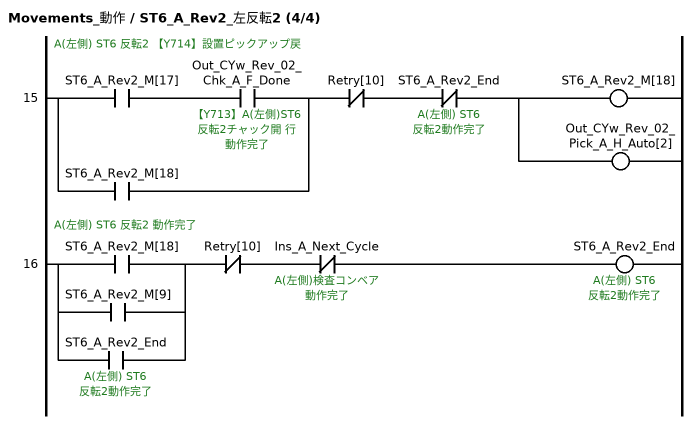
(* [picture p48: Movements_動作 / ST6_A_Rev2_左反転2, rungs 15-16] *)
(* Rung 15: A(左側) ST6 反転2 【Y714】設置ピックアップ戻 *)
_p89 := ((ST6_A_Rev2_M[17] AND Out_CYw_Rev_02_Chk_A_F_Done) OR ST6_A_Rev2_M[18]) AND NOT Retry[10] AND NOT ST6_A_Rev2_End;
ST6_A_Rev2_M[18] := _p89;
Out_CYw_Rev_02_Pick_A_H_Auto[2] := _p89;
(* Rung 16: A(左側) ST6 反転2 動作完了 *)
ST6_A_Rev2_End := (ST6_A_Rev2_M[18] OR ST6_A_Rev2_M[9] OR ST6_A_Rev2_End) AND NOT Retry[10] AND NOT Ins_A_Next_Cycle;

(* Section ST7_A_Dis2_左SF排出: ladder, written here as Structured Text *)

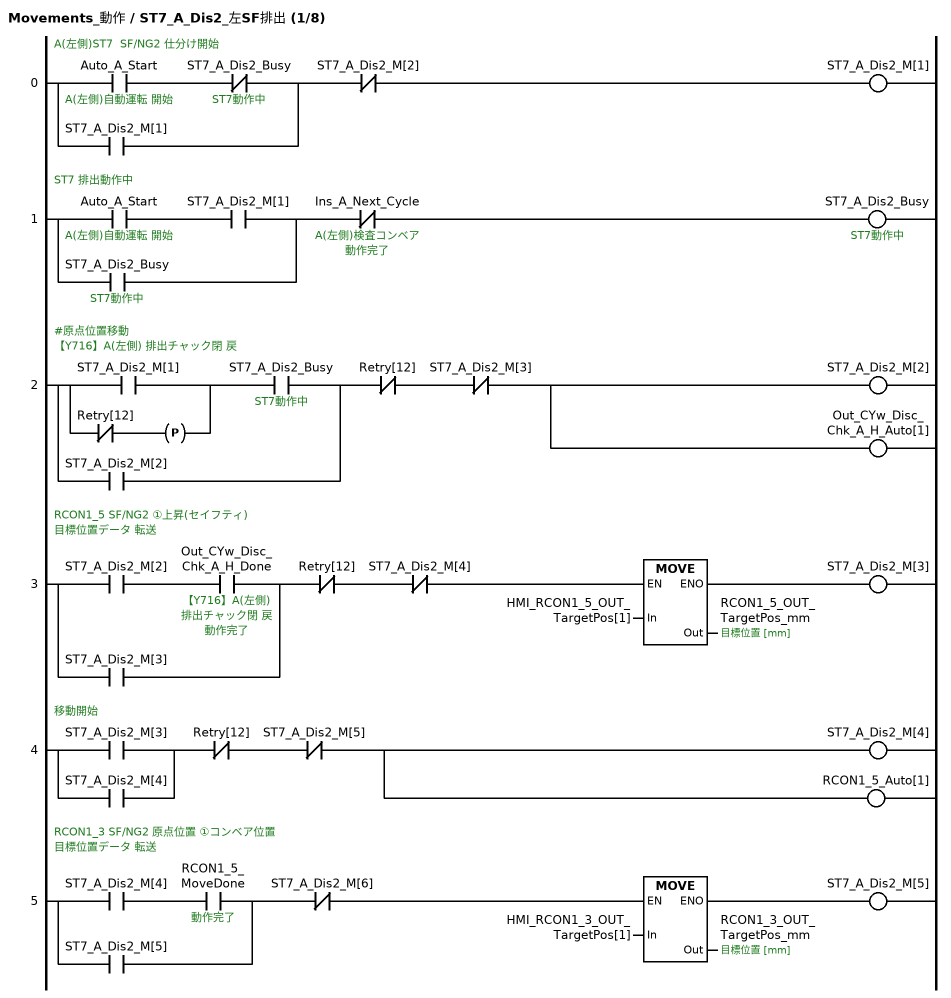
(* Rung 0: A(左側)ST7  SF/NG2 仕分け開始 *)
ST7_A_Dis2_M[1] := ((Auto_A_Start AND NOT ST7_A_Dis2_Busy) OR ST7_A_Dis2_M[1]) AND NOT ST7_A_Dis2_M[2];
(* Rung 1: ST7 排出動作中 *)
ST7_A_Dis2_Busy := ((Auto_A_Start AND ST7_A_Dis2_M[1]) OR ST7_A_Dis2_Busy) AND NOT Ins_A_Next_Cycle;
(* Rung 2: #原点位置移動 / 【Y716】A(左側) 排出チャック閉 戻 *)
_e90(CLK := NOT Retry[12]);
_p91 := (((ST7_A_Dis2_M[1] OR _e90.Q) AND ST7_A_Dis2_Busy) OR ST7_A_Dis2_M[2]) AND NOT Retry[12] AND NOT ST7_A_Dis2_M[3];
ST7_A_Dis2_M[2] := _p91;
Out_CYw_Disc_Chk_A_H_Auto[1] := _p91;
(* Rung 3: RCON1_5 SF/NG2 ①上昇(セイフティ) / 目標位置データ 転送 *)
IF ((ST7_A_Dis2_M[2] AND Out_CYw_Disc_Chk_A_H_Done) OR ST7_A_Dis2_M[3]) AND NOT Retry[12] AND NOT ST7_A_Dis2_M[4] THEN
    RCON1_5_OUT_TargetPos_mm := HMI_RCON1_5_OUT_TargetPos[1];
END_IF;
ST7_A_Dis2_M[3] := ((ST7_A_Dis2_M[2] AND Out_CYw_Disc_Chk_A_H_Done) OR ST7_A_Dis2_M[3]) AND NOT Retry[12] AND NOT ST7_A_Dis2_M[4];
(* Rung 4: 移動開始 *)
_p92 := (ST7_A_Dis2_M[3] OR ST7_A_Dis2_M[4]) AND NOT Retry[12] AND NOT ST7_A_Dis2_M[5];
ST7_A_Dis2_M[4] := _p92;
RCON1_5_Auto[1] := _p92;
(* Rung 5: RCON1_3 SF/NG2 原点位置 ①コンベア位置 / 目標位置データ 転送 *)
IF ((ST7_A_Dis2_M[4] AND RCON1_5_MoveDone) OR ST7_A_Dis2_M[5]) AND NOT ST7_A_Dis2_M[6] THEN
    RCON1_3_OUT_TargetPos_mm := HMI_RCON1_3_OUT_TargetPos[1];
END_IF;
ST7_A_Dis2_M[5] := ((ST7_A_Dis2_M[4] AND RCON1_5_MoveDone) OR ST7_A_Dis2_M[5]) AND NOT ST7_A_Dis2_M[6];

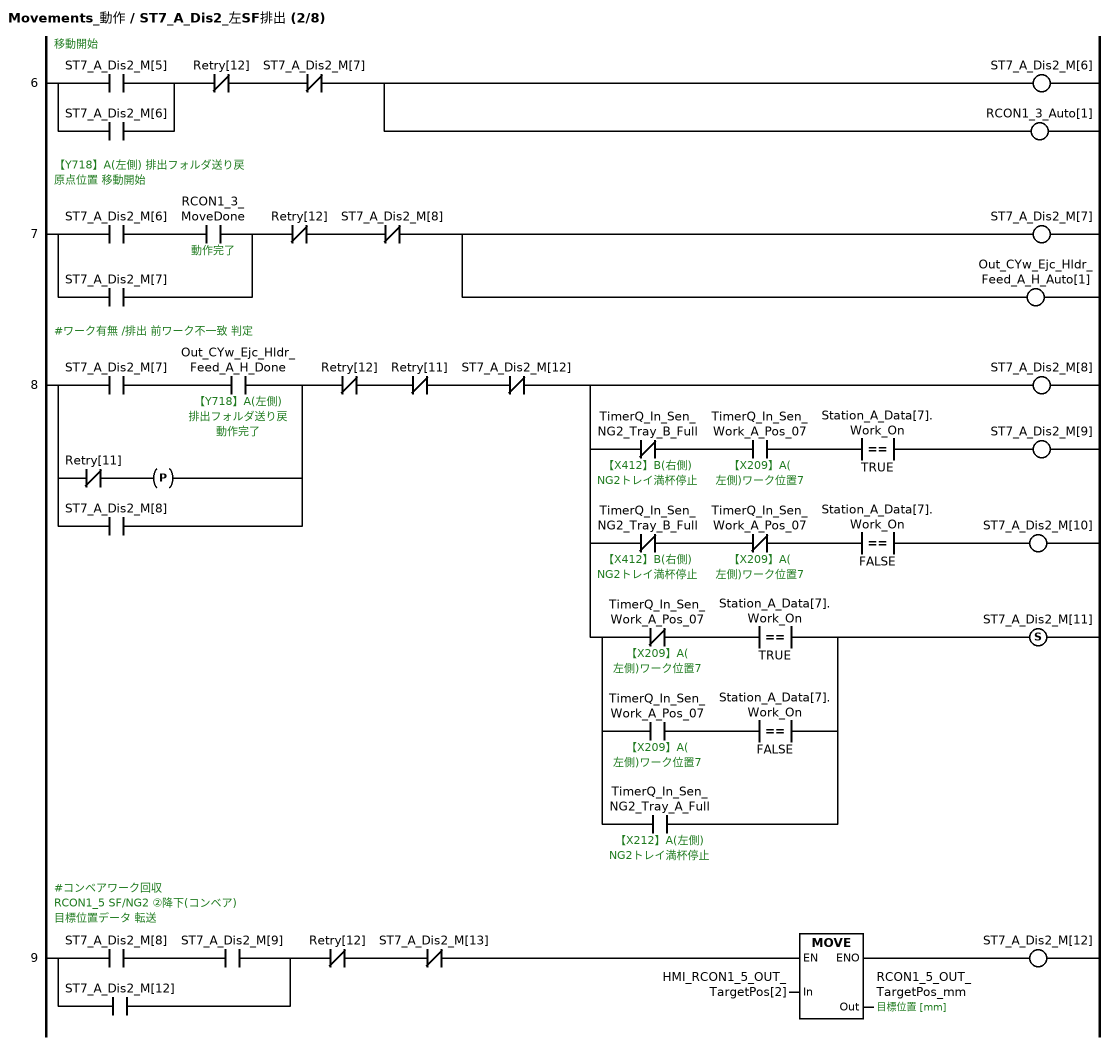
(* Rung 6: 移動開始 *)
_p93 := (ST7_A_Dis2_M[5] OR ST7_A_Dis2_M[6]) AND NOT Retry[12] AND NOT ST7_A_Dis2_M[7];
ST7_A_Dis2_M[6] := _p93;
RCON1_3_Auto[1] := _p93;
(* Rung 7: 【Y718】A(左側) 排出フォルダ送り戻 / 原点位置 移動開始 *)
_p94 := ((ST7_A_Dis2_M[6] AND RCON1_3_MoveDone) OR ST7_A_Dis2_M[7]) AND NOT Retry[12] AND NOT ST7_A_Dis2_M[8];
ST7_A_Dis2_M[7] := _p94;
Out_CYw_Ejc_Hldr_Feed_A_H_Auto[1] := _p94;
(* Rung 8: #ワーク有無 /排出 前ワーク不一致 判定 *)
_e95(CLK := NOT Retry[11]);
_p96 := ((ST7_A_Dis2_M[7] AND Out_CYw_Ejc_Hldr_Feed_A_H_Done) OR _e95.Q OR ST7_A_Dis2_M[8]) AND NOT Retry[12] AND NOT Retry[11] AND NOT ST7_A_Dis2_M[12];
ST7_A_Dis2_M[8] := _p96;
ST7_A_Dis2_M[9] := _p96 AND NOT TimerQ_In_Sen_NG2_Tray_B_Full AND TimerQ_In_Sen_Work_A_Pos_07 AND (Station_A_Data[7].Work_On = TRUE);
ST7_A_Dis2_M[10] := _p96 AND NOT TimerQ_In_Sen_NG2_Tray_B_Full AND NOT TimerQ_In_Sen_Work_A_Pos_07 AND (Station_A_Data[7].Work_On = FALSE);
IF _p96 AND ((NOT TimerQ_In_Sen_Work_A_Pos_07 AND (Station_A_Data[7].Work_On = TRUE)) OR (TimerQ_In_Sen_Work_A_Pos_07 AND (Station_A_Data[7].Work_On = FALSE)) OR TimerQ_In_Sen_NG2_Tray_A_Full) THEN
    ST7_A_Dis2_M[11] := TRUE;
END_IF;
(* Rung 9: #コンベアワーク回収 / RCON1_5 SF/NG2 ②降下(コンベア) / 目標位置データ 転送 *)
IF ((ST7_A_Dis2_M[8] AND ST7_A_Dis2_M[9]) OR ST7_A_Dis2_M[12]) AND NOT Retry[12] AND NOT ST7_A_Dis2_M[13] THEN
    RCON1_5_OUT_TargetPos_mm := HMI_RCON1_5_OUT_TargetPos[2];
END_IF;
ST7_A_Dis2_M[12] := ((ST7_A_Dis2_M[8] AND ST7_A_Dis2_M[9]) OR ST7_A_Dis2_M[12]) AND NOT Retry[12] AND NOT ST7_A_Dis2_M[13];

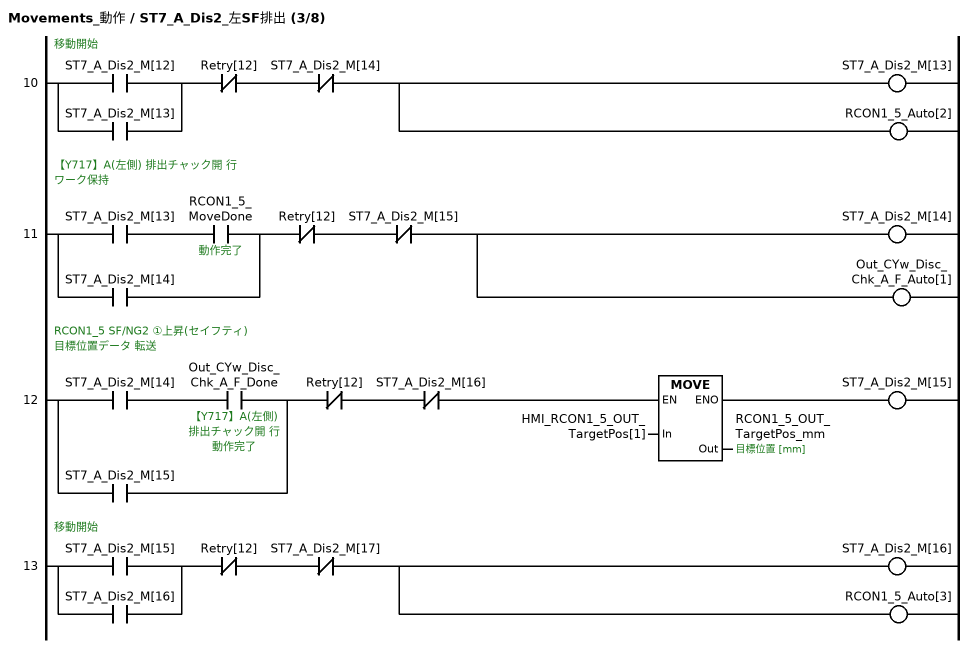
(* Rung 10: 移動開始 *)
_p97 := (ST7_A_Dis2_M[12] OR ST7_A_Dis2_M[13]) AND NOT Retry[12] AND NOT ST7_A_Dis2_M[14];
ST7_A_Dis2_M[13] := _p97;
RCON1_5_Auto[2] := _p97;
(* Rung 11: 【Y717】A(左側) 排出チャック開 行 / ワーク保持 *)
_p98 := ((ST7_A_Dis2_M[13] AND RCON1_5_MoveDone) OR ST7_A_Dis2_M[14]) AND NOT Retry[12] AND NOT ST7_A_Dis2_M[15];
ST7_A_Dis2_M[14] := _p98;
Out_CYw_Disc_Chk_A_F_Auto[1] := _p98;
(* Rung 12: RCON1_5 SF/NG2 ①上昇(セイフティ) / 目標位置データ 転送 *)
IF ((ST7_A_Dis2_M[14] AND Out_CYw_Disc_Chk_A_F_Done) OR ST7_A_Dis2_M[15]) AND NOT Retry[12] AND NOT ST7_A_Dis2_M[16] THEN
    RCON1_5_OUT_TargetPos_mm := HMI_RCON1_5_OUT_TargetPos[1];
END_IF;
ST7_A_Dis2_M[15] := ((ST7_A_Dis2_M[14] AND Out_CYw_Disc_Chk_A_F_Done) OR ST7_A_Dis2_M[15]) AND NOT Retry[12] AND NOT ST7_A_Dis2_M[16];
(* Rung 13: 移動開始 *)
_p99 := (ST7_A_Dis2_M[15] OR ST7_A_Dis2_M[16]) AND NOT Retry[12] AND NOT ST7_A_Dis2_M[17];
ST7_A_Dis2_M[16] := _p99;
RCON1_5_Auto[3] := _p99;

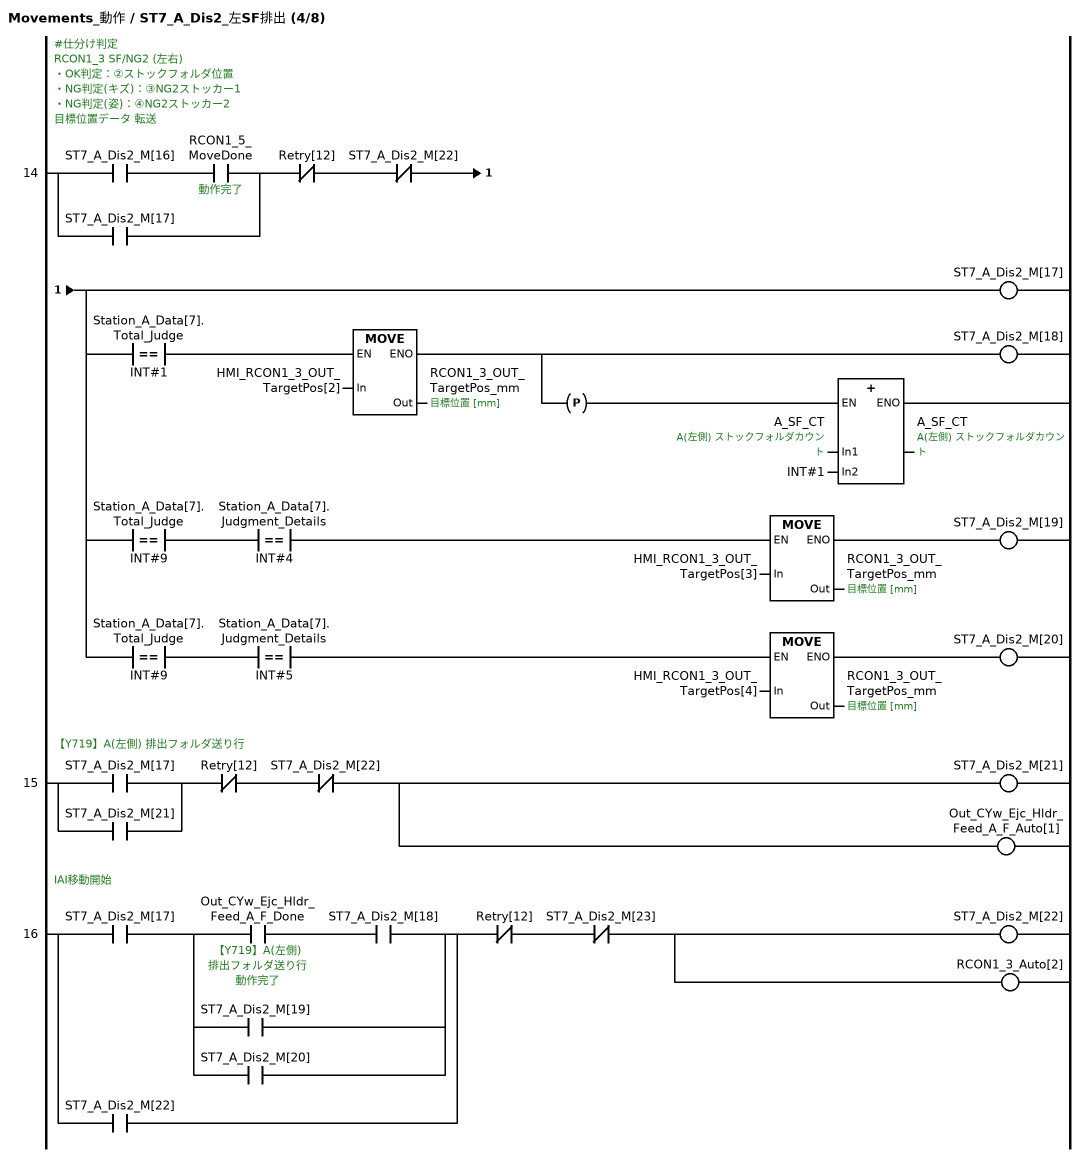
(* Rung 14: #仕分け判定 / RCON1_3 SF/NG2 (左右) / ・OK判定：②ストックフォルダ位置 / ・NG判定(キズ)：③NG2ストッカー1 / ・NG判定(姿)：④NG2ストッカー2 / 目標位置データ 転送 *)
_p100 := ((ST7_A_Dis2_M[16] AND RCON1_5_MoveDone) OR ST7_A_Dis2_M[17]) AND NOT Retry[12] AND NOT ST7_A_Dis2_M[22];
ST7_A_Dis2_M[17] := _p100;
IF _p100 AND (Station_A_Data[7].Total_Judge = INT#1) THEN
    RCON1_3_OUT_TargetPos_mm := HMI_RCON1_3_OUT_TargetPos[2];
END_IF;
_p101 := _p100 AND (Station_A_Data[7].Total_Judge = INT#1);
ST7_A_Dis2_M[18] := _p101;
_e102(CLK := _p101);
IF _e102.Q THEN A_SF_CT := A_SF_CT + INT#1; END_IF;
IF _p100 AND (Station_A_Data[7].Total_Judge = INT#9) AND (Station_A_Data[7].Judgment_Details = INT#4) THEN
    RCON1_3_OUT_TargetPos_mm := HMI_RCON1_3_OUT_TargetPos[3];
END_IF;
ST7_A_Dis2_M[19] := _p100 AND (Station_A_Data[7].Total_Judge = INT#9) AND (Station_A_Data[7].Judgment_Details = INT#4);
IF _p100 AND (Station_A_Data[7].Total_Judge = INT#9) AND (Station_A_Data[7].Judgment_Details = INT#5) THEN
    RCON1_3_OUT_TargetPos_mm := HMI_RCON1_3_OUT_TargetPos[4];
END_IF;
ST7_A_Dis2_M[20] := _p100 AND (Station_A_Data[7].Total_Judge = INT#9) AND (Station_A_Data[7].Judgment_Details = INT#5);
(* Rung 15: 【Y719】A(左側) 排出フォルダ送り行 *)
_p103 := (ST7_A_Dis2_M[17] OR ST7_A_Dis2_M[21]) AND NOT Retry[12] AND NOT ST7_A_Dis2_M[22];
ST7_A_Dis2_M[21] := _p103;
Out_CYw_Ejc_Hldr_Feed_A_F_Auto[1] := _p103;
(* Rung 16: IAI移動開始 *)
_p104 := ((ST7_A_Dis2_M[17] AND ((Out_CYw_Ejc_Hldr_Feed_A_F_Done AND ST7_A_Dis2_M[18]) OR ST7_A_Dis2_M[19] OR ST7_A_Dis2_M[20])) OR ST7_A_Dis2_M[22]) AND NOT Retry[12] AND NOT ST7_A_Dis2_M[23];
ST7_A_Dis2_M[22] := _p104;
RCON1_3_Auto[2] := _p104;

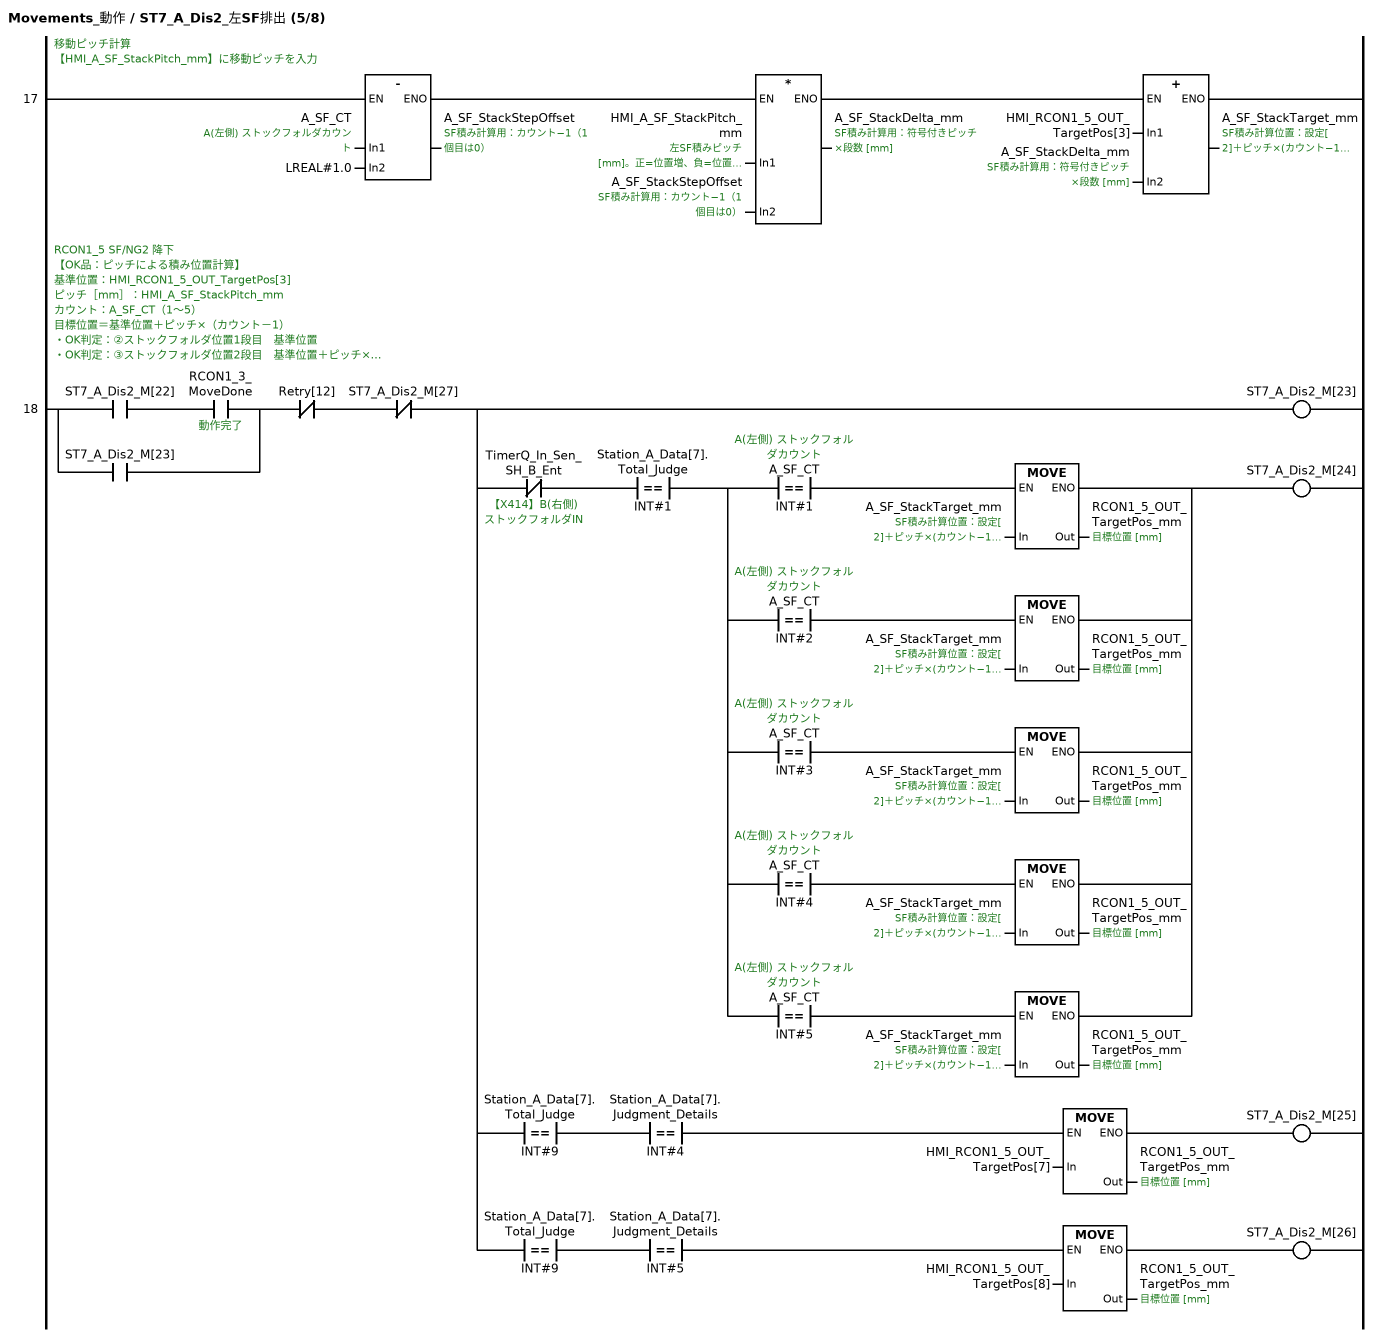
(* Rung 17: 移動ピッチ計算 / 【HMI_A_SF_StackPitch_mm】に移動ピッチを入力 *)
A_SF_StackStepOffset := A_SF_CT - LREAL#1.0;
A_SF_StackDelta_mm := HMI_A_SF_StackPitch_mm * A_SF_StackStepOffset;
A_SF_StackTarget_mm := HMI_RCON1_5_OUT_TargetPos[3] + A_SF_StackDelta_mm;
(* Rung 18: RCON1_5 SF/NG2 降下 / 【OK品：ピッチによる積み位置計算】 / 基準位置：HMI_RCON1_5_OUT_TargetPos[3] / ピッチ［mm］：HMI_A_SF_StackPitch_mm / カウント：A_SF_CT（1～5） / 目標位置＝基準位置＋ピッチ×（カウント－1） / ・OK判定：②ストックフォルダ位置1段目　基準位置 / ・OK判定：③ストックフォルダ位置2段目　基準位置＋ピッチ×1 / ・OK判定：④ストックフォルダ位置3段目　基準位置＋ピッチ×2 / ・OK判定：⑤ストックフォルダ位置4段目　基準位置＋ピッチ×3 / ・OK判定：⑥ストックフォルダ位置5段目　基準位置＋ピッチ×4 / 【NG品：従来の固定位置を使用】 / ・NG判定(キズ)：⑦NG2ストッカー1 / ・NG判定(姿)：⑧NG2ストッカー2 / 目標位置データ 転送 *)
_p105 := ((ST7_A_Dis2_M[22] AND RCON1_3_MoveDone) OR ST7_A_Dis2_M[23]) AND NOT Retry[12] AND NOT ST7_A_Dis2_M[27];
ST7_A_Dis2_M[23] := _p105;
_p106 := _p105 AND NOT TimerQ_In_Sen_SH_B_Ent AND (Station_A_Data[7].Total_Judge = INT#1);
IF _p106 AND (A_SF_CT = INT#1) THEN RCON1_5_OUT_TargetPos_mm := A_SF_StackTarget_mm; END_IF;
IF _p106 AND (A_SF_CT = INT#2) THEN RCON1_5_OUT_TargetPos_mm := A_SF_StackTarget_mm; END_IF;
IF _p106 AND (A_SF_CT = INT#3) THEN RCON1_5_OUT_TargetPos_mm := A_SF_StackTarget_mm; END_IF;
IF _p106 AND (A_SF_CT = INT#4) THEN RCON1_5_OUT_TargetPos_mm := A_SF_StackTarget_mm; END_IF;
IF _p106 AND (A_SF_CT = INT#5) THEN RCON1_5_OUT_TargetPos_mm := A_SF_StackTarget_mm; END_IF;
ST7_A_Dis2_M[24] := _p106 AND ((A_SF_CT = INT#1) OR (A_SF_CT = INT#2) OR (A_SF_CT = INT#3) OR (A_SF_CT = INT#4) OR (A_SF_CT = INT#5));
IF _p105 AND (Station_A_Data[7].Total_Judge = INT#9) AND (Station_A_Data[7].Judgment_Details = INT#4) THEN
    RCON1_5_OUT_TargetPos_mm := HMI_RCON1_5_OUT_TargetPos[7];
END_IF;
ST7_A_Dis2_M[25] := _p105 AND (Station_A_Data[7].Total_Judge = INT#9) AND (Station_A_Data[7].Judgment_Details = INT#4);
IF _p105 AND (Station_A_Data[7].Total_Judge = INT#9) AND (Station_A_Data[7].Judgment_Details = INT#5) THEN
    RCON1_5_OUT_TargetPos_mm := HMI_RCON1_5_OUT_TargetPos[8];
END_IF;
ST7_A_Dis2_M[26] := _p105 AND (Station_A_Data[7].Total_Judge = INT#9) AND (Station_A_Data[7].Judgment_Details = INT#5);

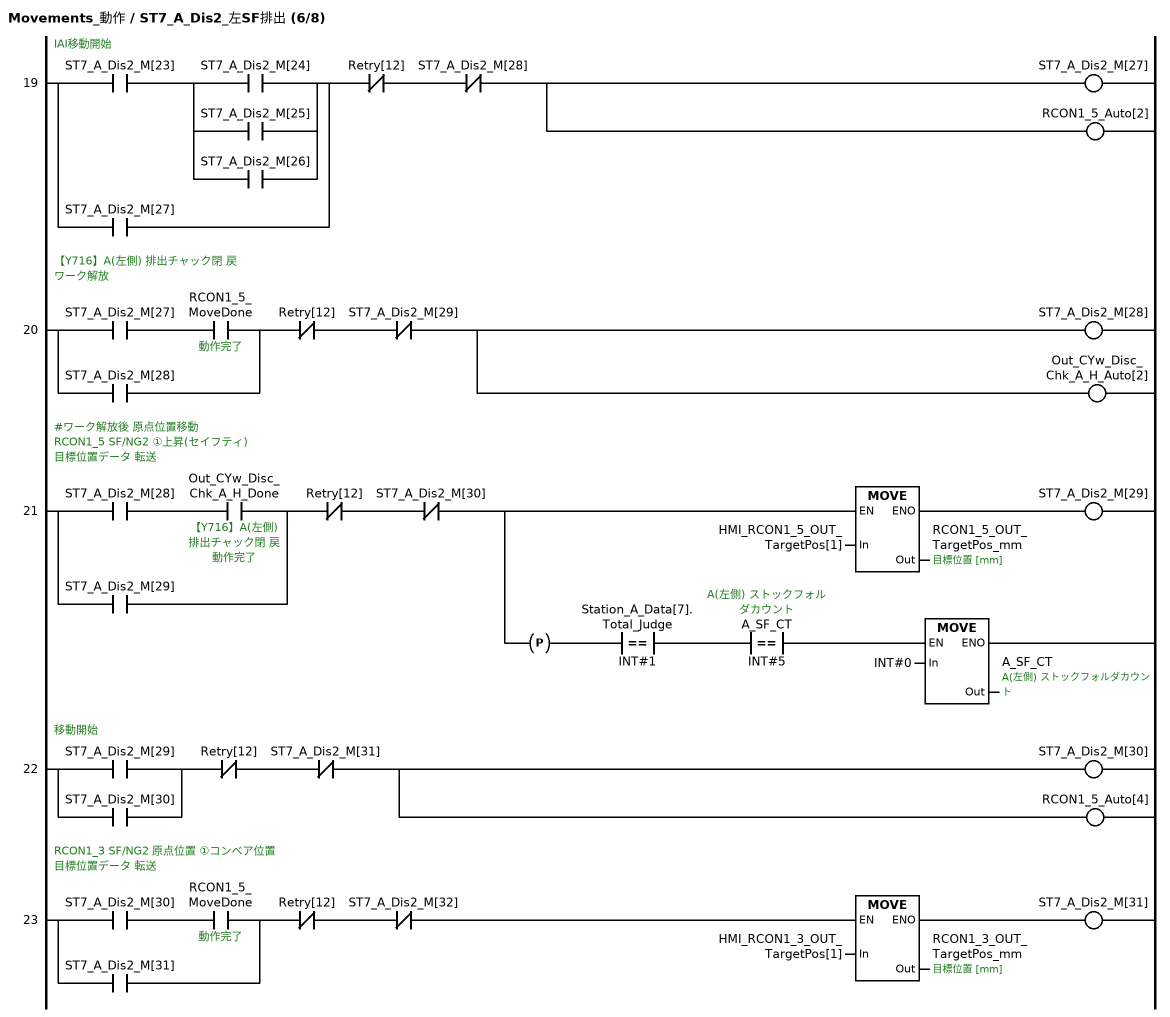
(* Rung 19: IAI移動開始 *)
_p107 := ((ST7_A_Dis2_M[23] AND (ST7_A_Dis2_M[24] OR ST7_A_Dis2_M[25] OR ST7_A_Dis2_M[26])) OR ST7_A_Dis2_M[27]) AND NOT Retry[12] AND NOT ST7_A_Dis2_M[28];
ST7_A_Dis2_M[27] := _p107;
RCON1_5_Auto[2] := _p107;
(* Rung 20: 【Y716】A(左側) 排出チャック閉 戻 / ワーク解放 *)
_p108 := ((ST7_A_Dis2_M[27] AND RCON1_5_MoveDone) OR ST7_A_Dis2_M[28]) AND NOT Retry[12] AND NOT ST7_A_Dis2_M[29];
ST7_A_Dis2_M[28] := _p108;
Out_CYw_Disc_Chk_A_H_Auto[2] := _p108;
(* Rung 21: #ワーク解放後 原点位置移動 / RCON1_5 SF/NG2 ①上昇(セイフティ) / 目標位置データ 転送 *)
_p109 := ((ST7_A_Dis2_M[28] AND Out_CYw_Disc_Chk_A_H_Done) OR ST7_A_Dis2_M[29]) AND NOT Retry[12] AND NOT ST7_A_Dis2_M[30];
IF _p109 THEN RCON1_5_OUT_TargetPos_mm := HMI_RCON1_5_OUT_TargetPos[1]; END_IF;
ST7_A_Dis2_M[29] := _p109;
_e110(CLK := _p109);
IF _e110.Q AND (Station_A_Data[7].Total_Judge = INT#1) AND (A_SF_CT = INT#5) THEN
    A_SF_CT := INT#0;
END_IF;
(* Rung 22: 移動開始 *)
_p111 := (ST7_A_Dis2_M[29] OR ST7_A_Dis2_M[30]) AND NOT Retry[12] AND NOT ST7_A_Dis2_M[31];
ST7_A_Dis2_M[30] := _p111;
RCON1_5_Auto[4] := _p111;
(* Rung 23: RCON1_3 SF/NG2 原点位置 ①コンベア位置 / 目標位置データ 転送 *)
IF ((ST7_A_Dis2_M[30] AND RCON1_5_MoveDone) OR ST7_A_Dis2_M[31]) AND NOT Retry[12] AND NOT ST7_A_Dis2_M[32] THEN
    RCON1_3_OUT_TargetPos_mm := HMI_RCON1_3_OUT_TargetPos[1];
END_IF;
ST7_A_Dis2_M[31] := ((ST7_A_Dis2_M[30] AND RCON1_5_MoveDone) OR ST7_A_Dis2_M[31]) AND NOT Retry[12] AND NOT ST7_A_Dis2_M[32];

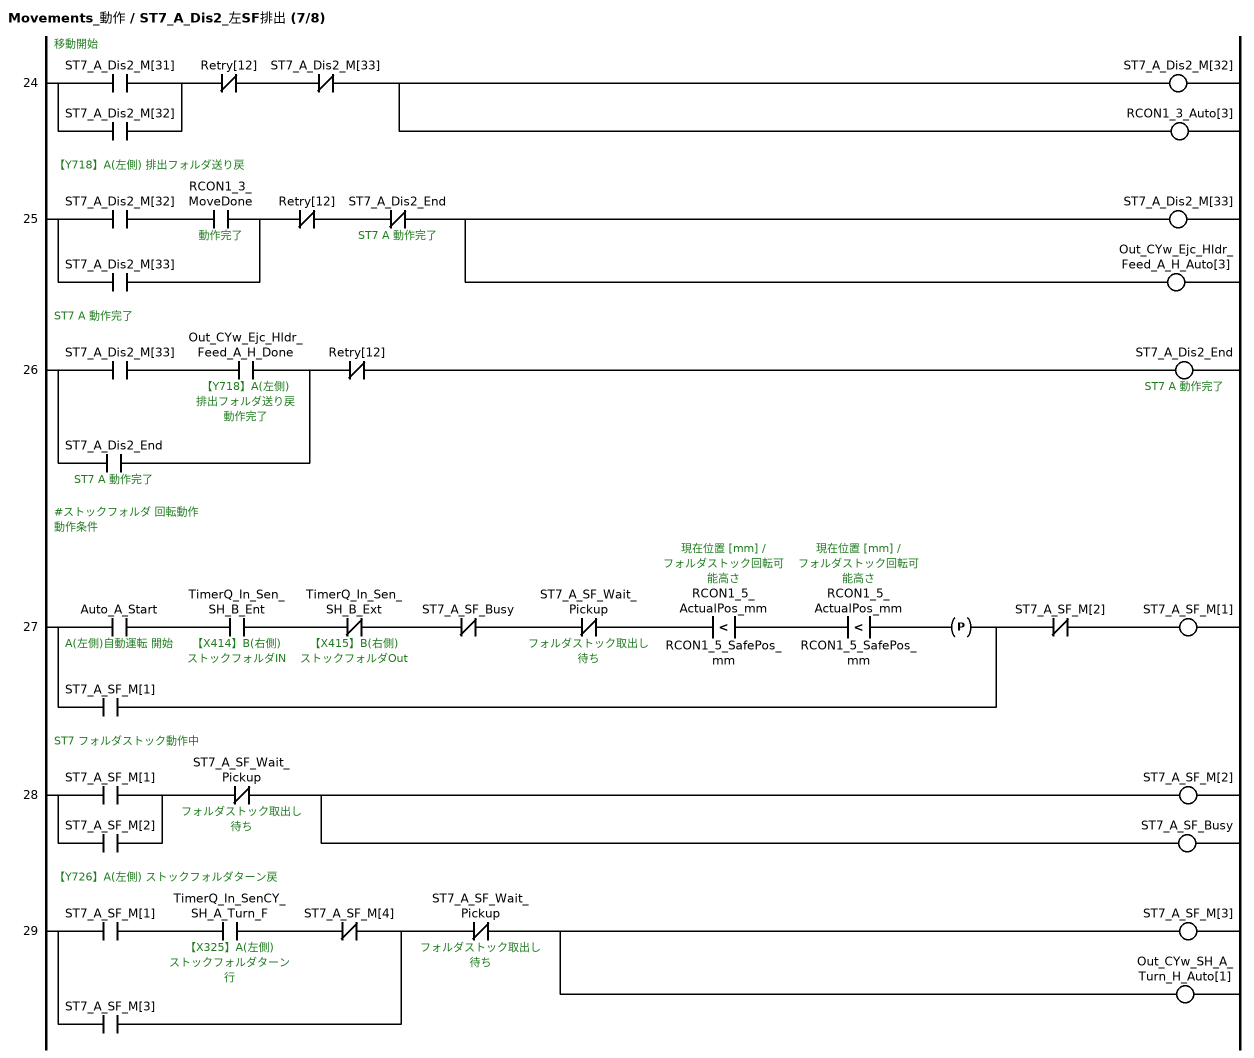
(* Rung 24: 移動開始 *)
_p112 := (ST7_A_Dis2_M[31] OR ST7_A_Dis2_M[32]) AND NOT Retry[12] AND NOT ST7_A_Dis2_M[33];
ST7_A_Dis2_M[32] := _p112;
RCON1_3_Auto[3] := _p112;
(* Rung 25: 【Y718】A(左側) 排出フォルダ送り戻 *)
_p113 := ((ST7_A_Dis2_M[32] AND RCON1_3_MoveDone) OR ST7_A_Dis2_M[33]) AND NOT Retry[12] AND NOT ST7_A_Dis2_End;
ST7_A_Dis2_M[33] := _p113;
Out_CYw_Ejc_Hldr_Feed_A_H_Auto[3] := _p113;
(* Rung 26: ST7 A 動作完了 *)
ST7_A_Dis2_End := ((ST7_A_Dis2_M[33] AND Out_CYw_Ejc_Hldr_Feed_A_H_Done) OR ST7_A_Dis2_End) AND NOT Retry[12];
(* Rung 27: #ストックフォルダ 回転動作 / 動作条件 *)
_e114(CLK := Auto_A_Start AND TimerQ_In_Sen_SH_B_Ent AND NOT TimerQ_In_Sen_SH_B_Ext AND NOT ST7_A_SF_Busy AND NOT ST7_A_SF_Wait_Pickup AND (RCON1_5_ActualPos_mm < RCON1_5_SafePos_mm) AND (RCON1_5_ActualPos_mm < RCON1_5_SafePos_mm));
ST7_A_SF_M[1] := (_e114.Q OR ST7_A_SF_M[1]) AND NOT ST7_A_SF_M[2];
(* Rung 28: ST7 フォルダストック動作中 *)
_p115 := (ST7_A_SF_M[1] OR ST7_A_SF_M[2]) AND NOT ST7_A_SF_Wait_Pickup;
ST7_A_SF_M[2] := _p115;
ST7_A_SF_Busy := _p115;
(* Rung 29: 【Y726】A(左側) ストックフォルダターン戻 *)
_p116 := ((ST7_A_SF_M[1] AND TimerQ_In_SenCY_SH_A_Turn_F AND NOT ST7_A_SF_M[4]) OR ST7_A_SF_M[3]) AND NOT ST7_A_SF_Wait_Pickup;
ST7_A_SF_M[3] := _p116;
Out_CYw_SH_A_Turn_H_Auto[1] := _p116;

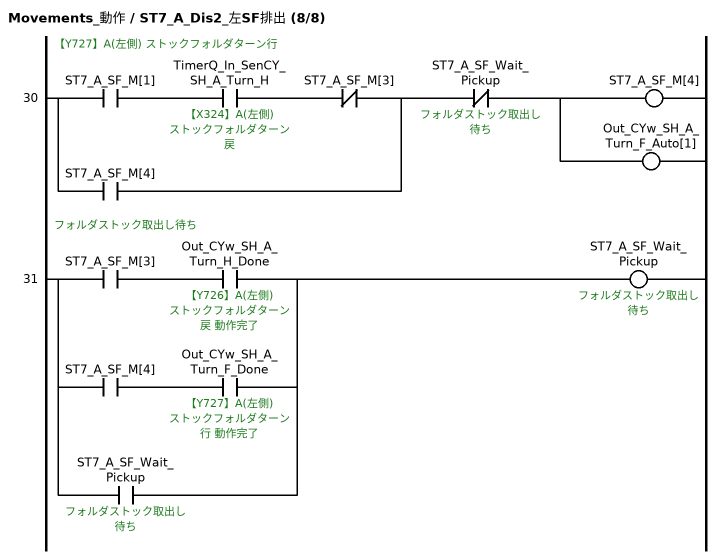
(* Rung 30: 【Y727】A(左側) ストックフォルダターン行 *)
_p117 := ((ST7_A_SF_M[1] AND TimerQ_In_SenCY_SH_A_Turn_H AND NOT ST7_A_SF_M[3]) OR ST7_A_SF_M[4]) AND NOT ST7_A_SF_Wait_Pickup;
ST7_A_SF_M[4] := _p117;
Out_CYw_SH_A_Turn_F_Auto[1] := _p117;
(* Rung 31: フォルダストック取出し待ち *)
ST7_A_SF_Wait_Pickup := (ST7_A_SF_M[3] AND Out_CYw_SH_A_Turn_H_Done) OR (ST7_A_SF_M[4] AND Out_CYw_SH_A_Turn_F_Done) OR ST7_A_SF_Wait_Pickup;

(* Section Destacker_段バラシ: ladder, written here as Structured Text *)

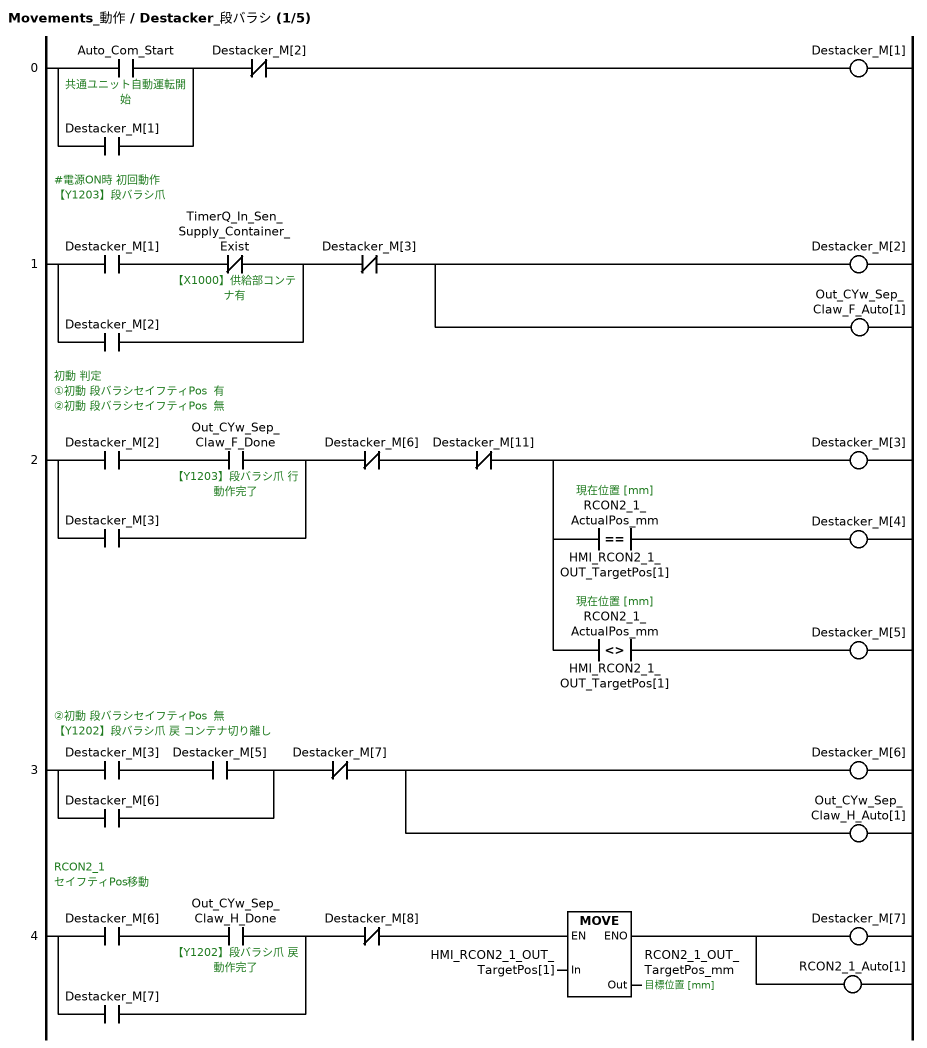
(* Rung 0 *)
Destacker_M[1] := (Auto_Com_Start OR Destacker_M[1]) AND NOT Destacker_M[2];
(* Rung 1: #電源ON時 初回動作 / 【Y1203】段バラシ爪 *)
_p118 := ((Destacker_M[1] AND NOT TimerQ_In_Sen_Supply_Container_Exist) OR Destacker_M[2]) AND NOT Destacker_M[3];
Destacker_M[2] := _p118;
Out_CYw_Sep_Claw_F_Auto[1] := _p118;
(* Rung 2: 初動 判定 / ①初動 段バラシセイフティPos  有 / ②初動 段バラシセイフティPos  無 *)
_p119 := ((Destacker_M[2] AND Out_CYw_Sep_Claw_F_Done) OR Destacker_M[3]) AND NOT Destacker_M[6] AND NOT Destacker_M[11];
Destacker_M[3] := _p119;
Destacker_M[4] := _p119 AND (RCON2_1_ActualPos_mm = HMI_RCON2_1_OUT_TargetPos[1]);
Destacker_M[5] := _p119 AND (RCON2_1_ActualPos_mm <> HMI_RCON2_1_OUT_TargetPos[1]);
(* Rung 3: ②初動 段バラシセイフティPos  無 / 【Y1202】段バラシ爪 戻 コンテナ切り離し *)
_p120 := ((Destacker_M[3] AND Destacker_M[5]) OR Destacker_M[6]) AND NOT Destacker_M[7];
Destacker_M[6] := _p120;
Out_CYw_Sep_Claw_H_Auto[1] := _p120;
(* Rung 4: RCON2_1 / セイフティPos移動 *)
IF ((Destacker_M[6] AND Out_CYw_Sep_Claw_H_Done) OR Destacker_M[7]) AND NOT Destacker_M[8] THEN
    RCON2_1_OUT_TargetPos_mm := HMI_RCON2_1_OUT_TargetPos[1];
END_IF;
_p121 := ((Destacker_M[6] AND Out_CYw_Sep_Claw_H_Done) OR Destacker_M[7]) AND NOT Destacker_M[8];
Destacker_M[7] := _p121;
RCON2_1_Auto[1] := _p121;

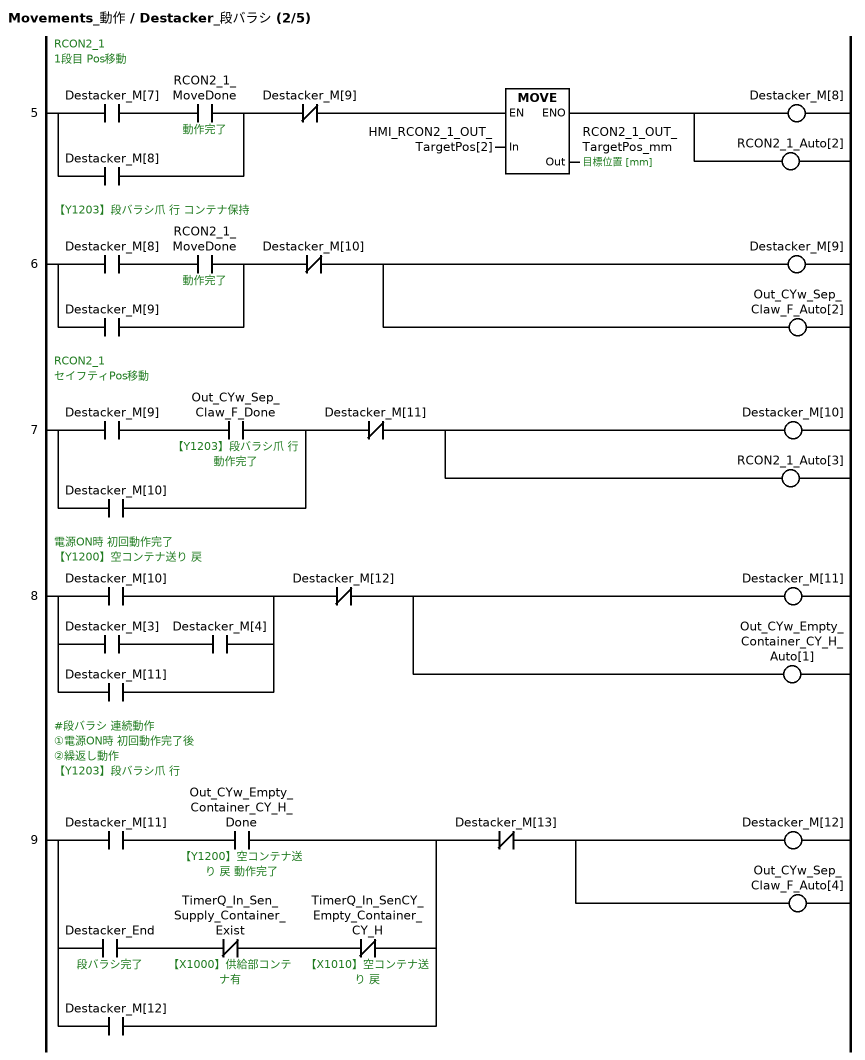
(* Rung 5: RCON2_1 / 1段目 Pos移動 *)
IF ((Destacker_M[7] AND RCON2_1_MoveDone) OR Destacker_M[8]) AND NOT Destacker_M[9] THEN
    RCON2_1_OUT_TargetPos_mm := HMI_RCON2_1_OUT_TargetPos[2];
END_IF;
_p122 := ((Destacker_M[7] AND RCON2_1_MoveDone) OR Destacker_M[8]) AND NOT Destacker_M[9];
Destacker_M[8] := _p122;
RCON2_1_Auto[2] := _p122;
(* Rung 6: 【Y1203】段バラシ爪 行 コンテナ保持 *)
_p123 := ((Destacker_M[8] AND RCON2_1_MoveDone) OR Destacker_M[9]) AND NOT Destacker_M[10];
Destacker_M[9] := _p123;
Out_CYw_Sep_Claw_F_Auto[2] := _p123;
(* Rung 7: RCON2_1 / セイフティPos移動 *)
_p124 := ((Destacker_M[9] AND Out_CYw_Sep_Claw_F_Done) OR Destacker_M[10]) AND NOT Destacker_M[11];
Destacker_M[10] := _p124;
RCON2_1_Auto[3] := _p124;
(* Rung 8: 電源ON時 初回動作完了 / 【Y1200】空コンテナ送り 戻 *)
_p125 := (Destacker_M[10] OR (Destacker_M[3] AND Destacker_M[4]) OR Destacker_M[11]) AND NOT Destacker_M[12];
Destacker_M[11] := _p125;
Out_CYw_Empty_Container_CY_H_Auto[1] := _p125;
(* Rung 9: #段バラシ 連続動作 / ①電源ON時 初回動作完了後 / ②繰返し動作 / 【Y1203】段バラシ爪 行 *)
_p126 := ((Destacker_M[11] AND Out_CYw_Empty_Container_CY_H_Done) OR (Destacker_End AND NOT TimerQ_In_Sen_Supply_Container_Exist AND NOT TimerQ_In_SenCY_Empty_Container_CY_H) OR Destacker_M[12]) AND NOT Destacker_M[13];
Destacker_M[12] := _p126;
Out_CYw_Sep_Claw_F_Auto[4] := _p126;

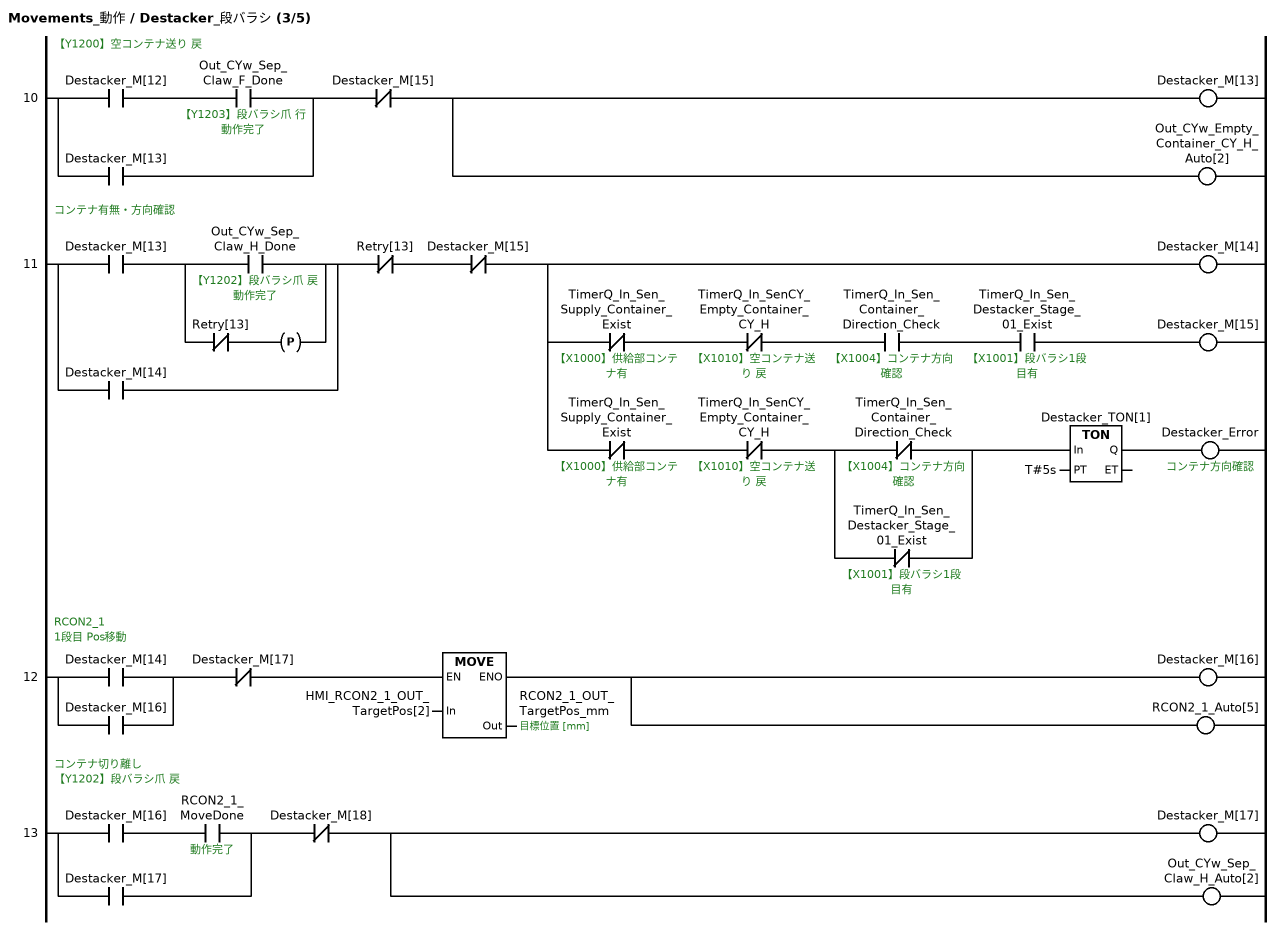
(* Rung 10: 【Y1200】空コンテナ送り 戻 *)
_p127 := ((Destacker_M[12] AND Out_CYw_Sep_Claw_F_Done) OR Destacker_M[13]) AND NOT Destacker_M[15];
Destacker_M[13] := _p127;
Out_CYw_Empty_Container_CY_H_Auto[2] := _p127;
(* Rung 11: コンテナ有無・方向確認 *)
_e128(CLK := Destacker_M[13] AND NOT Retry[13]);
_p129 := ((Destacker_M[13] AND Out_CYw_Sep_Claw_H_Done) OR _e128.Q OR Destacker_M[14]) AND NOT Retry[13] AND NOT Destacker_M[15];
Destacker_M[14] := _p129;
Destacker_M[15] := _p129 AND NOT TimerQ_In_Sen_Supply_Container_Exist AND NOT TimerQ_In_SenCY_Empty_Container_CY_H AND TimerQ_In_Sen_Container_Direction_Check AND TimerQ_In_Sen_Destacker_Stage_01_Exist;
Destacker_TON[1](In := _p129 AND NOT TimerQ_In_Sen_Supply_Container_Exist AND NOT TimerQ_In_SenCY_Empty_Container_CY_H AND (NOT TimerQ_In_Sen_Container_Direction_Check OR NOT TimerQ_In_Sen_Destacker_Stage_01_Exist), PT := T#5s);
Destacker_Error := Destacker_TON[1].Q;
(* Rung 12: RCON2_1 / 1段目 Pos移動 *)
IF (Destacker_M[14] OR Destacker_M[16]) AND NOT Destacker_M[17] THEN
    RCON2_1_OUT_TargetPos_mm := HMI_RCON2_1_OUT_TargetPos[2];
END_IF;
_p130 := (Destacker_M[14] OR Destacker_M[16]) AND NOT Destacker_M[17];
Destacker_M[16] := _p130;
RCON2_1_Auto[5] := _p130;
(* Rung 13: コンテナ切り離し / 【Y1202】段バラシ爪 戻 *)
_p131 := ((Destacker_M[16] AND RCON2_1_MoveDone) OR Destacker_M[17]) AND NOT Destacker_M[18];
Destacker_M[17] := _p131;
Out_CYw_Sep_Claw_H_Auto[2] := _p131;

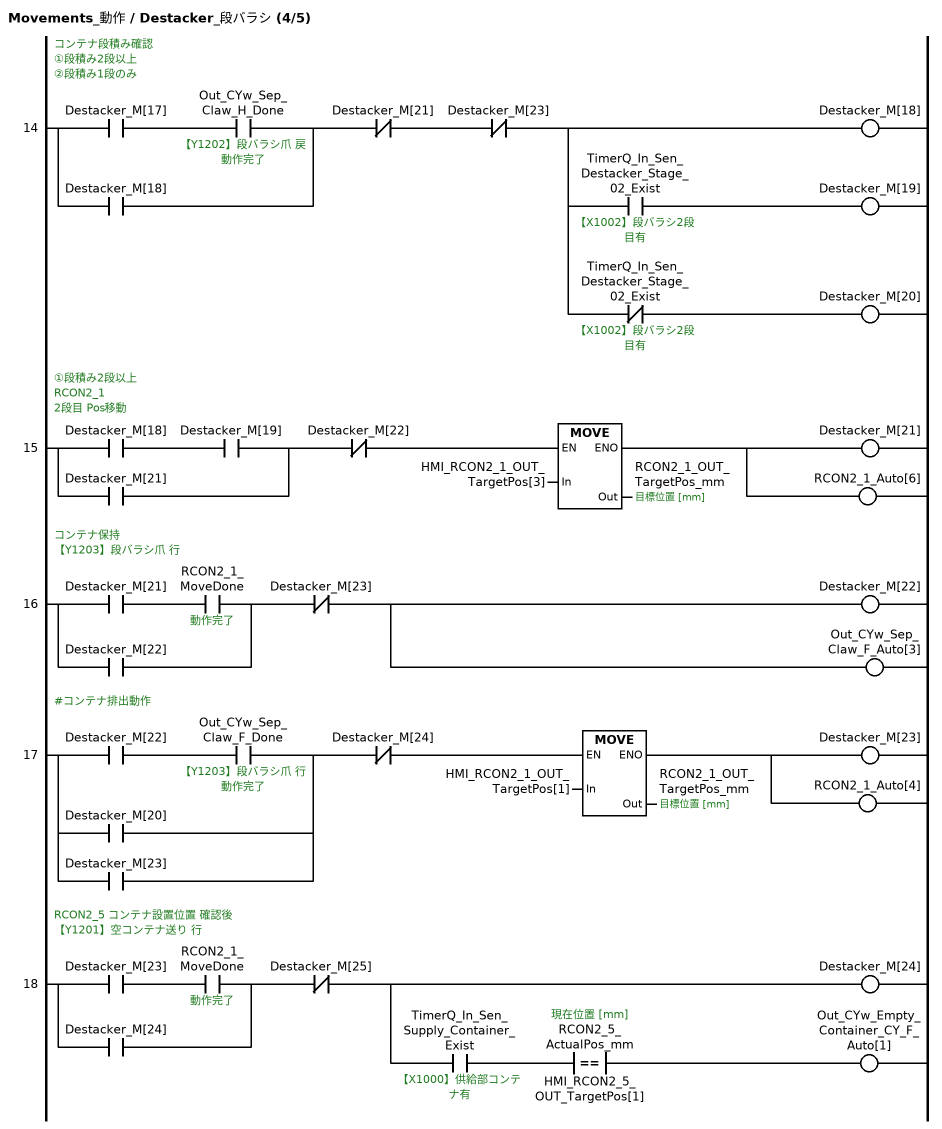
(* Rung 14: コンテナ段積み確認 / ①段積み2段以上 / ②段積み1段のみ *)
_p132 := ((Destacker_M[17] AND Out_CYw_Sep_Claw_H_Done) OR Destacker_M[18]) AND NOT Destacker_M[21] AND NOT Destacker_M[23];
Destacker_M[18] := _p132;
Destacker_M[19] := _p132 AND TimerQ_In_Sen_Destacker_Stage_02_Exist;
Destacker_M[20] := _p132 AND NOT TimerQ_In_Sen_Destacker_Stage_02_Exist;
(* Rung 15: ①段積み2段以上 / RCON2_1 / 2段目 Pos移動 *)
IF ((Destacker_M[18] AND Destacker_M[19]) OR Destacker_M[21]) AND NOT Destacker_M[22] THEN
    RCON2_1_OUT_TargetPos_mm := HMI_RCON2_1_OUT_TargetPos[3];
END_IF;
_p133 := ((Destacker_M[18] AND Destacker_M[19]) OR Destacker_M[21]) AND NOT Destacker_M[22];
Destacker_M[21] := _p133;
RCON2_1_Auto[6] := _p133;
(* Rung 16: コンテナ保持 / 【Y1203】段バラシ爪 行 *)
_p134 := ((Destacker_M[21] AND RCON2_1_MoveDone) OR Destacker_M[22]) AND NOT Destacker_M[23];
Destacker_M[22] := _p134;
Out_CYw_Sep_Claw_F_Auto[3] := _p134;
(* Rung 17: #コンテナ排出動作 *)
IF ((Destacker_M[22] AND Out_CYw_Sep_Claw_F_Done) OR Destacker_M[20] OR Destacker_M[23]) AND NOT Destacker_M[24] THEN
    RCON2_1_OUT_TargetPos_mm := HMI_RCON2_1_OUT_TargetPos[1];
END_IF;
_p135 := ((Destacker_M[22] AND Out_CYw_Sep_Claw_F_Done) OR Destacker_M[20] OR Destacker_M[23]) AND NOT Destacker_M[24];
Destacker_M[23] := _p135;
RCON2_1_Auto[4] := _p135;
(* Rung 18: RCON2_5 コンテナ設置位置 確認後 / 【Y1201】空コンテナ送り 行 *)
_p136 := ((Destacker_M[23] AND RCON2_1_MoveDone) OR Destacker_M[24]) AND NOT Destacker_M[25];
Destacker_M[24] := _p136;
Out_CYw_Empty_Container_CY_F_Auto[1] := _p136 AND TimerQ_In_Sen_Supply_Container_Exist AND (RCON2_5_ActualPos_mm = HMI_RCON2_5_OUT_TargetPos[1]);

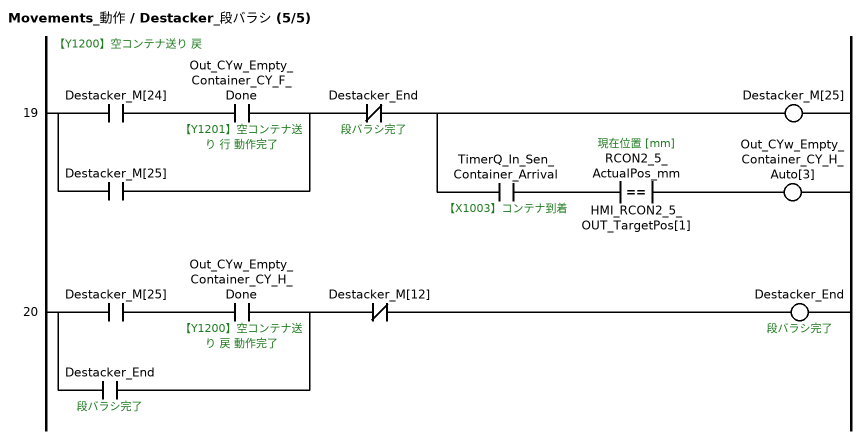
(* Rung 19: 【Y1200】空コンテナ送り 戻 *)
_p137 := ((Destacker_M[24] AND Out_CYw_Empty_Container_CY_F_Done) OR Destacker_M[25]) AND NOT Destacker_End;
Destacker_M[25] := _p137;
Out_CYw_Empty_Container_CY_H_Auto[3] := _p137 AND TimerQ_In_Sen_Container_Arrival AND (RCON2_5_ActualPos_mm = HMI_RCON2_5_OUT_TargetPos[1]);
(* Rung 20 *)
Destacker_End := ((Destacker_M[25] AND Out_CYw_Empty_Container_CY_H_Done) OR Destacker_End) AND NOT Destacker_M[12];

(* Section BoxPacking_箱詰め: ladder, written here as Structured Text *)

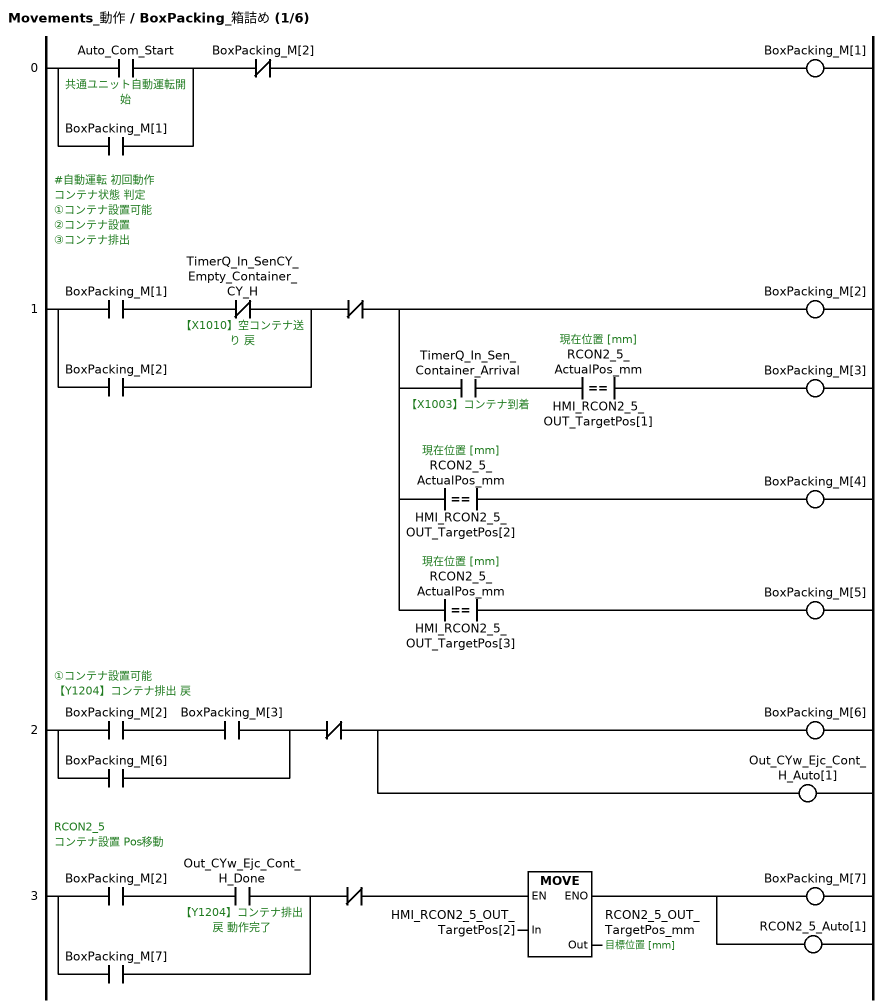
(* Rung 0 *)
BoxPacking_M[1] := (Auto_Com_Start OR BoxPacking_M[1]) AND NOT BoxPacking_M[2];
(* Rung 1: #自動運転 初回動作 / コンテナ状態 判定 / ①コンテナ設置可能 / ②コンテナ設置 / ③コンテナ排出 *)
_p138 := ((BoxPacking_M[1] AND NOT TimerQ_In_SenCY_Empty_Container_CY_H) OR BoxPacking_M[2]) AND NOT ();
BoxPacking_M[2] := _p138;
BoxPacking_M[3] := _p138 AND TimerQ_In_Sen_Container_Arrival AND (RCON2_5_ActualPos_mm = HMI_RCON2_5_OUT_TargetPos[1]);
BoxPacking_M[4] := _p138 AND (RCON2_5_ActualPos_mm = HMI_RCON2_5_OUT_TargetPos[2]);
BoxPacking_M[5] := _p138 AND (RCON2_5_ActualPos_mm = HMI_RCON2_5_OUT_TargetPos[3]);
(* Rung 2: ①コンテナ設置可能 / 【Y1204】コンテナ排出 戻 *)
_p139 := ((BoxPacking_M[2] AND BoxPacking_M[3]) OR BoxPacking_M[6]) AND NOT ();
BoxPacking_M[6] := _p139;
Out_CYw_Ejc_Cont_H_Auto[1] := _p139;
(* Rung 3: RCON2_5 / コンテナ設置 Pos移動 *)
IF ((BoxPacking_M[2] AND Out_CYw_Ejc_Cont_H_Done) OR BoxPacking_M[7]) AND NOT () THEN
    RCON2_5_OUT_TargetPos_mm := HMI_RCON2_5_OUT_TargetPos[2];
END_IF;
_p140 := ((BoxPacking_M[2] AND Out_CYw_Ejc_Cont_H_Done) OR BoxPacking_M[7]) AND NOT ();
BoxPacking_M[7] := _p140;
RCON2_5_Auto[1] := _p140;

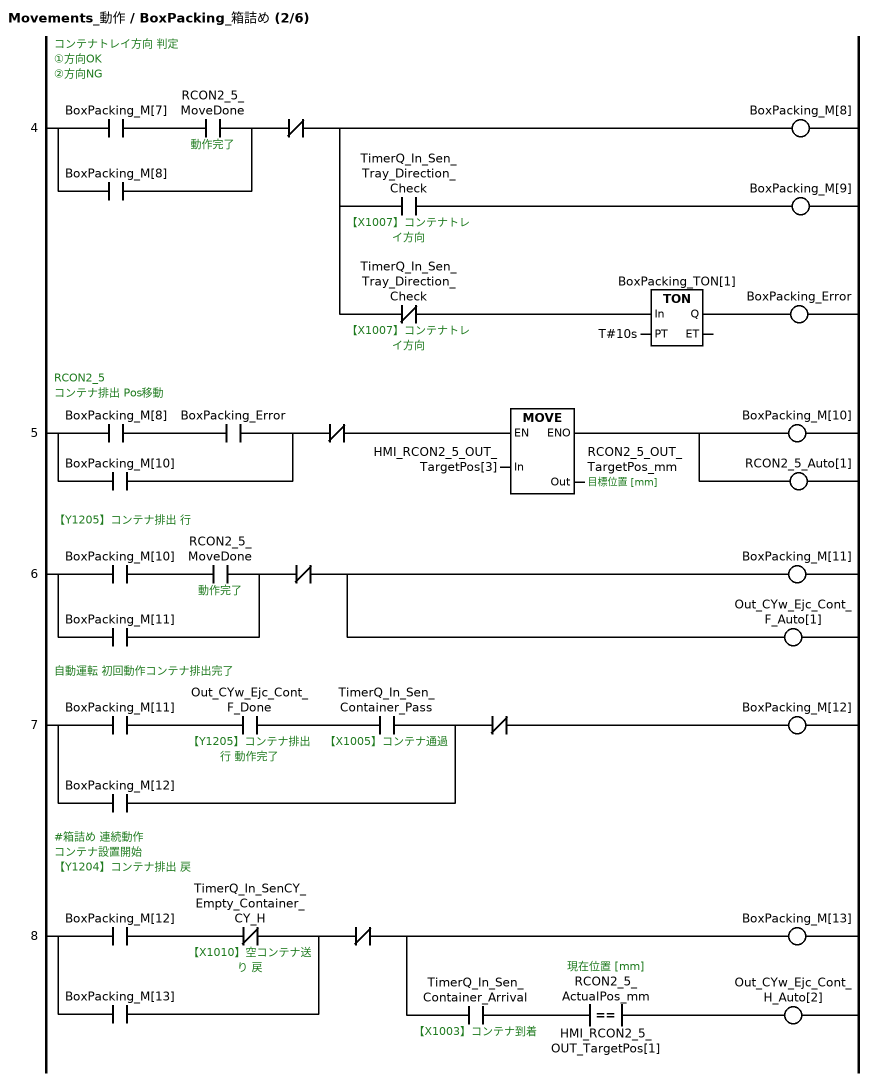
(* Rung 4: コンテナトレイ方向 判定 / ①方向OK / ②方向NG *)
_p141 := ((BoxPacking_M[7] AND RCON2_5_MoveDone) OR BoxPacking_M[8]) AND NOT ();
BoxPacking_M[8] := _p141;
BoxPacking_M[9] := _p141 AND TimerQ_In_Sen_Tray_Direction_Check;
BoxPacking_TON[1](In := _p141 AND NOT TimerQ_In_Sen_Tray_Direction_Check, PT := T#10s);
BoxPacking_Error := BoxPacking_TON[1].Q;
(* Rung 5: RCON2_5 / コンテナ排出 Pos移動 *)
IF ((BoxPacking_M[8] AND BoxPacking_Error) OR BoxPacking_M[10]) AND NOT () THEN
    RCON2_5_OUT_TargetPos_mm := HMI_RCON2_5_OUT_TargetPos[3];
END_IF;
_p142 := ((BoxPacking_M[8] AND BoxPacking_Error) OR BoxPacking_M[10]) AND NOT ();
BoxPacking_M[10] := _p142;
RCON2_5_Auto[1] := _p142;
(* Rung 6: 【Y1205】コンテナ排出 行 *)
_p143 := ((BoxPacking_M[10] AND RCON2_5_MoveDone) OR BoxPacking_M[11]) AND NOT ();
BoxPacking_M[11] := _p143;
Out_CYw_Ejc_Cont_F_Auto[1] := _p143;
(* Rung 7: 自動運転 初回動作コンテナ排出完了 *)
BoxPacking_M[12] := ((BoxPacking_M[11] AND Out_CYw_Ejc_Cont_F_Done AND TimerQ_In_Sen_Container_Pass) OR BoxPacking_M[12]) AND NOT ();
(* Rung 8: #箱詰め 連続動作 / コンテナ設置開始 / 【Y1204】コンテナ排出 戻 *)
_p144 := ((BoxPacking_M[12] AND NOT TimerQ_In_SenCY_Empty_Container_CY_H) OR BoxPacking_M[13]) AND NOT ();
BoxPacking_M[13] := _p144;
Out_CYw_Ejc_Cont_H_Auto[2] := _p144 AND TimerQ_In_Sen_Container_Arrival AND (RCON2_5_ActualPos_mm = HMI_RCON2_5_OUT_TargetPos[1]);

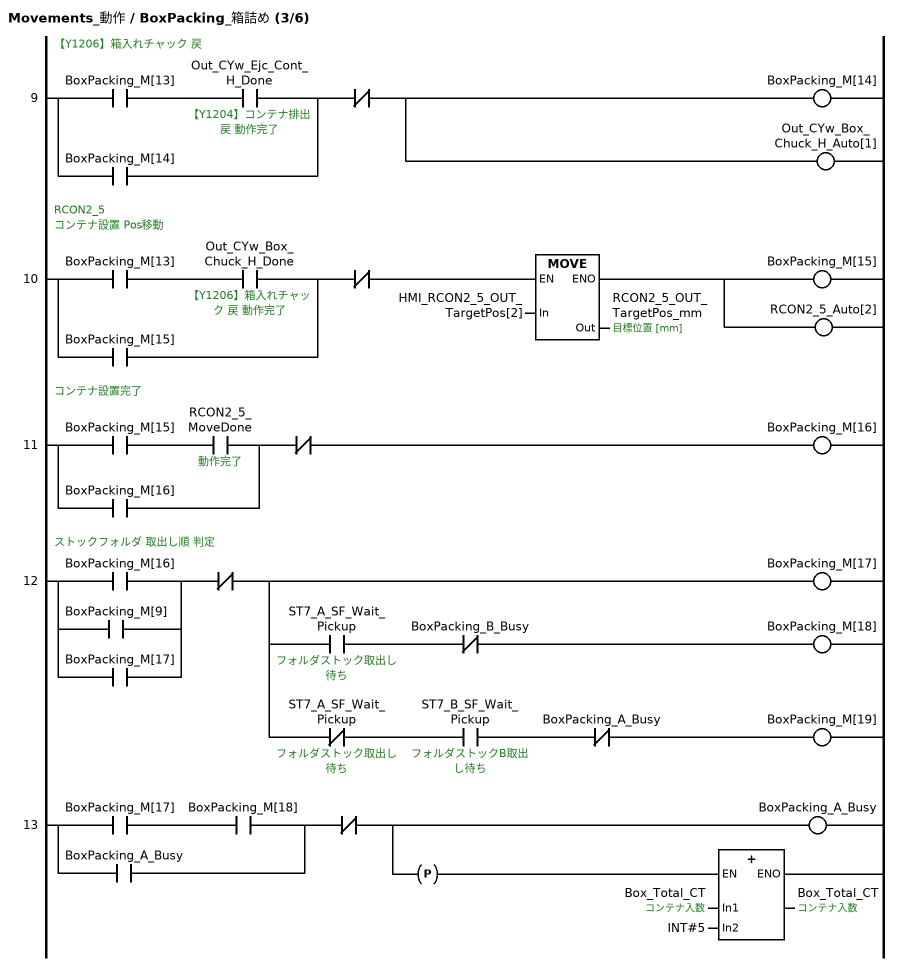
(* Rung 9: 【Y1206】箱入れチャック 戻 *)
_p145 := ((BoxPacking_M[13] AND Out_CYw_Ejc_Cont_H_Done) OR BoxPacking_M[14]) AND NOT ();
BoxPacking_M[14] := _p145;
Out_CYw_Box_Chuck_H_Auto[1] := _p145;
(* Rung 10: RCON2_5 / コンテナ設置 Pos移動 *)
IF ((BoxPacking_M[13] AND Out_CYw_Box_Chuck_H_Done) OR BoxPacking_M[15]) AND NOT () THEN
    RCON2_5_OUT_TargetPos_mm := HMI_RCON2_5_OUT_TargetPos[2];
END_IF;
_p146 := ((BoxPacking_M[13] AND Out_CYw_Box_Chuck_H_Done) OR BoxPacking_M[15]) AND NOT ();
BoxPacking_M[15] := _p146;
RCON2_5_Auto[2] := _p146;
(* Rung 11: コンテナ設置完了 *)
BoxPacking_M[16] := ((BoxPacking_M[15] AND RCON2_5_MoveDone) OR BoxPacking_M[16]) AND NOT ();
(* Rung 12: ストックフォルダ 取出し順 判定 *)
_p147 := (BoxPacking_M[16] OR BoxPacking_M[9] OR BoxPacking_M[17]) AND NOT ();
BoxPacking_M[17] := _p147;
BoxPacking_M[18] := _p147 AND ST7_A_SF_Wait_Pickup AND NOT BoxPacking_B_Busy;
BoxPacking_M[19] := _p147 AND NOT ST7_A_SF_Wait_Pickup AND ST7_B_SF_Wait_Pickup AND NOT BoxPacking_A_Busy;
(* Rung 13 *)
_p148 := ((BoxPacking_M[17] AND BoxPacking_M[18]) OR BoxPacking_A_Busy) AND NOT ();
BoxPacking_A_Busy := _p148;
_e149(CLK := _p148);
IF _e149.Q THEN Box_Total_CT := Box_Total_CT + INT#5; END_IF;

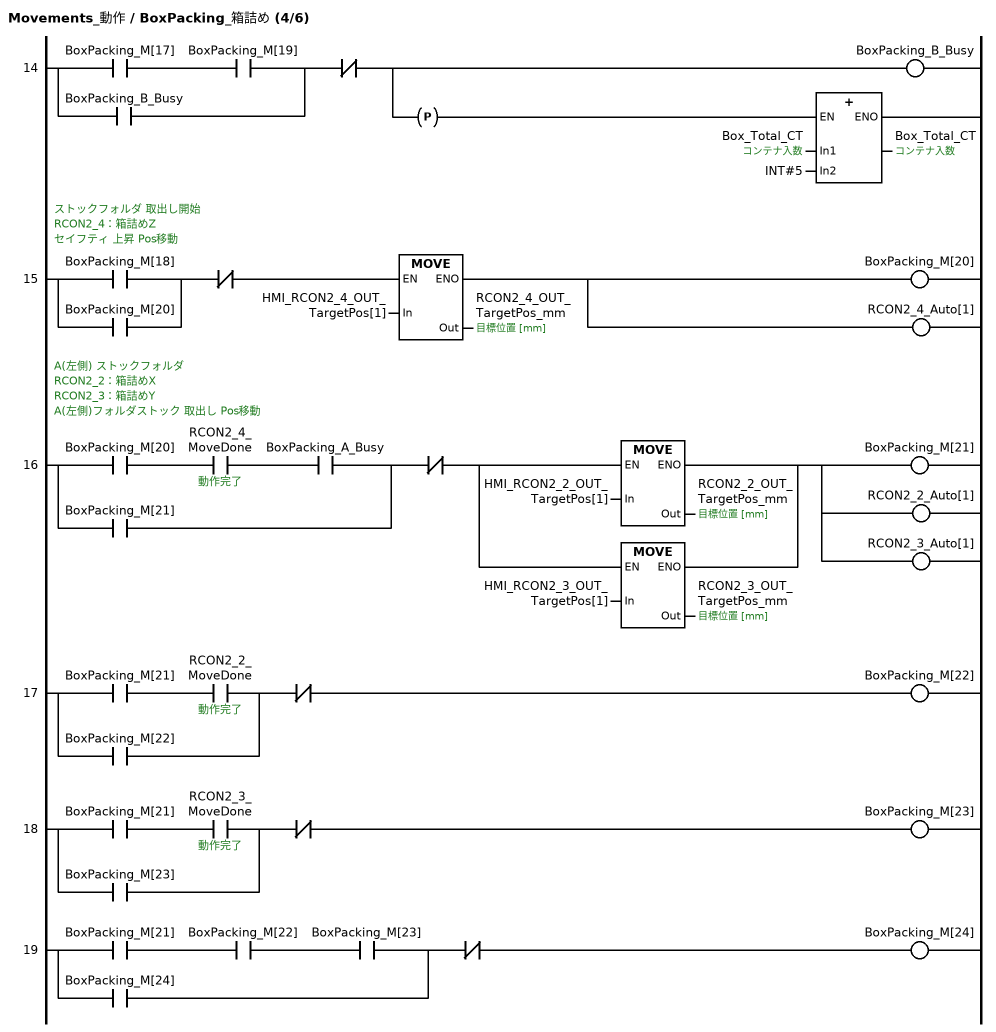
(* Rung 14 *)
_p150 := ((BoxPacking_M[17] AND BoxPacking_M[19]) OR BoxPacking_B_Busy) AND NOT ();
BoxPacking_B_Busy := _p150;
_e151(CLK := _p150);
IF _e151.Q THEN Box_Total_CT := Box_Total_CT + INT#5; END_IF;
(* Rung 15: ストックフォルダ 取出し開始 / RCON2_4：箱詰めZ / セイフティ 上昇 Pos移動 *)
IF (BoxPacking_M[18] OR BoxPacking_M[20]) AND NOT () THEN
    RCON2_4_OUT_TargetPos_mm := HMI_RCON2_4_OUT_TargetPos[1];
END_IF;
_p152 := (BoxPacking_M[18] OR BoxPacking_M[20]) AND NOT ();
BoxPacking_M[20] := _p152;
RCON2_4_Auto[1] := _p152;
(* Rung 16: A(左側) ストックフォルダ / RCON2_2：箱詰めX / RCON2_3：箱詰めY / A(左側)フォルダストック 取出し Pos移動 *)
_p153 := ((BoxPacking_M[20] AND RCON2_4_MoveDone AND BoxPacking_A_Busy) OR BoxPacking_M[21]) AND NOT ();
IF _p153 THEN
    RCON2_2_OUT_TargetPos_mm := HMI_RCON2_2_OUT_TargetPos[1];
    RCON2_3_OUT_TargetPos_mm := HMI_RCON2_3_OUT_TargetPos[1];
END_IF;
BoxPacking_M[21] := _p153;
RCON2_2_Auto[1] := _p153;
RCON2_3_Auto[1] := _p153;
(* Rung 17 *)
BoxPacking_M[22] := ((BoxPacking_M[21] AND RCON2_2_MoveDone) OR BoxPacking_M[22]) AND NOT ();
(* Rung 18 *)
BoxPacking_M[23] := ((BoxPacking_M[21] AND RCON2_3_MoveDone) OR BoxPacking_M[23]) AND NOT ();
(* Rung 19 *)
BoxPacking_M[24] := ((BoxPacking_M[21] AND BoxPacking_M[22] AND BoxPacking_M[23]) OR BoxPacking_M[24]) AND NOT ();

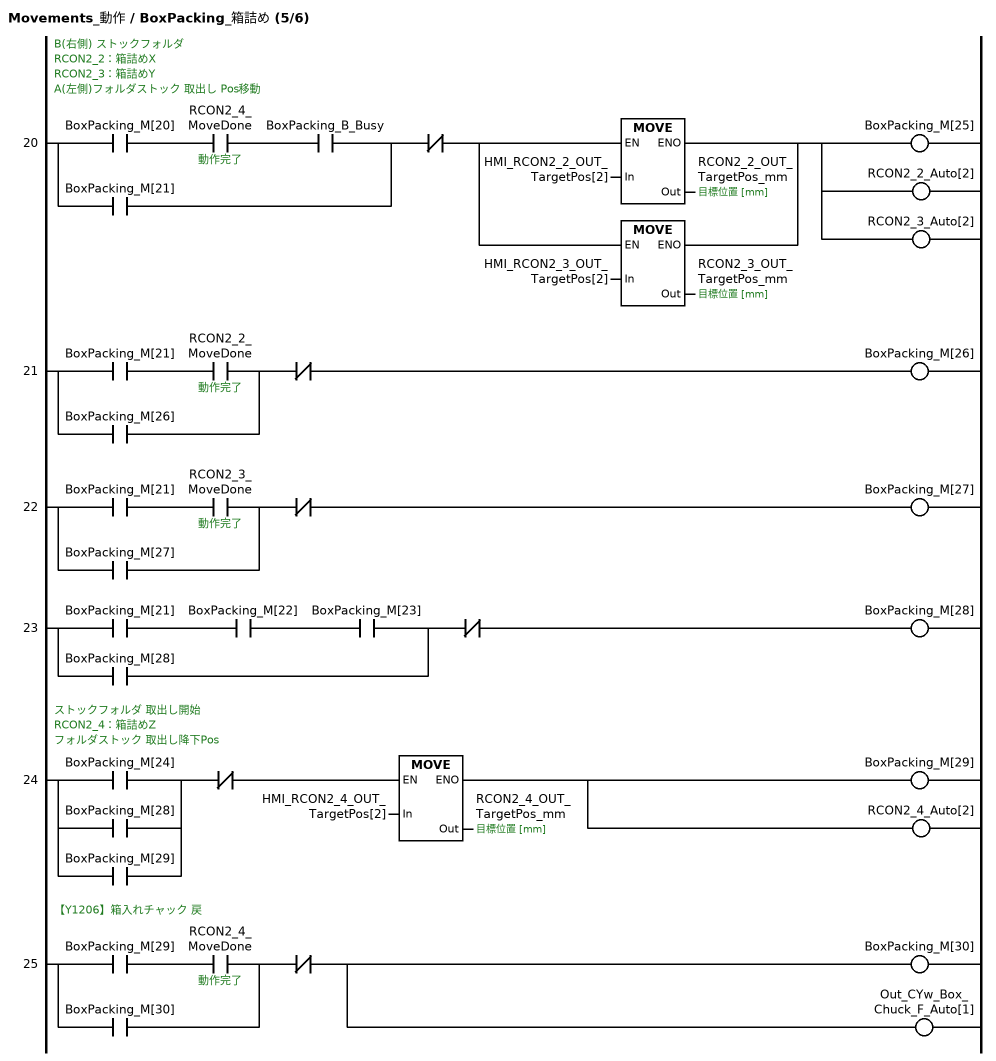
(* Rung 20: B(右側) ストックフォルダ / RCON2_2：箱詰めX / RCON2_3：箱詰めY / A(左側)フォルダストック 取出し Pos移動 *)
_p154 := ((BoxPacking_M[20] AND RCON2_4_MoveDone AND BoxPacking_B_Busy) OR BoxPacking_M[21]) AND NOT ();
IF _p154 THEN
    RCON2_2_OUT_TargetPos_mm := HMI_RCON2_2_OUT_TargetPos[2];
    RCON2_3_OUT_TargetPos_mm := HMI_RCON2_3_OUT_TargetPos[2];
END_IF;
BoxPacking_M[25] := _p154;
RCON2_2_Auto[2] := _p154;
RCON2_3_Auto[2] := _p154;
(* Rung 21 *)
BoxPacking_M[26] := ((BoxPacking_M[21] AND RCON2_2_MoveDone) OR BoxPacking_M[26]) AND NOT ();
(* Rung 22 *)
BoxPacking_M[27] := ((BoxPacking_M[21] AND RCON2_3_MoveDone) OR BoxPacking_M[27]) AND NOT ();
(* Rung 23 *)
BoxPacking_M[28] := ((BoxPacking_M[21] AND BoxPacking_M[22] AND BoxPacking_M[23]) OR BoxPacking_M[28]) AND NOT ();
(* Rung 24: ストックフォルダ 取出し開始 / RCON2_4：箱詰めZ / フォルダストック 取出し降下Pos *)
IF (BoxPacking_M[24] OR BoxPacking_M[28] OR BoxPacking_M[29]) AND NOT () THEN
    RCON2_4_OUT_TargetPos_mm := HMI_RCON2_4_OUT_TargetPos[2];
END_IF;
_p155 := (BoxPacking_M[24] OR BoxPacking_M[28] OR BoxPacking_M[29]) AND NOT ();
BoxPacking_M[29] := _p155;
RCON2_4_Auto[2] := _p155;
(* Rung 25: 【Y1206】箱入れチャック 戻 *)
_p156 := ((BoxPacking_M[29] AND RCON2_4_MoveDone) OR BoxPacking_M[30]) AND NOT ();
BoxPacking_M[30] := _p156;
Out_CYw_Box_Chuck_F_Auto[1] := _p156;

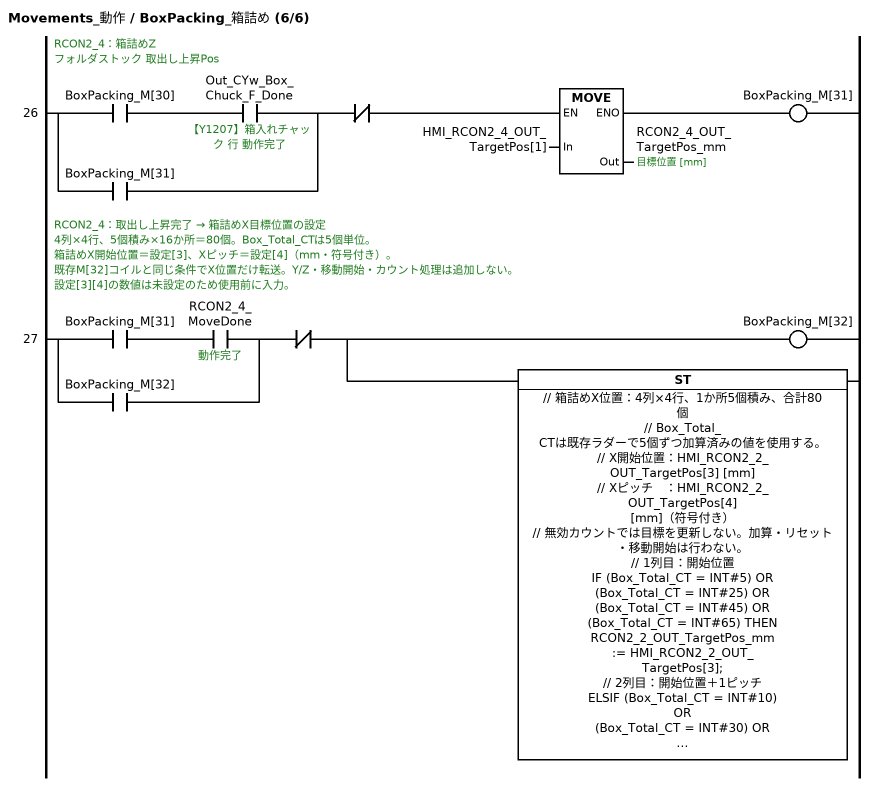
(* Rung 26: RCON2_4：箱詰めZ / フォルダストック 取出し上昇Pos *)
IF ((BoxPacking_M[30] AND Out_CYw_Box_Chuck_F_Done) OR BoxPacking_M[31]) AND NOT () THEN
    RCON2_4_OUT_TargetPos_mm := HMI_RCON2_4_OUT_TargetPos[1];
END_IF;
BoxPacking_M[31] := ((BoxPacking_M[30] AND Out_CYw_Box_Chuck_F_Done) OR BoxPacking_M[31]) AND NOT ();
(* Rung 27: RCON2_4：取出し上昇完了 → 箱詰めX目標位置の設定 / 4列×4行、5個積み×16か所＝80個。Box_Total_CTは5個単位。 / 箱詰めX開始位置＝設定[3]、Xピッチ＝設定[4]（mm・符号付き）。 / 既存M[32]コイルと同じ条件でX位置だけ転送。Y/Z・移動開始・カウント処理は追加しない。 / 設定[3][4]の数値は未設定のため使用前に入力。 *)
_p157 := ((BoxPacking_M[31] AND RCON2_4_MoveDone) OR BoxPacking_M[32]) AND NOT ();
BoxPacking_M[32] := _p157;
IF _p157 THEN
    // 箱詰めX位置：4列×4行、1か所5個積み、合計80個
    // Box_Total_CTは既存ラダーで5個ずつ加算済みの値を使用する。
    // X開始位置：HMI_RCON2_2_OUT_TargetPos[3] [mm]
    // Xピッチ　：HMI_RCON2_2_OUT_TargetPos[4] [mm]（符号付き）
    // 無効カウントでは目標を更新しない。加算・リセット・移動開始は行わない。
    
    // 1列目：開始位置
    IF (Box_Total_CT = INT#5) OR
       (Box_Total_CT = INT#25) OR
       (Box_Total_CT = INT#45) OR
       (Box_Total_CT = INT#65) THEN
    
        RCON2_2_OUT_TargetPos_mm := HMI_RCON2_2_OUT_TargetPos[3];
    
    // 2列目：開始位置＋1ピッチ
    ELSIF (Box_Total_CT = INT#10) OR
          (Box_Total_CT = INT#30) OR
          (Box_Total_CT = INT#50) OR
          (Box_Total_CT = INT#70) THEN
    
        RCON2_2_OUT_TargetPos_mm :=
            HMI_RCON2_2_OUT_TargetPos[3] +
            HMI_RCON2_2_OUT_TargetPos[4];
    
    // 3列目：開始位置＋2ピッチ
    ELSIF (Box_Total_CT = INT#15) OR
          (Box_Total_CT = INT#35) OR
          (Box_Total_CT = INT#55) OR
          (Box_Total_CT = INT#75) THEN
    
        RCON2_2_OUT_TargetPos_mm :=
            HMI_RCON2_2_OUT_TargetPos[3] +
            HMI_RCON2_2_OUT_TargetPos[4] * LREAL#2.0;
    
    // 4列目：開始位置＋3ピッチ
    ELSIF (Box_Total_CT = INT#20) OR
          (Box_Total_CT = INT#40) OR
          (Box_Total_CT = INT#60) OR
          (Box_Total_CT = INT#80) THEN
    
        RCON2_2_OUT_TargetPos_mm :=
            HMI_RCON2_2_OUT_TargetPos[3] +
            HMI_RCON2_2_OUT_TargetPos[4] * LREAL#3.0;
    END_IF;
END_IF;
END_PROGRAM

PROGRAM OtherDevice_外部機器
VAR
    FH_M : BOOL;
    GT2_M : BOOL;
    IAI_M : BOOL;  (* 旧ダミーマーカー（ST許可ではない） *)
    HMI_M : BOOL;
    FH_A_ST1_M : ARRAY[0..99] OF Bool;  (* [1] ST1 FH測定中; [5] ST1 測定完了 *)
    FH_A_ST1_OK : BOOL;  (* ST1 OK判定 *)
    FH_A_ST1_NG : BOOL;  (* ST1 NG 判定 *)
    FH_A_ST1_TON : ARRAY[0..99] OF TON;
    FH_A_ST1_TOF : ARRAY[0..99] OF TOF;
    ４ : UINT;
    ConvWordIndex : INT;  (* 作業用 ワード番号 *)
    ConvAxisIndex : INT;  (* 作業用 軸番号（RCON1:1～6／RCON2:1～5） *)
    ConvBase : INT;  (* 作業用 軸先頭ワード番号 *)
    ConvDWord : DWORD;  (* 作業用 32bit分割・結合 *)
    ConvPos : DINT;  (* 作業用 目標位置 [0.01mm・符号付き] *)
    ConvBand : UDINT;  (* 作業用 位置決め幅 [0.01mm] *)
    ConvSpeed : UINT;  (* 作業用 速度送信値 *)
    ConvAccDec : UINT;  (* 作業用 共通加減速 [0.01G] *)
    ConvPush : UINT;  (* 作業用 押付け制限 [255=100%] *)
    ConvScaled : LREAL;  (* 作業用 換算後の小数値 *)
    ConvWord : WORD;  (* 作業用 16bitワード *)
    ConvUnitOK : BOOL;  (* 作業用 速度単位正常 *)
    RCON1_1_TOF : ARRAY[0..99] OF TOF;  (* 開始要求100ms保持; [1] 開始要求100ms保持 *)
    RCON1_1_TON : ARRAY[0..99] OF TON;  (* 準備・完了タイマー; [1] 準備100ms確認; [2] 動作完了100ms保持 *)
    Stm_A_Rev_Axis000_ZeroSet : MC_SetPosition;
    Stm_A_Rev_Axis000_HomeWithParameter : MC_HomeWithParameter;
    Stm_A_Rev_Axis000_Power : MC_Power;  (* A(左側)ステッピングモータ000 電源ON状態 *)
    Stm_A_Rev_Axis000_MoveAbsolute : MC_MoveAbsolute;
    Stm_A_Rev_Axis000_MoveVel : LREAL;  (* 動作速度 *)
    Stm_A_Rev_Axis000_MoveAcc : LREAL;  (* 動作加速度 *)
    Stm_A_Rev_Axis000_MoveDec : LREAL;  (* 動作減速度 *)
    Stm_A_Rev_Axis000_MoveBusy : BOOL;  (* 動作中 *)
    Stm_A_Rev_Axis000_TON : ARRAY[0..99] OF TON;
    FH_A_ST5_M : ARRAY[0..99] OF Bool;  (* A(左側) ST5 FH工程; [1] A(左側) ST5 測定要求; [2] A(左側) ST5 シーン切替; [3] A(左側) ST5 コマンド完了; [4] A(左側) ST5 測定トリガー; [5] A(左側) ST5 測定完了; [6] A(左側) ST5 OK保持; [7] A(左側) ST5 NG／完了保持 *)
    FH_A_ST5_OK : BOOL;  (* A(左側) ST5 OK判定 *)
    FH_A_ST5_NG : BOOL;  (* A(左側) ST5 NG判定 *)
    FH_A_ST5_TON : ARRAY[0..99] OF TON;  (* A(左側) ST5 FH遅延タイマー *)
    FH_A_ST5_TOF : ARRAY[0..99] OF TOF;  (* A(左側) ST5 FHトリガ保持; [1] A(左側) ST5 トリガー100ms *)
    Stm_A_Rev_Axis001_ZeroSet : MC_SetPosition;  (* A(左側) ST6 反転2 位置ゼロ設定 *)
    Stm_A_Rev_Axis001_HomeWithParameter : MC_HomeWithParameter;  (* A(左側) ST6 反転2 原点復帰FB *)
    Stm_A_Rev_Axis001_Power : MC_Power;  (* A(左側) ST6 反転2 電源ON状態 *)
    Stm_A_Rev_Axis001_MoveAbsolute : MC_MoveAbsolute;  (* A(左側) ST6 反転2 絶対位置決めFB *)
    Stm_A_Rev_Axis001_MoveVel : LREAL;  (* A(左側) ST6 反転2 速度 *)
    Stm_A_Rev_Axis001_MoveAcc : LREAL;  (* A(左側) ST6 反転2 加速度 *)
    Stm_A_Rev_Axis001_MoveDec : LREAL;  (* A(左側) ST6 反転2 減速度 *)
    Stm_A_Rev_Axis001_MoveBusy : BOOL;  (* A(左側) ST6 反転2 移動中 *)
    Stm_A_Rev_Axis001_TON : ARRAY[0..99] OF TON;  (* A(左側) ST6 反転2 完了保持タイマー *)
    RCON1_2_TOF : ARRAY[0..99] OF TOF;  (* 開始要求100ms保持; [1] 開始要求100ms保持 *)
    RCON1_2_TON : ARRAY[0..99] OF TON;  (* 準備・完了タイマー; [1] 準備100ms確認; [2] 動作完了100ms保持 *)
    RCON1_3_TOF : ARRAY[0..99] OF TOF;  (* 開始要求100ms保持; [1] 開始要求100ms保持 *)
    RCON1_3_TON : ARRAY[0..99] OF TON;  (* 準備・完了タイマー; [1] 準備100ms確認; [2] 動作完了100ms保持 *)
    RCON1_4_TOF : ARRAY[0..99] OF TOF;  (* 開始要求100ms保持; [1] 開始要求100ms保持 *)
    RCON1_4_TON : ARRAY[0..99] OF TON;  (* 準備・完了タイマー; [1] 準備100ms確認; [2] 動作完了100ms保持 *)
    RCON1_5_TOF : ARRAY[0..99] OF TOF;  (* 開始要求100ms保持; [1] 開始要求100ms保持 *)
    RCON1_5_TON : ARRAY[0..99] OF TON;  (* 準備・完了タイマー; [1] 準備100ms確認; [2] 動作完了100ms保持 *)
    RCON1_6_TOF : ARRAY[0..99] OF TOF;  (* 開始要求100ms保持; [1] 開始要求100ms保持 *)
    RCON1_6_TON : ARRAY[0..99] OF TON;  (* 準備・完了タイマー; [1] 準備100ms確認; [2] 動作完了100ms保持 *)
    RCON2_1_TOF : ARRAY[0..99] OF TOF;  (* 開始要求100ms保持; [1] 開始要求100ms保持 *)
    RCON2_1_TON : ARRAY[0..99] OF TON;  (* 準備・完了タイマー; [1] 準備100ms確認; [2] 動作完了100ms保持 *)
    RCON2_2_TOF : ARRAY[0..99] OF TOF;  (* 開始要求100ms保持; [1] 開始要求100ms保持 *)
    RCON2_2_TON : ARRAY[0..99] OF TON;  (* 準備・完了タイマー; [1] 準備100ms確認; [2] 動作完了100ms保持 *)
    RCON2_3_TOF : ARRAY[0..99] OF TOF;  (* 開始要求100ms保持; [1] 開始要求100ms保持 *)
    RCON2_3_TON : ARRAY[0..99] OF TON;  (* 準備・完了タイマー; [1] 準備100ms確認; [2] 動作完了100ms保持 *)
    RCON2_4_TOF : ARRAY[0..99] OF TOF;  (* 開始要求100ms保持; [1] 開始要求100ms保持 *)
    RCON2_4_TON : ARRAY[0..99] OF TON;  (* 準備・完了タイマー; [1] 準備100ms確認; [2] 動作完了100ms保持 *)
    RCON2_5_TOF : ARRAY[0..99] OF TOF;  (* 開始要求100ms保持; [1] 開始要求100ms保持 *)
    RCON2_5_TON : ARRAY[0..99] OF TON;  (* 準備・完了タイマー; [1] 準備100ms確認; [2] 動作完了100ms保持 *)
END_VAR
VAR_EXTERNAL
    HMI_MessageNo : ARRAY[0..9] OF UINT;
    HMI_Message : ARRAY[0..9] OF String[256];
    HMI_Language : BOOL;
    FH_Line0_Trigger_Ready_1 : BOOL;
    FH_Line0_Trigger_1 : BOOL;
    M9999 : BOOL;
    FH_Line0_Busy_1 : BOOL;
    FH_Line0_Result_Notification_1 : BOOL;
    FH_Line0_DINT_Result_Data_0_1 : DINT;
    FH_Line0_DINT_Result_Data_1_1 : DINT;
    FH_Line0_DINT_Result_Data_2_1 : DINT;
    FH_Line0_Command_Code_1 : DWORD;
    FH_Line0_Command_Request_1 : BOOL;
    FH_Line0_Command_Completion_1 : BOOL;
    MdlChg : BOOL;  (* 機種切替：ON【GA120】 OFF【GA90】 *)
    FH_Line0_Error_Status_1 : BOOL;
    FH_A_ST1_Auto : BOOL;  (* ST1 FH測定開始 *)
    FH_A_ST1_Manual : BOOL;  (* ST1 *)
    Pause : ARRAY[0..99] OF Bool;  (* [3] FH A(左側) ST1; [9] FH A(左側) ST5; [10] FH B(右側) ST1; [11] FH B(右側) ST5; [12] A(左側) ST6 反転2 ワーク不一致 *)
    FH_A_ST1_Done : BOOL;  (* ST1 画像検査完了 *)
    Station_A_Data : ARRAY[0..8] OF sData;
    DLEP1_OUT : ARRAY[0..79] OF BOOL;
    DLEP2_OUT : ARRAY[0..79] OF BOOL;
    DLEP1_IN : ARRAY[0..167] OF byte;
    DLEP2_IN : ARRAY[0..167] OF byte;
    DLEP2_IN_Error : BOOL;  (* B(右側)センサエラー *)
    DLEP1_IN_Error : BOOL;  (* A(右側)センサエラー *)
    GT2_A_CurrentVal : INT;  (* A(左側) 測定値 *)
    GT2_B_CurrentVal : INT;  (* B(右側) 測定値 *)
    Hgt_A_Ins_Data : LREAL;  (* A測定データに変換 *)
    Hgt_B_Ins_Data : LREAL;
    Hgt_A_ComputedValueData : LREAL;  (* A測定データ+13.000mm 算定データ *)
    Hgt_B_ComputedValueData : LREAL;  (* B測定データ+13.000mm 算定データ *)
    E001_In_IN00_2004_01 : UINT;  (* IN00 GW状態 *)
    E001_In_IN01_2004_02 : UINT;  (* IN01 軸リンク状態 *)
    E001_In_IN02_2004_03 : UINT;  (* IN02 電源状態0 *)
    E001_In_IN03_2004_04 : UINT;  (* IN03 電源状態1 *)
    E001_In_IN04_2004_05 : UINT;  (* IN04 電源状態2 *)
    E001_In_IN05_2004_06 : UINT;  (* IN05 電源状態3 *)
    E001_In_IN06_2004_07 : UINT;  (* IN06 電源状態4（構成依存） *)
    E001_In_IN07_2004_08 : UINT;  (* IN07 予約（使用禁止） *)
    E001_In_IN08_2004_09 : UINT;  (* IN08 現在位置 下位 [0.01mm] *)
    E001_In_IN09_2004_0A : UINT;  (* IN09 現在位置 上位 [0.01mm] *)
    E001_In_IN10_2004_0B : UINT;  (* IN10 指令電流 下位 [mA] *)
    E001_In_IN11_2004_0C : UINT;  (* IN11 指令電流 上位 [mA] *)
    E001_In_IN12_2004_0D : UINT;  (* IN12 現在速度 [実機単位・符号付き] *)
    E001_In_IN13_2004_0E : UINT;  (* IN13 予約（使用禁止） *)
    E001_In_IN14_2004_0F : UINT;  (* IN14 軸異常コード *)
    E001_In_IN15_2004_10 : UINT;  (* IN15 状態信号（PEND/SV等） *)
    E001_In_IN16_2004_11 : UINT;  (* IN16 現在位置 下位 [0.01mm] *)
    E001_In_IN17_2004_12 : UINT;  (* IN17 現在位置 上位 [0.01mm] *)
    E001_In_IN18_2004_13 : UINT;  (* IN18 指令電流 下位 [mA] *)
    E001_In_IN19_2004_14 : UINT;  (* IN19 指令電流 上位 [mA] *)
    E001_In_IN20_2004_15 : UINT;  (* IN20 現在速度 [実機単位・符号付き] *)
    E001_In_IN21_2004_16 : UINT;  (* IN21 予約（使用禁止） *)
    E001_In_IN22_2004_17 : UINT;  (* IN22 軸異常コード *)
    E001_In_IN23_2004_18 : UINT;  (* IN23 状態信号（PEND/SV等） *)
    E001_In_IN24_2004_19 : UINT;  (* IN24 現在位置 下位 [0.01mm] *)
    E001_In_IN25_2004_1A : UINT;  (* IN25 現在位置 上位 [0.01mm] *)
    E001_In_IN26_2004_1B : UINT;  (* IN26 指令電流 下位 [mA] *)
    E001_In_IN27_2004_1C : UINT;  (* IN27 指令電流 上位 [mA] *)
    E001_In_IN28_2004_1D : UINT;  (* IN28 現在速度 [実機単位・符号付き] *)
    E001_In_IN29_2004_1E : UINT;  (* IN29 予約（使用禁止） *)
    E001_In_IN30_2004_1F : UINT;  (* IN30 軸異常コード *)
    E001_In_IN31_2004_20 : UINT;  (* IN31 状態信号（PEND/SV等） *)
    E001_In_IN32_2004_21 : UINT;  (* IN32 現在位置 下位 [0.01mm] *)
    E001_In_IN33_2004_22 : UINT;  (* IN33 現在位置 上位 [0.01mm] *)
    E001_In_IN34_2004_23 : UINT;  (* IN34 指令電流 下位 [mA] *)
    E001_In_IN35_2004_24 : UINT;  (* IN35 指令電流 上位 [mA] *)
    E001_In_IN36_2004_25 : UINT;  (* IN36 現在速度 [実機単位・符号付き] *)
    E001_In_IN37_2004_26 : UINT;  (* IN37 予約（使用禁止） *)
    E001_In_IN38_2004_27 : UINT;  (* IN38 軸異常コード *)
    E001_In_IN39_2004_28 : UINT;  (* IN39 状態信号（PEND/SV等） *)
    E001_In_IN40_2004_29 : UINT;  (* IN40 現在位置 下位 [0.01mm] *)
    E001_In_IN41_2004_2A : UINT;  (* IN41 現在位置 上位 [0.01mm] *)
    E001_In_IN42_2004_2B : UINT;  (* IN42 指令電流 下位 [mA] *)
    E001_In_IN43_2004_2C : UINT;  (* IN43 指令電流 上位 [mA] *)
    E001_In_IN44_2004_2D : UINT;  (* IN44 現在速度 [実機単位・符号付き] *)
    E001_In_IN45_2004_2E : UINT;  (* IN45 予約（使用禁止） *)
    E001_In_IN46_2004_2F : UINT;  (* IN46 軸異常コード *)
    E001_In_IN47_2004_30 : UINT;  (* IN47 状態信号（PEND/SV等） *)
    E001_In_IN48_2004_31 : UINT;  (* IN48 現在位置 下位 [0.01mm] *)
    E001_In_IN49_2004_32 : UINT;  (* IN49 現在位置 上位 [0.01mm] *)
    E001_In_IN50_2004_33 : UINT;  (* IN50 指令電流 下位 [mA] *)
    E001_In_IN51_2004_34 : UINT;  (* IN51 指令電流 上位 [mA] *)
    E001_In_IN52_2004_35 : UINT;  (* IN52 現在速度 [実機単位・符号付き] *)
    E001_In_IN53_2004_36 : UINT;  (* IN53 予約（使用禁止） *)
    E001_In_IN54_2004_37 : UINT;  (* IN54 軸異常コード *)
    E001_In_IN55_2004_38 : UINT;  (* IN55 状態信号（PEND/SV等） *)
    E001_In_IN56_2004_39 : UINT;  (* IN56 112Byte範囲外（未割付・不使用） *)
    E001_In_IN57_2004_3A : UINT;  (* IN57 112Byte範囲外（未割付・不使用） *)
    E001_In_IN58_2004_3B : UINT;  (* IN58 112Byte範囲外（未割付・不使用） *)
    E001_In_IN59_2004_3C : UINT;  (* IN59 112Byte範囲外（未割付・不使用） *)
    E001_In_IN60_2004_3D : UINT;  (* IN60 112Byte範囲外（未割付・不使用） *)
    E001_In_IN61_2004_3E : UINT;  (* IN61 112Byte範囲外（未割付・不使用） *)
    E001_In_IN62_2004_3F : UINT;  (* IN62 112Byte範囲外（未割付・不使用） *)
    E001_In_IN63_2004_40 : UINT;  (* IN63 112Byte範囲外（未割付・不使用） *)
    E001_In_IN64_2004_41 : UINT;  (* IN64 112Byte範囲外（未割付・不使用） *)
    E001_In_IN65_2004_42 : UINT;  (* IN65 112Byte範囲外（未割付・不使用） *)
    E001_In_IN66_2004_43 : UINT;  (* IN66 112Byte範囲外（未割付・不使用） *)
    E001_In_IN67_2004_44 : UINT;  (* IN67 112Byte範囲外（未割付・不使用） *)
    E001_In_IN68_2004_45 : UINT;  (* IN68 112Byte範囲外（未割付・不使用） *)
    E001_In_IN69_2004_46 : UINT;  (* IN69 112Byte範囲外（未割付・不使用） *)
    E001_In_IN70_2004_47 : UINT;  (* IN70 112Byte範囲外（未割付・不使用） *)
    E001_In_IN71_2004_48 : UINT;  (* IN71 112Byte範囲外（未割付・不使用） *)
    E001_Out_OUT00_2003_01 : UINT;  (* OUT00 共通制御（MON/RTE） *)
    E001_Out_OUT08_2003_09 : UINT;  (* OUT08 目標位置 下位 [0.01mm] *)
    E001_Out_OUT09_2003_0A : UINT;  (* OUT09 目標位置 上位 [0.01mm] *)
    E001_Out_OUT10_2003_0B : UINT;  (* OUT10 位置決め幅 下位 [0.01mm] *)
    E001_Out_OUT11_2003_0C : UINT;  (* OUT11 位置決め幅 上位 [0.01mm] *)
    E001_Out_OUT12_2003_0D : UINT;  (* OUT12 速度指令 [実機単位] *)
    E001_Out_OUT13_2003_0E : UINT;  (* OUT13 共通加減速 [0.01G] *)
    E001_Out_OUT14_2003_0F : UINT;  (* OUT14 押付け制限 [255=100%] *)
    E001_Out_OUT15_2003_10 : UINT;  (* OUT15 制御信号（DSTR/SON等） *)
    E001_Out_OUT16_2003_11 : UINT;  (* OUT16 目標位置 下位 [0.01mm] *)
    E001_Out_OUT17_2003_12 : UINT;  (* OUT17 目標位置 上位 [0.01mm] *)
    E001_Out_OUT18_2003_13 : UINT;  (* OUT18 位置決め幅 下位 [0.01mm] *)
    E001_Out_OUT19_2003_14 : UINT;  (* OUT19 位置決め幅 上位 [0.01mm] *)
    E001_Out_OUT20_2003_15 : UINT;  (* OUT20 速度指令 [実機単位] *)
    E001_Out_OUT21_2003_16 : UINT;  (* OUT21 共通加減速 [0.01G] *)
    E001_Out_OUT22_2003_17 : UINT;  (* OUT22 押付け制限 [255=100%] *)
    E001_Out_OUT23_2003_18 : UINT;  (* OUT23 制御信号（DSTR/SON等） *)
    E001_Out_OUT24_2003_19 : UINT;  (* OUT24 目標位置 下位 [0.01mm] *)
    E001_Out_OUT25_2003_1A : UINT;  (* OUT25 目標位置 上位 [0.01mm] *)
    E001_Out_OUT26_2003_1B : UINT;  (* OUT26 位置決め幅 下位 [0.01mm] *)
    E001_Out_OUT27_2003_1C : UINT;  (* OUT27 位置決め幅 上位 [0.01mm] *)
    E001_Out_OUT28_2003_1D : UINT;  (* OUT28 速度指令 [実機単位] *)
    E001_Out_OUT29_2003_1E : UINT;  (* OUT29 共通加減速 [0.01G] *)
    E001_Out_OUT30_2003_1F : UINT;  (* OUT30 押付け制限 [255=100%] *)
    E001_Out_OUT31_2003_20 : UINT;  (* OUT31 制御信号（DSTR/SON等） *)
    E001_Out_OUT32_2003_21 : UINT;  (* OUT32 目標位置 下位 [0.01mm] *)
    E001_Out_OUT33_2003_22 : UINT;  (* OUT33 目標位置 上位 [0.01mm] *)
    E001_Out_OUT34_2003_23 : UINT;  (* OUT34 位置決め幅 下位 [0.01mm] *)
    E001_Out_OUT35_2003_24 : UINT;  (* OUT35 位置決め幅 上位 [0.01mm] *)
    E001_Out_OUT36_2003_25 : UINT;  (* OUT36 速度指令 [実機単位] *)
    E001_Out_OUT37_2003_26 : UINT;  (* OUT37 共通加減速 [0.01G] *)
    E001_Out_OUT38_2003_27 : UINT;  (* OUT38 押付け制限 [255=100%] *)
    E001_Out_OUT39_2003_28 : UINT;  (* OUT39 制御信号（DSTR/SON等） *)
    E001_Out_OUT40_2003_29 : UINT;  (* OUT40 目標位置 下位 [0.01mm] *)
    E001_Out_OUT41_2003_2A : UINT;  (* OUT41 目標位置 上位 [0.01mm] *)
    E001_Out_OUT42_2003_2B : UINT;  (* OUT42 位置決め幅 下位 [0.01mm] *)
    E001_Out_OUT43_2003_2C : UINT;  (* OUT43 位置決め幅 上位 [0.01mm] *)
    E001_Out_OUT44_2003_2D : UINT;  (* OUT44 速度指令 [実機単位] *)
    E001_Out_OUT45_2003_2E : UINT;  (* OUT45 共通加減速 [0.01G] *)
    E001_Out_OUT46_2003_2F : UINT;  (* OUT46 押付け制限 [255=100%] *)
    E001_Out_OUT47_2003_30 : UINT;  (* OUT47 制御信号（DSTR/SON等） *)
    E001_Out_OUT48_2003_31 : UINT;  (* OUT48 目標位置 下位 [0.01mm] *)
    E001_Out_OUT49_2003_32 : UINT;  (* OUT49 目標位置 上位 [0.01mm] *)
    E001_Out_OUT50_2003_33 : UINT;  (* OUT50 位置決め幅 下位 [0.01mm] *)
    E001_Out_OUT51_2003_34 : UINT;  (* OUT51 位置決め幅 上位 [0.01mm] *)
    E001_Out_OUT52_2003_35 : UINT;  (* OUT52 速度指令 [実機単位] *)
    E001_Out_OUT53_2003_36 : UINT;  (* OUT53 共通加減速 [0.01G] *)
    E001_Out_OUT54_2003_37 : UINT;  (* OUT54 押付け制限 [255=100%] *)
    E001_Out_OUT55_2003_38 : UINT;  (* OUT55 制御信号（DSTR/SON等） *)
    E005_In_IN00_2004_01_1 : UINT;  (* IN00 GW状態 *)
    E005_In_IN01_2004_02_1 : UINT;  (* IN01 軸リンク状態 *)
    E005_In_IN02_2004_03_1 : UINT;  (* IN02 電源状態0 *)
    E005_In_IN03_2004_04_1 : UINT;  (* IN03 電源状態1 *)
    E005_In_IN04_2004_05_1 : UINT;  (* IN04 電源状態2 *)
    E005_In_IN05_2004_06_1 : UINT;  (* IN05 電源状態3 *)
    E005_In_IN06_2004_07_1 : UINT;  (* IN06 電源状態4（構成依存） *)
    E005_In_IN07_2004_08_1 : UINT;  (* IN07 予約（使用禁止） *)
    E005_In_IN08_2004_09_1 : UINT;  (* #RCON2_1 段バラシ / IN08 現在位置 下位 [0.01mm] *)
    E005_In_IN09_2004_0A_1 : UINT;  (* IN09 現在位置 上位 [0.01mm] *)
    E005_In_IN10_2004_0B_1 : UINT;  (* IN10 指令電流 下位 [mA] *)
    E005_In_IN11_2004_0C_1 : UINT;  (* IN11 指令電流 上位 [mA] *)
    E005_In_IN12_2004_0D_1 : UINT;  (* IN12 現在速度 [実機単位・符号付き] *)
    E005_In_IN13_2004_0E_1 : UINT;  (* IN13 予約（使用禁止） *)
    E005_In_IN14_2004_0F_1 : UINT;  (* IN14 軸異常コード *)
    E005_In_IN15_2004_10_1 : UINT;  (* IN15 状態信号（PEND/SV等） *)
    E005_In_IN16_2004_11_1 : UINT;  (* #RCON2_2 箱詰めX / IN16 現在位置 下位 [0.01mm] *)
    E005_In_IN17_2004_12_1 : UINT;  (* IN17 現在位置 上位 [0.01mm] *)
    E005_In_IN18_2004_13_1 : UINT;  (* IN18 指令電流 下位 [mA] *)
    E005_In_IN19_2004_14_1 : UINT;  (* IN19 指令電流 上位 [mA] *)
    E005_In_IN20_2004_15_1 : UINT;  (* IN20 現在速度 [実機単位・符号付き] *)
    E005_In_IN21_2004_16_1 : UINT;  (* IN21 予約（使用禁止） *)
    E005_In_IN22_2004_17_1 : UINT;  (* IN22 軸異常コード *)
    E005_In_IN23_2004_18_1 : UINT;  (* IN23 状態信号（PEND/SV等） *)
    E005_In_IN24_2004_19_1 : UINT;  (* #RCON2_3 箱詰めY / IN24 現在位置 下位 [0.01mm] *)
    E005_In_IN25_2004_1A_1 : UINT;  (* IN25 現在位置 上位 [0.01mm] *)
    E005_In_IN26_2004_1B_1 : UINT;  (* IN26 指令電流 下位 [mA] *)
    E005_In_IN27_2004_1C_1 : UINT;  (* IN27 指令電流 上位 [mA] *)
    E005_In_IN28_2004_1D_1 : UINT;  (* IN28 現在速度 [実機単位・符号付き] *)
    E005_In_IN29_2004_1E_1 : UINT;  (* IN29 予約（使用禁止） *)
    E005_In_IN30_2004_1F_1 : UINT;  (* IN30 軸異常コード *)
    E005_In_IN31_2004_20_1 : UINT;  (* IN31 状態信号（PEND/SV等） *)
    E005_In_IN32_2004_21_1 : UINT;  (* #RCON2_4 箱詰めZ / IN32 現在位置 下位 [0.01mm] *)
    E005_In_IN33_2004_22_1 : UINT;  (* IN33 現在位置 上位 [0.01mm] *)
    E005_In_IN34_2004_23_1 : UINT;  (* IN34 指令電流 下位 [mA] *)
    E005_In_IN35_2004_24_1 : UINT;  (* IN35 指令電流 上位 [mA] *)
    E005_In_IN36_2004_25_1 : UINT;  (* IN36 現在速度 [実機単位・符号付き] *)
    E005_In_IN37_2004_26_1 : UINT;  (* IN37 予約（使用禁止） *)
    E005_In_IN38_2004_27_1 : UINT;  (* IN38 軸異常コード *)
    E005_In_IN39_2004_28_1 : UINT;  (* IN39 状態信号（PEND/SV等） *)
    E005_In_IN40_2004_29_1 : UINT;  (* #RCON2_5 コンテナ設置 / IN40 現在位置 下位 [0.01mm] *)
    E005_In_IN41_2004_2A_1 : UINT;  (* IN41 現在位置 上位 [0.01mm] *)
    E005_In_IN42_2004_2B_1 : UINT;  (* IN42 指令電流 下位 [mA] *)
    E005_In_IN43_2004_2C_1 : UINT;  (* IN43 指令電流 上位 [mA] *)
    E005_In_IN44_2004_2D_1 : UINT;  (* IN44 現在速度 [実機単位・符号付き] *)
    E005_In_IN45_2004_2E_1 : UINT;  (* IN45 予約（使用禁止） *)
    E005_In_IN46_2004_2F_1 : UINT;  (* IN46 軸異常コード *)
    E005_In_IN47_2004_30_1 : UINT;  (* IN47 状態信号（PEND/SV等） *)
    E005_In_IN48_2004_31_1 : UINT;  (* IN48 用途未確認（今回未使用） *)
    E005_In_IN49_2004_32_1 : UINT;  (* IN49 用途未確認（今回未使用） *)
    E005_In_IN50_2004_33_1 : UINT;  (* IN50 用途未確認（今回未使用） *)
    E005_In_IN51_2004_34_1 : UINT;  (* IN51 用途未確認（今回未使用） *)
    E005_In_IN52_2004_35_1 : UINT;  (* IN52 用途未確認（今回未使用） *)
    E005_In_IN53_2004_36_1 : UINT;  (* IN53 用途未確認（今回未使用） *)
    E005_In_IN54_2004_37_1 : UINT;  (* IN54 用途未確認（今回未使用） *)
    E005_In_IN55_2004_38_1 : UINT;  (* IN55 用途未確認（今回未使用） *)
    E005_Out_OUT00_2003_01_1 : UINT;  (* OUT00 共通制御（MON/RTE） *)
    E005_Out_OUT08_2003_09_1 : UINT;  (* #RCON2_1 段バラシ / OUT08 目標位置 下位 [0.01mm] *)
    E005_Out_OUT09_2003_0A_1 : UINT;  (* OUT09 目標位置 上位 [0.01mm] *)
    E005_Out_OUT10_2003_0B_1 : UINT;  (* OUT10 位置決め幅 下位 [0.01mm] *)
    E005_Out_OUT11_2003_0C_1 : UINT;  (* OUT11 位置決め幅 上位 [0.01mm] *)
    E005_Out_OUT12_2003_0D_1 : UINT;  (* OUT12 速度指令 [実機単位] *)
    E005_Out_OUT13_2003_0E_1 : UINT;  (* OUT13 共通加減速 [0.01G] *)
    E005_Out_OUT14_2003_0F_1 : UINT;  (* OUT14 押付け制限 [255=100%] *)
    E005_Out_OUT15_2003_10_1 : UINT;  (* OUT15 制御信号（DSTR/SON等） *)
    E005_Out_OUT16_2003_11_1 : UINT;  (* #RCON2_2 箱詰めX / OUT16 目標位置 下位 [0.01mm] *)
    E005_Out_OUT17_2003_12_1 : UINT;  (* OUT17 目標位置 上位 [0.01mm] *)
    E005_Out_OUT18_2003_13_1 : UINT;  (* OUT18 位置決め幅 下位 [0.01mm] *)
    E005_Out_OUT19_2003_14_1 : UINT;  (* OUT19 位置決め幅 上位 [0.01mm] *)
    E005_Out_OUT20_2003_15_1 : UINT;  (* OUT20 速度指令 [実機単位] *)
    E005_Out_OUT21_2003_16_1 : UINT;  (* OUT21 共通加減速 [0.01G] *)
    E005_Out_OUT22_2003_17_1 : UINT;  (* OUT22 押付け制限 [255=100%] *)
    E005_Out_OUT23_2003_18_1 : UINT;  (* OUT23 制御信号（DSTR/SON等） *)
    E005_Out_OUT24_2003_19_1 : UINT;  (* #RCON2_3 箱詰めY / OUT24 目標位置 下位 [0.01mm] *)
    E005_Out_OUT25_2003_1A_1 : UINT;  (* OUT25 目標位置 上位 [0.01mm] *)
    E005_Out_OUT26_2003_1B_1 : UINT;  (* OUT26 位置決め幅 下位 [0.01mm] *)
    E005_Out_OUT27_2003_1C_1 : UINT;  (* OUT27 位置決め幅 上位 [0.01mm] *)
    E005_Out_OUT28_2003_1D_1 : UINT;  (* OUT28 速度指令 [実機単位] *)
    E005_Out_OUT29_2003_1E_1 : UINT;  (* OUT29 共通加減速 [0.01G] *)
    E005_Out_OUT30_2003_1F_1 : UINT;  (* OUT30 押付け制限 [255=100%] *)
    E005_Out_OUT31_2003_20_1 : UINT;  (* OUT31 制御信号（DSTR/SON等） *)
    E005_Out_OUT32_2003_21_1 : UINT;  (* #RCON2_4 箱詰めZ / OUT32 目標位置 下位 [0.01mm] *)
    E005_Out_OUT33_2003_22_1 : UINT;  (* OUT33 目標位置 上位 [0.01mm] *)
    E005_Out_OUT34_2003_23_1 : UINT;  (* OUT34 位置決め幅 下位 [0.01mm] *)
    E005_Out_OUT35_2003_24_1 : UINT;  (* OUT35 位置決め幅 上位 [0.01mm] *)
    E005_Out_OUT36_2003_25_1 : UINT;  (* OUT36 速度指令 [実機単位] *)
    E005_Out_OUT37_2003_26_1 : UINT;  (* OUT37 共通加減速 [0.01G] *)
    E005_Out_OUT38_2003_27_1 : UINT;  (* OUT38 押付け制限 [255=100%] *)
    E005_Out_OUT39_2003_28_1 : UINT;  (* OUT39 制御信号（DSTR/SON等） *)
    E005_Out_OUT40_2003_29_1 : UINT;  (* #RCON2_5 コンテナ設置 / OUT40 目標位置 下位 [0.01mm] *)
    E005_Out_OUT41_2003_2A_1 : UINT;  (* OUT41 目標位置 上位 [0.01mm] *)
    E005_Out_OUT42_2003_2B_1 : UINT;  (* OUT42 位置決め幅 下位 [0.01mm] *)
    E005_Out_OUT43_2003_2C_1 : UINT;  (* OUT43 位置決め幅 上位 [0.01mm] *)
    E005_Out_OUT44_2003_2D_1 : UINT;  (* OUT44 速度指令 [実機単位] *)
    E005_Out_OUT45_2003_2E_1 : UINT;  (* OUT45 共通加減速 [0.01G] *)
    E005_Out_OUT46_2003_2F_1 : UINT;  (* OUT46 押付け制限 [255=100%] *)
    E005_Out_OUT47_2003_30_1 : UINT;  (* OUT47 制御信号（DSTR/SON等） *)
    RCON1_AxisApply : ARRAY[1..6] OF BOOL;  (* 軸別出力更新許可（OFF=前値保持）; [1] 出力更新許可（OFF=前値保持）; [2] 出力更新許可（OFF=前値保持）; [3] 出力更新許可（OFF=前値保持）; [4] 出力更新許可（OFF=前値保持）; [5] 出力更新許可（OFF=前値保持）; [6] 出力更新許可（OFF=前値保持） *)
    RCON1_AxisLinked : ARRAY[1..6] OF BOOL;  (* 軸別リンク状態; [1] リンク状態; [2] リンク状態; [3] リンク状態; [4] リンク状態; [5] リンク状態; [6] リンク状態 *)
    RCON1_AxisWritten : ARRAY[1..6] OF BOOL;  (* 軸別出力代入済み（RCON受付とは別）; [1] 出力代入済み（RCON受付とは別）; [2] 出力代入済み（RCON受付とは別）; [3] 出力代入済み（RCON受付とは別）; [4] 出力代入済み（RCON受付とは別）; [5] 出力代入済み（RCON受付とは別）; [6] 出力代入済み（RCON受付とは別） *)
    RCON1_ByteOrderConfirmed : BOOL;  (* ワード・バイト順確認済み（初期OFF） *)
    RCON1_CommOK : BOOL;  (* 通信正常（外部判定・固定ON不可） *)
    RCON1_EncodeError : ARRAY[1..6] OF UINT;  (* 軸別変換エラー番号（0=正常）; [1] 変換エラー番号; [2] 変換エラー番号; [3] 変換エラー番号; [4] 変換エラー番号; [5] 変換エラー番号; [6] 変換エラー番号 *)
    RCON1_EncodeOK : ARRAY[1..6] OF BOOL;  (* 軸別変換正常（運転許可とは別）; [1] 変換正常; [2] 変換正常; [3] 変換正常; [4] 変換正常; [5] 変換正常; [6] 変換正常 *)
    RCON1_GwAlarmCode : UINT;  (* GW異常コード（ALMC/b0～7） *)
    RCON1_GwApply : BOOL;  (* 共通出力更新許可（OFF=前値保持） *)
    RCON1_GwAxisCommError : BOOL;  (* GW－軸 通信異常（ERRT/b13） *)
    RCON1_GwControllerCommLatch : BOOL;  (* GW通信異常保持（LERC/b14） *)
    RCON1_GwHeavyAlarm : BOOL;  (* GW重故障（ALMH/b11） *)
    RCON1_GwLightAlarm : BOOL;  (* GW軽故障（ALML/b10） *)
    RCON1_GwMON_Request : BOOL;  (* MON要求（b15） *)
    RCON1_GwManual : BOOL;  (* 手動モード（MOD/b12） *)
    RCON1_GwRTE_Request : BOOL;  (* 通信異常ラッチ解除要求（b13） *)
    RCON1_GwRun : BOOL;  (* GW動作中（RUN/b15） *)
    RCON1_GwSystemStop : BOOL;  (* システム停止状態（SEMG/b8・監視用） *)
    RCON1_GwWritten : BOOL;  (* 共通出力代入済み（RCON受付とは別） *)
    RCON1_IN : ARRAY[1..6] OF ST_RCON_Direct_IN_Axis;  (* #RCON1 入力値; [1] #A(左側) NG1排出(上下); [2] #B(右側) NG1排出(上下); [3] #A(左側) SF/NG2仕分け(左右); [4] #B(右側) SF/NG2排出(送り); [5] #A(左側) SF/NG2排出(上下); [6] #B(右側) SF/NG2排出(上下); [1].ActualPos_mm 現在位置 [mm]; [1].Current_mA 指令電流 [mA]; [1].ActualSpeed_mm_s 現在速度 [mm/s]; [1].AlarmCode 異常コード; [1].DataValid 入力有効（安全許可とは別）; [1].Status.PositionDone 位置決め完了; [1].Status.HomeDone 原点復帰完了; [1].Status.Moving 移動中; [1].Status.Alarm 軸異常; [1].Status.ServoReady サーボON状態; [1].Status.PushMiss 押付け空振り（未使用）; [1].Status.OverloadWarning 過負荷警告; [1].Status.CommandDone 指令完了（空振り含む）; [1].Status.Zone1 ゾーン1内; [1].Status.Zone2 ゾーン2内; [1].Status.ControllerReady 準備完了; [1].Status.EmergencyStop 非常停止状態（監視）; [2].ActualPos_mm 現在位置 [mm]; [2].Current_mA 指令電流 [mA]; [2].ActualSpeed_mm_s 現在速度 [mm/s]; [2].AlarmCode 異常コード; [2].DataValid 入力有効（安全許可とは別）; [2].Status.PositionDone 位置決め完了; [2].Status.HomeDone 原点復帰完了; [2].Status.Moving 移動中; [2].Status.Alarm 軸異常; [2].Status.ServoReady サーボON状態; [2].Status.PushMiss 押付け空振り（未使用）; [2].Status.OverloadWarning 過負荷警告; [2].Status.CommandDone 指令完了（空振り含む）; [2].Status.Zone1 ゾーン1内; [2].Status.Zone2 ゾーン2内; [2].Status.ControllerReady 準備完了; [2].Status.EmergencyStop 非常停止状態（監視）; [3].ActualPos_mm 現在位置 [mm]; [3].Current_mA 指令電流 [mA]; [3].ActualSpeed_mm_s 現在速度 [mm/s]; [3].AlarmCode 異常コード; [3].DataValid 入力有効（安全許可とは別）; [3].Status.PositionDone 位置決め完了; [3].Status.HomeDone 原点復帰完了; [3].Status.Moving 移動中; [3].Status.Alarm 軸異常; [3].Status.ServoReady サーボON状態; [3].Status.PushMiss 押付け空振り（未使用）; [3].Status.OverloadWarning 過負荷警告; [3].Status.CommandDone 指令完了（空振り含む）; [3].Status.Zone1 ゾーン1内; [3].Status.Zone2 ゾーン2内; [3].Status.ControllerReady 準備完了; [3].Status.EmergencyStop 非常停止状態（監視）; [4].ActualPos_mm 現在位置 [mm]; [4].Current_mA 指令電流 [mA]; [4].ActualSpeed_mm_s 現在速度 [mm/s]; [4].AlarmCode 異常コード; [4].DataValid 入力有効（安全許可とは別）; [4].Status.PositionDone 位置決め完了; [4].Status.HomeDone 原点復帰完了; [4].Status.Moving 移動中; [4].Status.Alarm 軸異常; [4].Status.ServoReady サーボON状態; [4].Status.PushMiss 押付け空振り（未使用）; [4].Status.OverloadWarning 過負荷警告; [4].Status.CommandDone 指令完了（空振り含む）; [4].Status.Zone1 ゾーン1内; [4].Status.Zone2 ゾーン2内; [4].Status.ControllerReady 準備完了; [4].Status.EmergencyStop 非常停止状態（監視）; [5].ActualPos_mm 現在位置 [mm]; [5].Current_mA 指令電流 [mA]; [5].ActualSpeed_mm_s 現在速度 [mm/s]; [5].AlarmCode 異常コード; [5].DataValid 入力有効（安全許可とは別）; [5].Status.PositionDone 位置決め完了; [5].Status.HomeDone 原点復帰完了; [5].Status.Moving 移動中; [5].Status.Alarm 軸異常; [5].Status.ServoReady サーボON状態; [5].Status.PushMiss 押付け空振り（未使用）; [5].Status.OverloadWarning 過負荷警告; [5].Status.CommandDone 指令完了（空振り含む）; [5].Status.Zone1 ゾーン1内; [5].Status.Zone2 ゾーン2内; [5].Status.ControllerReady 準備完了; [5].Status.EmergencyStop 非常停止状態（監視）; [6].ActualPos_mm 現在位置 [mm]; [6].Current_mA 指令電流 [mA]; [6].ActualSpeed_mm_s 現在速度 [mm/s]; [6].AlarmCode 異常コード; [6].DataValid 入力有効（安全許可とは別）; [6].Status.PositionDone 位置決め完了; [6].Status.HomeDone 原点復帰完了; [6].Status.Moving 移動中; [6].Status.Alarm 軸異常; [6].Status.ServoReady サーボON状態; [6].Status.PushMiss 押付け空振り（未使用）; [6].Status.OverloadWarning 過負荷警告; [6].Status.CommandDone 指令完了（空振り含む）; [6].Status.Zone1 ゾーン1内; [6].Status.Zone2 ゾーン2内; [6].Status.ControllerReady 準備完了; [6].Status.EmergencyStop 非常停止状態（監視） *)
    RCON1_LayoutConfirmed : BOOL;  (* I/O配置確認済み（初期OFF） *)
    RCON1_MotionPermit : ARRAY[1..6] OF BOOL;  (* 軸別運転許可（外部判定・初期OFF）; [1] 運転許可（外部判定）; [2] 運転許可（外部判定）; [3] 運転許可（外部判定）; [4] 運転許可（外部判定）; [5] 運転許可（外部判定）; [6] 運転許可（外部判定） *)
    RCON1_OUT : ARRAY[1..6] OF ST_RCON_Direct_OUT_Axis;  (* #RCON1 出力値; [2] #B(右側) NG1排出(上下); [3] #A(左側) SF/NG2仕分け(左右); [4] #B(右側) SF/NG2排出(送り); [5] #A(左側) SF/NG2排出(上下); [6] #B(右側) SF/NG2排出(上下); [1].Control.Pause 一時停止（安全停止とは別）（未接続）; [1] #A(左側) NG1排出(上下); [1].TargetPos_mm 目標位置 [mm]; [1].PositionBand_mm 位置決め幅 [mm]; [1].Speed_mm_s 指令速度 [mm/s]; [1].AccDec_G 加減速度 [G]; [1].PushLimit_pct 押付け制限 [%]（未使用）; [1].Control.Start 移動開始; [1].Control.Home 原点復帰（未接続）; [1].Control.Reset 異常リセット; [1].Control.ServoOn サーボON; [1].Control.InchingSelect インチング選択（OFF=ジョグ）; [1].Control.JogSpeedSelect ジョグ速度切替（未接続）; [1].Control.JogMinus 原点方向ジョグ（未接続）; [1].Control.JogPlus 反原点方向ジョグ（未接続）; [1].Control.GainSelect0 ゲイン選択0（未使用）; [1].Control.GainSelect1 ゲイン選択1（未使用）; [1].Control.PushEnable 押付け選択（OFF=位置決め）（未使用）; [1].Control.PushDirection 押付け方向（未使用）; [1].Control.RelativeMove 相対移動（OFF=絶対）（未使用）; [1].Control.BrakeRelease ブレーキ強制解除（落下注意）; [2].TargetPos_mm 目標位置 [mm]; [2].PositionBand_mm 位置決め幅 [mm]; [2].Speed_mm_s 指令速度 [mm/s]; [2].AccDec_G 加減速度 [G]; [2].PushLimit_pct 押付け制限 [%]（未使用）; [2].Control.Start 移動開始; [2].Control.Home 原点復帰（未接続）; [2].Control.Pause 一時停止（安全停止とは別）（未接続）; [2].Control.Reset 異常リセット; [2].Control.ServoOn サーボON; [2].Control.InchingSelect インチング選択（OFF=ジョグ）; [2].Control.JogSpeedSelect ジョグ速度切替（未接続）; [2].Control.JogMinus 原点方向ジョグ（未接続）; [2].Control.JogPlus 反原点方向ジョグ（未接続）; [2].Control.GainSelect0 ゲイン選択0（未使用）; [2].Control.GainSelect1 ゲイン選択1（未使用）; [2].Control.PushEnable 押付け選択（OFF=位置決め）（未使用）; [2].Control.PushDirection 押付け方向（未使用）; [2].Control.RelativeMove 相対移動（OFF=絶対）（未使用）; [2].Control.BrakeRelease ブレーキ強制解除（落下注意）; [3].TargetPos_mm 目標位置 [mm]; [3].PositionBand_mm 位置決め幅 [mm]; [3].Speed_mm_s 指令速度 [mm/s]; [3].AccDec_G 加減速度 [G]; [3].PushLimit_pct 押付け制限 [%]（未使用）; [3].Control.Start 移動開始; [3].Control.Home 原点復帰（未接続）; [3].Control.Pause 一時停止（安全停止とは別）（未接続）; [3].Control.Reset 異常リセット; [3].Control.ServoOn サーボON; [3].Control.InchingSelect インチング選択（OFF=ジョグ）; [3].Control.JogSpeedSelect ジョグ速度切替（未接続）; [3].Control.JogMinus 原点方向ジョグ（未接続）; [3].Control.JogPlus 反原点方向ジョグ（未接続）; [3].Control.GainSelect0 ゲイン選択0（未使用）; [3].Control.GainSelect1 ゲイン選択1（未使用）; [3].Control.PushEnable 押付け選択（OFF=位置決め）（未使用）; [3].Control.PushDirection 押付け方向（未使用）; [3].Control.RelativeMove 相対移動（OFF=絶対）（未使用）; [3].Control.BrakeRelease ブレーキ強制解除（落下注意）; [4].TargetPos_mm 目標位置 [mm]; [4].PositionBand_mm 位置決め幅 [mm]; [4].Speed_mm_s 指令速度 [mm/s]; [4].AccDec_G 加減速度 [G]; [4].PushLimit_pct 押付け制限 [%]（未使用）; [4].Control.Start 移動開始; [4].Control.Home 原点復帰（未接続）; [4].Control.Pause 一時停止（安全停止とは別）（未接続）; [4].Control.Reset 異常リセット; [4].Control.ServoOn サーボON; [4].Control.InchingSelect インチング選択（OFF=ジョグ）; [4].Control.JogSpeedSelect ジョグ速度切替（未接続）; [4].Control.JogMinus 原点方向ジョグ（未接続）; [4].Control.JogPlus 反原点方向ジョグ（未接続）; [4].Control.GainSelect0 ゲイン選択0（未使用）; [4].Control.GainSelect1 ゲイン選択1（未使用）; [4].Control.PushEnable 押付け選択（OFF=位置決め）（未使用）; [4].Control.PushDirection 押付け方向（未使用）; [4].Control.RelativeMove 相対移動（OFF=絶対）（未使用）; [4].Control.BrakeRelease ブレーキ強制解除（落下注意）; [5].TargetPos_mm 目標位置 [mm]; [5].PositionBand_mm 位置決め幅 [mm]; [5].Speed_mm_s 指令速度 [mm/s]; [5].AccDec_G 加減速度 [G]; [5].PushLimit_pct 押付け制限 [%]（未使用）; [5].Control.Start 移動開始; [5].Control.Home 原点復帰（未接続）; [5].Control.Pause 一時停止（安全停止とは別）（未接続）; [5].Control.Reset 異常リセット; [5].Control.ServoOn サーボON; [5].Control.InchingSelect インチング選択（OFF=ジョグ）; [5].Control.JogSpeedSelect ジョグ速度切替（未接続）; [5].Control.JogMinus 原点方向ジョグ（未接続）; [5].Control.JogPlus 反原点方向ジョグ（未接続）; [5].Control.GainSelect0 ゲイン選択0（未使用）; [5].Control.GainSelect1 ゲイン選択1（未使用）; [5].Control.PushEnable 押付け選択（OFF=位置決め）（未使用）; [5].Control.PushDirection 押付け方向（未使用）; [5].Control.RelativeMove 相対移動（OFF=絶対）（未使用）; [5].Control.BrakeRelease ブレーキ強制解除（落下注意）; [6].TargetPos_mm 目標位置 [mm]; [6].PositionBand_mm 位置決め幅 [mm]; [6].Speed_mm_s 指令速度 [mm/s]; [6].AccDec_G 加減速度 [G]; [6].PushLimit_pct 押付け制限 [%]（未使用）; [6].Control.Start 移動開始; [6].Control.Home 原点復帰（未接続）; [6].Control.Pause 一時停止（安全停止とは別）（未接続）; [6].Control.Reset 異常リセット; [6].Control.ServoOn サーボON; [6].Control.InchingSelect インチング選択（OFF=ジョグ）; [6].Control.JogSpeedSelect ジョグ速度切替（未接続）; [6].Control.JogMinus 原点方向ジョグ（未接続）; [6].Control.JogPlus 反原点方向ジョグ（未接続）; [6].Control.GainSelect0 ゲイン選択0（未使用）; [6].Control.GainSelect1 ゲイン選択1（未使用）; [6].Control.PushEnable 押付け選択（OFF=位置決め）（未使用）; [6].Control.PushDirection 押付け方向（未使用）; [6].Control.RelativeMove 相対移動（OFF=絶対）（未使用）; [6].Control.BrakeRelease ブレーキ強制解除（落下注意） *)
    RCON1_PowerStateRaw : ARRAY[0..4] OF WORD;  (* 電源状態ワード（詳細未確認）; [0] IN02 電源状態0（詳細未確認）; [1] IN03 電源状態1（詳細未確認）; [2] IN04 電源状態2（詳細未確認）; [3] IN05 電源状態3（詳細未確認）; [4] IN06 電源状態4（詳細未確認） *)
    RCON1_RxRaw : ARRAY[0..55] OF UINT;  (* 受信値（バイト交換前）; [0] IN00 GW状態; [1] IN01 軸リンク状態; [2] IN02 電源状態0; [3] IN03 電源状態1; [4] IN04 電源状態2; [5] IN05 電源状態3; [6] IN06 電源状態4（構成依存）; [7] IN07 予約（使用禁止）; [8] IN08 A(左側) RCON1_1 NG1上下降 現在位置 下位 [0.01mm]; [9] IN09 A(左側) RCON1_1 NG1上下降 現在位置 上位 [0.01mm]; [10] IN10 A(左側) RCON1_1 NG1上下降 指令電流 下位 [mA]; [11] IN11 A(左側) RCON1_1 NG1上下降 指令電流 上位 [mA]; [12] IN12 A(左側) RCON1_1 NG1上下降 現在速度 [実機単位・符号付き]; [13] IN13 A(左側) RCON1_1 NG1上下降 予約（使用禁止）; [14] IN14 A(左側) RCON1_1 NG1上下降 軸異常コード; [15] IN15 A(左側) RCON1_1 NG1上下降 状態信号（PEND/SV等）; [16] IN16 B(右側) RCON1_2 NG1上下降 現在位置 下位 [0.01mm]; [17] IN17 B(右側) RCON1_2 NG1上下降 現在位置 上位 [0.01mm]; [18] IN18 B(右側) RCON1_2 NG1上下降 指令電流 下位 [mA]; [19] IN19 B(右側) RCON1_2 NG1上下降 指令電流 上位 [mA]; [20] IN20 B(右側) RCON1_2 NG1上下降 現在速度 [実機単位・符号付き]; [21] IN21 B(右側) RCON1_2 NG1上下降 予約（使用禁止）; [22] IN22 B(右側) RCON1_2 NG1上下降 軸異常コード; [23] IN23 B(右側) RCON1_2 NG1上下降 状態信号（PEND/SV等）; [24] IN24 A(左側) RCON1_3 SF/NG2仕分け(左右) 現在位置 下位 [0.01mm]; [25] IN25 A(左側) RCON1_3 SF/NG2仕分け(左右) 現在位置 上位 [0.01mm]; [26] IN26 A(左側) RCON1_3 SF/NG2仕分け(左右) 指令電流 下位 [mA]; [27] IN27 A(左側) RCON1_3 SF/NG2仕分け(左右) 指令電流 上位 [mA]; [28] IN28 A(左側) RCON1_3 SF/NG2仕分け(左右) 現在速度 [実機単位・符号付き]; [29] IN29 A(左側) RCON1_3 SF/NG2仕分け(左右) 予約（使用禁止）; [30] IN30 A(左側) RCON1_3 SF/NG2仕分け(左右) 軸異常コード; [31] IN31 A(左側) RCON1_3 SF/NG2仕分け(左右) 状態信号（PEND/SV等）; [32] IN32 B(右側) RCON1_4 SF/NG2送り 現在位置 下位 [0.01mm]; [33] IN33 B(右側) RCON1_4 SF/NG2送り 現在位置 上位 [0.01mm]; [34] IN34 B(右側) RCON1_4 SF/NG2送り 指令電流 下位 [mA]; [35] IN35 B(右側) RCON1_4 SF/NG2送り 指令電流 上位 [mA]; [36] IN36 B(右側) RCON1_4 SF/NG2送り 現在速度 [実機単位・符号付き]; [37] IN37 B(右側) RCON1_4 SF/NG2送り 予約（使用禁止）; [38] IN38 B(右側) RCON1_4 SF/NG2送り 軸異常コード; [39] IN39 B(右側) RCON1_4 SF/NG2送り 状態信号（PEND/SV等）; [40] IN40 A(左側) RCON1_5 SF/NG2上下降 現在位置 下位 [0.01mm]; [41] IN41 A(左側) RCON1_5 SF/NG2上下降 現在位置 上位 [0.01mm]; [42] IN42 A(左側) RCON1_5 SF/NG2上下降 指令電流 下位 [mA]; [43] IN43 A(左側) RCON1_5 SF/NG2上下降 指令電流 上位 [mA]; [44] IN44 A(左側) RCON1_5 SF/NG2上下降 現在速度 [実機単位・符号付き]; [45] IN45 A(左側) RCON1_5 SF/NG2上下降 予約（使用禁止）; [46] IN46 A(左側) RCON1_5 SF/NG2上下降 軸異常コード; [47] IN47 A(左側) RCON1_5 SF/NG2上下降 状態信号（PEND/SV等）; [48] IN48 B(右側) RCON1_6 SF/NG2上下降 現在位置 下位 [0.01mm]; [49] IN49 B(右側) RCON1_6 SF/NG2上下降 現在位置 上位 [0.01mm]; [50] IN50 B(右側) RCON1_6 SF/NG2上下降 指令電流 下位 [mA]; [51] IN51 B(右側) RCON1_6 SF/NG2上下降 指令電流 上位 [mA]; [52] IN52 B(右側) RCON1_6 SF/NG2上下降 現在速度 [実機単位・符号付き]; [53] IN53 B(右側) RCON1_6 SF/NG2上下降 予約（使用禁止）; [54] IN54 B(右側) RCON1_6 SF/NG2上下降 軸異常コード; [55] IN55 B(右側) RCON1_6 SF/NG2上下降 状態信号（PEND/SV等） *)
    RCON1_RxWord : ARRAY[0..55] OF WORD;  (* 受信ワード（正規化後）; [0] IN00 GW状態; [1] IN01 軸リンク状態; [2] IN02 電源状態0; [3] IN03 電源状態1; [4] IN04 電源状態2; [5] IN05 電源状態3; [6] IN06 電源状態4（構成依存）; [7] IN07 予約（使用禁止）; [8] IN08 A(左側) RCON1_1 NG1上下降 現在位置 下位 [0.01mm]; [9] IN09 A(左側) RCON1_1 NG1上下降 現在位置 上位 [0.01mm]; [10] IN10 A(左側) RCON1_1 NG1上下降 指令電流 下位 [mA]; [11] IN11 A(左側) RCON1_1 NG1上下降 指令電流 上位 [mA]; [12] IN12 A(左側) RCON1_1 NG1上下降 現在速度 [実機単位・符号付き]; [13] IN13 A(左側) RCON1_1 NG1上下降 予約（使用禁止）; [14] IN14 A(左側) RCON1_1 NG1上下降 軸異常コード; [15] IN15 A(左側) RCON1_1 NG1上下降 状態信号（PEND/SV等）; [16] IN16 B(右側) RCON1_2 NG1上下降 現在位置 下位 [0.01mm]; [17] IN17 B(右側) RCON1_2 NG1上下降 現在位置 上位 [0.01mm]; [18] IN18 B(右側) RCON1_2 NG1上下降 指令電流 下位 [mA]; [19] IN19 B(右側) RCON1_2 NG1上下降 指令電流 上位 [mA]; [20] IN20 B(右側) RCON1_2 NG1上下降 現在速度 [実機単位・符号付き]; [21] IN21 B(右側) RCON1_2 NG1上下降 予約（使用禁止）; [22] IN22 B(右側) RCON1_2 NG1上下降 軸異常コード; [23] IN23 B(右側) RCON1_2 NG1上下降 状態信号（PEND/SV等）; [24] IN24 A(左側) RCON1_3 SF/NG2仕分け(左右) 現在位置 下位 [0.01mm]; [25] IN25 A(左側) RCON1_3 SF/NG2仕分け(左右) 現在位置 上位 [0.01mm]; [26] IN26 A(左側) RCON1_3 SF/NG2仕分け(左右) 指令電流 下位 [mA]; [27] IN27 A(左側) RCON1_3 SF/NG2仕分け(左右) 指令電流 上位 [mA]; [28] IN28 A(左側) RCON1_3 SF/NG2仕分け(左右) 現在速度 [実機単位・符号付き]; [29] IN29 A(左側) RCON1_3 SF/NG2仕分け(左右) 予約（使用禁止）; [30] IN30 A(左側) RCON1_3 SF/NG2仕分け(左右) 軸異常コード; [31] IN31 A(左側) RCON1_3 SF/NG2仕分け(左右) 状態信号（PEND/SV等）; [32] IN32 B(右側) RCON1_4 SF/NG2送り 現在位置 下位 [0.01mm]; [33] IN33 B(右側) RCON1_4 SF/NG2送り 現在位置 上位 [0.01mm]; [34] IN34 B(右側) RCON1_4 SF/NG2送り 指令電流 下位 [mA]; [35] IN35 B(右側) RCON1_4 SF/NG2送り 指令電流 上位 [mA]; [36] IN36 B(右側) RCON1_4 SF/NG2送り 現在速度 [実機単位・符号付き]; [37] IN37 B(右側) RCON1_4 SF/NG2送り 予約（使用禁止）; [38] IN38 B(右側) RCON1_4 SF/NG2送り 軸異常コード; [39] IN39 B(右側) RCON1_4 SF/NG2送り 状態信号（PEND/SV等）; [40] IN40 A(左側) RCON1_5 SF/NG2上下降 現在位置 下位 [0.01mm]; [41] IN41 A(左側) RCON1_5 SF/NG2上下降 現在位置 上位 [0.01mm]; [42] IN42 A(左側) RCON1_5 SF/NG2上下降 指令電流 下位 [mA]; [43] IN43 A(左側) RCON1_5 SF/NG2上下降 指令電流 上位 [mA]; [44] IN44 A(左側) RCON1_5 SF/NG2上下降 現在速度 [実機単位・符号付き]; [45] IN45 A(左側) RCON1_5 SF/NG2上下降 予約（使用禁止）; [46] IN46 A(左側) RCON1_5 SF/NG2上下降 軸異常コード; [47] IN47 A(左側) RCON1_5 SF/NG2上下降 状態信号（PEND/SV等）; [48] IN48 B(右側) RCON1_6 SF/NG2上下降 現在位置 下位 [0.01mm]; [49] IN49 B(右側) RCON1_6 SF/NG2上下降 現在位置 上位 [0.01mm]; [50] IN50 B(右側) RCON1_6 SF/NG2上下降 指令電流 下位 [mA]; [51] IN51 B(右側) RCON1_6 SF/NG2上下降 指令電流 上位 [mA]; [52] IN52 B(右側) RCON1_6 SF/NG2上下降 現在速度 [実機単位・符号付き]; [53] IN53 B(右側) RCON1_6 SF/NG2上下降 予約（使用禁止）; [54] IN54 B(右側) RCON1_6 SF/NG2上下降 軸異常コード; [55] IN55 B(右側) RCON1_6 SF/NG2上下降 状態信号（PEND/SV等） *)
    RCON1_SpeedUnit_mm_s : LREAL;  (* 速度単位 [mm/s/カウント]（1.0/0.1） *)
    RCON1_SwapBytes : BOOL;  (* 上下バイト交換設定（ON=交換） *)
    RCON1_TxUInt : ARRAY[0..55] OF UINT;  (* 送信UINT候補（実I/Oではない）; [0] OUT00 共通制御（MON/RTE）; [1] OUT01 予約（書込禁止）; [2] OUT02 予約（書込禁止）; [3] OUT03 予約（書込禁止）; [4] OUT04 予約（書込禁止）; [5] OUT05 予約（書込禁止）; [6] OUT06 予約（書込禁止）; [7] OUT07 予約（書込禁止）; [8] OUT08 A(左側) RCON1_1 NG1上下降 目標位置 下位 [0.01mm]; [9] OUT09 A(左側) RCON1_1 NG1上下降 目標位置 上位 [0.01mm]; [10] OUT10 A(左側) RCON1_1 NG1上下降 位置決め幅 下位 [0.01mm]; [11] OUT11 A(左側) RCON1_1 NG1上下降 位置決め幅 上位 [0.01mm]; [12] OUT12 A(左側) RCON1_1 NG1上下降 速度指令 [実機単位]; [13] OUT13 A(左側) RCON1_1 NG1上下降 共通加減速 [0.01G]; [14] OUT14 A(左側) RCON1_1 NG1上下降 押付け制限 [255=100%]; [15] OUT15 A(左側) RCON1_1 NG1上下降 制御信号（DSTR/SON等）; [16] OUT16 B(右側) RCON1_2 NG1上下降 目標位置 下位 [0.01mm]; [17] OUT17 B(右側) RCON1_2 NG1上下降 目標位置 上位 [0.01mm]; [18] OUT18 B(右側) RCON1_2 NG1上下降 位置決め幅 下位 [0.01mm]; [19] OUT19 B(右側) RCON1_2 NG1上下降 位置決め幅 上位 [0.01mm]; [20] OUT20 B(右側) RCON1_2 NG1上下降 速度指令 [実機単位]; [21] OUT21 B(右側) RCON1_2 NG1上下降 共通加減速 [0.01G]; [22] OUT22 B(右側) RCON1_2 NG1上下降 押付け制限 [255=100%]; [23] OUT23 B(右側) RCON1_2 NG1上下降 制御信号（DSTR/SON等）; [24] OUT24 A(左側) RCON1_3 SF/NG2仕分け(左右) 目標位置 下位 [0.01mm]; [25] OUT25 A(左側) RCON1_3 SF/NG2仕分け(左右) 目標位置 上位 [0.01mm]; [26] OUT26 A(左側) RCON1_3 SF/NG2仕分け(左右) 位置決め幅 下位 [0.01mm]; [27] OUT27 A(左側) RCON1_3 SF/NG2仕分け(左右) 位置決め幅 上位 [0.01mm]; [28] OUT28 A(左側) RCON1_3 SF/NG2仕分け(左右) 速度指令 [実機単位]; [29] OUT29 A(左側) RCON1_3 SF/NG2仕分け(左右) 共通加減速 [0.01G]; [30] OUT30 A(左側) RCON1_3 SF/NG2仕分け(左右) 押付け制限 [255=100%]; [31] OUT31 A(左側) RCON1_3 SF/NG2仕分け(左右) 制御信号（DSTR/SON等）; [32] OUT32 B(右側) RCON1_4 SF/NG2送り 目標位置 下位 [0.01mm]; [33] OUT33 B(右側) RCON1_4 SF/NG2送り 目標位置 上位 [0.01mm]; [34] OUT34 B(右側) RCON1_4 SF/NG2送り 位置決め幅 下位 [0.01mm]; [35] OUT35 B(右側) RCON1_4 SF/NG2送り 位置決め幅 上位 [0.01mm]; [36] OUT36 B(右側) RCON1_4 SF/NG2送り 速度指令 [実機単位]; [37] OUT37 B(右側) RCON1_4 SF/NG2送り 共通加減速 [0.01G]; [38] OUT38 B(右側) RCON1_4 SF/NG2送り 押付け制限 [255=100%]; [39] OUT39 B(右側) RCON1_4 SF/NG2送り 制御信号（DSTR/SON等）; [40] OUT40 A(左側) RCON1_5 SF/NG2上下降 目標位置 下位 [0.01mm]; [41] OUT41 A(左側) RCON1_5 SF/NG2上下降 目標位置 上位 [0.01mm]; [42] OUT42 A(左側) RCON1_5 SF/NG2上下降 位置決め幅 下位 [0.01mm]; [43] OUT43 A(左側) RCON1_5 SF/NG2上下降 位置決め幅 上位 [0.01mm]; [44] OUT44 A(左側) RCON1_5 SF/NG2上下降 速度指令 [実機単位]; [45] OUT45 A(左側) RCON1_5 SF/NG2上下降 共通加減速 [0.01G]; [46] OUT46 A(左側) RCON1_5 SF/NG2上下降 押付け制限 [255=100%]; [47] OUT47 A(左側) RCON1_5 SF/NG2上下降 制御信号（DSTR/SON等）; [48] OUT48 B(右側) RCON1_6 SF/NG2上下降 目標位置 下位 [0.01mm]; [49] OUT49 B(右側) RCON1_6 SF/NG2上下降 目標位置 上位 [0.01mm]; [50] OUT50 B(右側) RCON1_6 SF/NG2上下降 位置決め幅 下位 [0.01mm]; [51] OUT51 B(右側) RCON1_6 SF/NG2上下降 位置決め幅 上位 [0.01mm]; [52] OUT52 B(右側) RCON1_6 SF/NG2上下降 速度指令 [実機単位]; [53] OUT53 B(右側) RCON1_6 SF/NG2上下降 共通加減速 [0.01G]; [54] OUT54 B(右側) RCON1_6 SF/NG2上下降 押付け制限 [255=100%]; [55] OUT55 B(右側) RCON1_6 SF/NG2上下降 制御信号（DSTR/SON等） *)
    RCON1_TxWord : ARRAY[0..55] OF WORD;  (* 送信ワード候補; [0] OUT00 共通制御（MON/RTE）; [1] OUT01 予約（書込禁止）; [2] OUT02 予約（書込禁止）; [3] OUT03 予約（書込禁止）; [4] OUT04 予約（書込禁止）; [5] OUT05 予約（書込禁止）; [6] OUT06 予約（書込禁止）; [7] OUT07 予約（書込禁止）; [8] OUT08 A(左側) RCON1_1 NG1上下降 目標位置 下位 [0.01mm]; [9] OUT09 A(左側) RCON1_1 NG1上下降 目標位置 上位 [0.01mm]; [10] OUT10 A(左側) RCON1_1 NG1上下降 位置決め幅 下位 [0.01mm]; [11] OUT11 A(左側) RCON1_1 NG1上下降 位置決め幅 上位 [0.01mm]; [12] OUT12 A(左側) RCON1_1 NG1上下降 速度指令 [実機単位]; [13] OUT13 A(左側) RCON1_1 NG1上下降 共通加減速 [0.01G]; [14] OUT14 A(左側) RCON1_1 NG1上下降 押付け制限 [255=100%]; [15] OUT15 A(左側) RCON1_1 NG1上下降 制御信号（DSTR/SON等）; [16] OUT16 B(右側) RCON1_2 NG1上下降 目標位置 下位 [0.01mm]; [17] OUT17 B(右側) RCON1_2 NG1上下降 目標位置 上位 [0.01mm]; [18] OUT18 B(右側) RCON1_2 NG1上下降 位置決め幅 下位 [0.01mm]; [19] OUT19 B(右側) RCON1_2 NG1上下降 位置決め幅 上位 [0.01mm]; [20] OUT20 B(右側) RCON1_2 NG1上下降 速度指令 [実機単位]; [21] OUT21 B(右側) RCON1_2 NG1上下降 共通加減速 [0.01G]; [22] OUT22 B(右側) RCON1_2 NG1上下降 押付け制限 [255=100%]; [23] OUT23 B(右側) RCON1_2 NG1上下降 制御信号（DSTR/SON等）; [24] OUT24 A(左側) RCON1_3 SF/NG2仕分け(左右) 目標位置 下位 [0.01mm]; [25] OUT25 A(左側) RCON1_3 SF/NG2仕分け(左右) 目標位置 上位 [0.01mm]; [26] OUT26 A(左側) RCON1_3 SF/NG2仕分け(左右) 位置決め幅 下位 [0.01mm]; [27] OUT27 A(左側) RCON1_3 SF/NG2仕分け(左右) 位置決め幅 上位 [0.01mm]; [28] OUT28 A(左側) RCON1_3 SF/NG2仕分け(左右) 速度指令 [実機単位]; [29] OUT29 A(左側) RCON1_3 SF/NG2仕分け(左右) 共通加減速 [0.01G]; [30] OUT30 A(左側) RCON1_3 SF/NG2仕分け(左右) 押付け制限 [255=100%]; [31] OUT31 A(左側) RCON1_3 SF/NG2仕分け(左右) 制御信号（DSTR/SON等）; [32] OUT32 B(右側) RCON1_4 SF/NG2送り 目標位置 下位 [0.01mm]; [33] OUT33 B(右側) RCON1_4 SF/NG2送り 目標位置 上位 [0.01mm]; [34] OUT34 B(右側) RCON1_4 SF/NG2送り 位置決め幅 下位 [0.01mm]; [35] OUT35 B(右側) RCON1_4 SF/NG2送り 位置決め幅 上位 [0.01mm]; [36] OUT36 B(右側) RCON1_4 SF/NG2送り 速度指令 [実機単位]; [37] OUT37 B(右側) RCON1_4 SF/NG2送り 共通加減速 [0.01G]; [38] OUT38 B(右側) RCON1_4 SF/NG2送り 押付け制限 [255=100%]; [39] OUT39 B(右側) RCON1_4 SF/NG2送り 制御信号（DSTR/SON等）; [40] OUT40 A(左側) RCON1_5 SF/NG2上下降 目標位置 下位 [0.01mm]; [41] OUT41 A(左側) RCON1_5 SF/NG2上下降 目標位置 上位 [0.01mm]; [42] OUT42 A(左側) RCON1_5 SF/NG2上下降 位置決め幅 下位 [0.01mm]; [43] OUT43 A(左側) RCON1_5 SF/NG2上下降 位置決め幅 上位 [0.01mm]; [44] OUT44 A(左側) RCON1_5 SF/NG2上下降 速度指令 [実機単位]; [45] OUT45 A(左側) RCON1_5 SF/NG2上下降 共通加減速 [0.01G]; [46] OUT46 A(左側) RCON1_5 SF/NG2上下降 押付け制限 [255=100%]; [47] OUT47 A(左側) RCON1_5 SF/NG2上下降 制御信号（DSTR/SON等）; [48] OUT48 B(右側) RCON1_6 SF/NG2上下降 目標位置 下位 [0.01mm]; [49] OUT49 B(右側) RCON1_6 SF/NG2上下降 目標位置 上位 [0.01mm]; [50] OUT50 B(右側) RCON1_6 SF/NG2上下降 位置決め幅 下位 [0.01mm]; [51] OUT51 B(右側) RCON1_6 SF/NG2上下降 位置決め幅 上位 [0.01mm]; [52] OUT52 B(右側) RCON1_6 SF/NG2上下降 速度指令 [実機単位]; [53] OUT53 B(右側) RCON1_6 SF/NG2上下降 共通加減速 [0.01G]; [54] OUT54 B(右側) RCON1_6 SF/NG2上下降 押付け制限 [255=100%]; [55] OUT55 B(右側) RCON1_6 SF/NG2上下降 制御信号（DSTR/SON等） *)
    RCON1_WriteEnable : BOOL;  (* 実出力書込み許可（OFF=前値保持・停止不可） *)
    RCON2_AxisApply : ARRAY[1..5] OF BOOL;  (* 軸別出力更新許可（OFF=前値保持）; [1] 1軸目（No.0）出力更新許可（OFF=前値保持）; [2] 2軸目（No.1）出力更新許可（OFF=前値保持）; [3] 3軸目（No.2）出力更新許可（OFF=前値保持）; [4] 4軸目（No.3）出力更新許可（OFF=前値保持）; [5] 5軸目（No.4）出力更新許可（OFF=前値保持） *)
    RCON2_AxisLinked : ARRAY[1..5] OF BOOL;  (* 軸別リンク状態; [1] 1軸目（No.0）リンク状態; [2] 2軸目（No.1）リンク状態; [3] 3軸目（No.2）リンク状態; [4] 4軸目（No.3）リンク状態; [5] 5軸目（No.4）リンク状態 *)
    RCON2_AxisWritten : ARRAY[1..5] OF BOOL;  (* 軸別出力代入済み（RCON受付とは別）; [1] 1軸目（No.0）出力代入済み（RCON受付とは別）; [2] 2軸目（No.1）出力代入済み（RCON受付とは別）; [3] 3軸目（No.2）出力代入済み（RCON受付とは別）; [4] 4軸目（No.3）出力代入済み（RCON受付とは別）; [5] 5軸目（No.4）出力代入済み（RCON受付とは別） *)
    RCON2_ByteOrderConfirmed : BOOL;  (* ワード・バイト順確認済み（初期OFF） *)
    RCON2_CommOK : BOOL;  (* 通信正常（外部判定・固定ON不可） *)
    RCON2_EncodeError : ARRAY[1..5] OF UINT;  (* 軸別変換エラー番号（0=正常）; [1] 1軸目（No.0）変換エラー番号; [2] 2軸目（No.1）変換エラー番号; [3] 3軸目（No.2）変換エラー番号; [4] 4軸目（No.3）変換エラー番号; [5] 5軸目（No.4）変換エラー番号 *)
    RCON2_EncodeOK : ARRAY[1..5] OF BOOL;  (* 軸別変換正常（運転許可とは別）; [1] 1軸目（No.0）変換正常; [2] 2軸目（No.1）変換正常; [3] 3軸目（No.2）変換正常; [4] 4軸目（No.3）変換正常; [5] 5軸目（No.4）変換正常 *)
    RCON2_GwAlarmCode : UINT;  (* GW異常コード（ALMC/b0～7） *)
    RCON2_GwApply : BOOL;  (* 共通出力更新許可（OFF=前値保持） *)
    RCON2_GwAxisCommError : BOOL;  (* GW－軸 通信異常（ERRT/b13） *)
    RCON2_GwControllerCommLatch : BOOL;  (* GW通信異常保持（LERC/b14） *)
    RCON2_GwHeavyAlarm : BOOL;  (* GW重故障（ALMH/b11） *)
    RCON2_GwLightAlarm : BOOL;  (* GW軽故障（ALML/b10） *)
    RCON2_GwMON_Request : BOOL;  (* MON要求（b15） *)
    RCON2_GwManual : BOOL;  (* 手動モード（MOD/b12） *)
    RCON2_GwRTE_Request : BOOL;  (* 通信異常ラッチ解除要求（b13） *)
    RCON2_GwRun : BOOL;  (* GW動作中（RUN/b15） *)
    RCON2_GwSystemStop : BOOL;  (* システム停止状態（SEMG/b8・監視用） *)
    RCON2_GwWritten : BOOL;  (* 共通出力代入済み（RCON受付とは別） *)
    RCON2_IN : ARRAY[1..5] OF ST_RCON_Direct_IN_Axis;  (* #RCON2 入力値; [1] #RCON2_1 段バラシ; [2] #RCON2_2 箱詰めX; [3] #RCON2_3 箱詰めY; [4] #RCON2_4 箱詰めZ; [5] #RCON2_5 コンテナ設置 *)
    RCON2_LayoutConfirmed : BOOL;  (* I/O配置確認済み（初期OFF） *)
    RCON2_MotionPermit : ARRAY[1..5] OF BOOL;  (* 軸別運転許可（外部判定・初期OFF）; [1] 1軸目（No.0）運転許可（外部判定）; [2] 2軸目（No.1）運転許可（外部判定）; [3] 3軸目（No.2）運転許可（外部判定）; [4] 4軸目（No.3）運転許可（外部判定）; [5] 5軸目（No.4）運転許可（外部判定） *)
    RCON2_OUT : ARRAY[1..5] OF ST_RCON_Direct_OUT_Axis;  (* #RCON2 出力値; [1] #RCON2_1 段バラシ; [2] #RCON2_2 箱詰めX; [3] #RCON2_3 箱詰めY; [4] #RCON2_4 箱詰めZ; [5] #RCON2_5 コンテナ設置 *)
    RCON2_PowerStateRaw : ARRAY[0..4] OF WORD;  (* 電源状態ワード（詳細未確認）; [0] IN02 電源状態0（詳細未確認）; [1] IN03 電源状態1（詳細未確認）; [2] IN04 電源状態2（詳細未確認）; [3] IN05 電源状態3（詳細未確認）; [4] IN06 電源状態4（詳細未確認） *)
    RCON2_RxRaw : ARRAY[0..55] OF UINT;  (* 受信値（バイト交換前）; [0] IN00 GW状態; [1] IN01 軸リンク状態; [2] IN02 電源状態0; [3] IN03 電源状態1; [4] IN04 電源状態2; [5] IN05 電源状態3; [6] IN06 電源状態4（構成依存）; [7] IN07 予約（使用禁止）; [8] IN08 1軸目 現在位置 下位 [0.01mm]; [9] IN09 1軸目 現在位置 上位 [0.01mm]; [10] IN10 1軸目 指令電流 下位 [mA]; [11] IN11 1軸目 指令電流 上位 [mA]; [12] IN12 1軸目 現在速度 [実機単位・符号付き]; [13] IN13 1軸目 予約（使用禁止）; [14] IN14 1軸目 軸異常コード; [15] IN15 1軸目 状態信号（PEND/SV等）; [16] IN16 2軸目 現在位置 下位 [0.01mm]; [17] IN17 2軸目 現在位置 上位 [0.01mm]; [18] IN18 2軸目 指令電流 下位 [mA]; [19] IN19 2軸目 指令電流 上位 [mA]; [20] IN20 2軸目 現在速度 [実機単位・符号付き]; [21] IN21 2軸目 予約（使用禁止）; [22] IN22 2軸目 軸異常コード; [23] IN23 2軸目 状態信号（PEND/SV等）; [24] IN24 3軸目 現在位置 下位 [0.01mm]; [25] IN25 3軸目 現在位置 上位 [0.01mm]; [26] IN26 3軸目 指令電流 下位 [mA]; [27] IN27 3軸目 指令電流 上位 [mA]; [28] IN28 3軸目 現在速度 [実機単位・符号付き]; [29] IN29 3軸目 予約（使用禁止）; [30] IN30 3軸目 軸異常コード; [31] IN31 3軸目 状態信号（PEND/SV等）; [32] IN32 4軸目 現在位置 下位 [0.01mm]; [33] IN33 4軸目 現在位置 上位 [0.01mm]; [34] IN34 4軸目 指令電流 下位 [mA]; [35] IN35 4軸目 指令電流 上位 [mA]; [36] IN36 4軸目 現在速度 [実機単位・符号付き]; [37] IN37 4軸目 予約（使用禁止）; [38] IN38 4軸目 軸異常コード; [39] IN39 4軸目 状態信号（PEND/SV等）; [40] IN40 5軸目 現在位置 下位 [0.01mm]; [41] IN41 5軸目 現在位置 上位 [0.01mm]; [42] IN42 5軸目 指令電流 下位 [mA]; [43] IN43 5軸目 指令電流 上位 [mA]; [44] IN44 5軸目 現在速度 [実機単位・符号付き]; [45] IN45 5軸目 予約（使用禁止）; [46] IN46 5軸目 軸異常コード; [47] IN47 5軸目 状態信号（PEND/SV等）; [48] IN48 用途未確認（今回未使用）; [49] IN49 用途未確認（今回未使用）; [50] IN50 用途未確認（今回未使用）; [51] IN51 用途未確認（今回未使用）; [52] IN52 用途未確認（今回未使用）; [53] IN53 用途未確認（今回未使用）; [54] IN54 用途未確認（今回未使用）; [55] IN55 用途未確認（今回未使用） *)
    RCON2_RxWord : ARRAY[0..55] OF WORD;  (* 受信ワード（正規化後）; [0] IN00 GW状態; [1] IN01 軸リンク状態; [2] IN02 電源状態0; [3] IN03 電源状態1; [4] IN04 電源状態2; [5] IN05 電源状態3; [6] IN06 電源状態4（構成依存）; [7] IN07 予約（使用禁止）; [8] IN08 1軸目 現在位置 下位 [0.01mm]; [9] IN09 1軸目 現在位置 上位 [0.01mm]; [10] IN10 1軸目 指令電流 下位 [mA]; [11] IN11 1軸目 指令電流 上位 [mA]; [12] IN12 1軸目 現在速度 [実機単位・符号付き]; [13] IN13 1軸目 予約（使用禁止）; [14] IN14 1軸目 軸異常コード; [15] IN15 1軸目 状態信号（PEND/SV等）; [16] IN16 2軸目 現在位置 下位 [0.01mm]; [17] IN17 2軸目 現在位置 上位 [0.01mm]; [18] IN18 2軸目 指令電流 下位 [mA]; [19] IN19 2軸目 指令電流 上位 [mA]; [20] IN20 2軸目 現在速度 [実機単位・符号付き]; [21] IN21 2軸目 予約（使用禁止）; [22] IN22 2軸目 軸異常コード; [23] IN23 2軸目 状態信号（PEND/SV等）; [24] IN24 3軸目 現在位置 下位 [0.01mm]; [25] IN25 3軸目 現在位置 上位 [0.01mm]; [26] IN26 3軸目 指令電流 下位 [mA]; [27] IN27 3軸目 指令電流 上位 [mA]; [28] IN28 3軸目 現在速度 [実機単位・符号付き]; [29] IN29 3軸目 予約（使用禁止）; [30] IN30 3軸目 軸異常コード; [31] IN31 3軸目 状態信号（PEND/SV等）; [32] IN32 4軸目 現在位置 下位 [0.01mm]; [33] IN33 4軸目 現在位置 上位 [0.01mm]; [34] IN34 4軸目 指令電流 下位 [mA]; [35] IN35 4軸目 指令電流 上位 [mA]; [36] IN36 4軸目 現在速度 [実機単位・符号付き]; [37] IN37 4軸目 予約（使用禁止）; [38] IN38 4軸目 軸異常コード; [39] IN39 4軸目 状態信号（PEND/SV等）; [40] IN40 5軸目 現在位置 下位 [0.01mm]; [41] IN41 5軸目 現在位置 上位 [0.01mm]; [42] IN42 5軸目 指令電流 下位 [mA]; [43] IN43 5軸目 指令電流 上位 [mA]; [44] IN44 5軸目 現在速度 [実機単位・符号付き]; [45] IN45 5軸目 予約（使用禁止）; [46] IN46 5軸目 軸異常コード; [47] IN47 5軸目 状態信号（PEND/SV等）; [48] IN48 用途未確認（今回未使用）; [49] IN49 用途未確認（今回未使用）; [50] IN50 用途未確認（今回未使用）; [51] IN51 用途未確認（今回未使用）; [52] IN52 用途未確認（今回未使用）; [53] IN53 用途未確認（今回未使用）; [54] IN54 用途未確認（今回未使用）; [55] IN55 用途未確認（今回未使用） *)
    RCON2_SpeedUnit_mm_s : LREAL;  (* 速度単位 [mm/s/カウント]（1.0/0.1） *)
    RCON2_SwapBytes : BOOL;  (* 上下バイト交換設定（ON=交換） *)
    RCON2_TxUInt : ARRAY[0..47] OF UINT;  (* 送信UINT候補（実I/Oではない）; [0] OUT00 共通制御（MON/RTE）; [1] OUT01 予約（書込禁止）; [2] OUT02 予約（書込禁止）; [3] OUT03 予約（書込禁止）; [4] OUT04 予約（書込禁止）; [5] OUT05 予約（書込禁止）; [6] OUT06 予約（書込禁止）; [7] OUT07 予約（書込禁止）; [8] OUT08 1軸目 目標位置 下位 [0.01mm]; [9] OUT09 1軸目 目標位置 上位 [0.01mm]; [10] OUT10 1軸目 位置決め幅 下位 [0.01mm]; [11] OUT11 1軸目 位置決め幅 上位 [0.01mm]; [12] OUT12 1軸目 速度指令 [実機単位]; [13] OUT13 1軸目 共通加減速 [0.01G]; [14] OUT14 1軸目 押付け制限 [255=100%]; [15] OUT15 1軸目 制御信号（DSTR/SON等）; [16] OUT16 2軸目 目標位置 下位 [0.01mm]; [17] OUT17 2軸目 目標位置 上位 [0.01mm]; [18] OUT18 2軸目 位置決め幅 下位 [0.01mm]; [19] OUT19 2軸目 位置決め幅 上位 [0.01mm]; [20] OUT20 2軸目 速度指令 [実機単位]; [21] OUT21 2軸目 共通加減速 [0.01G]; [22] OUT22 2軸目 押付け制限 [255=100%]; [23] OUT23 2軸目 制御信号（DSTR/SON等）; [24] OUT24 3軸目 目標位置 下位 [0.01mm]; [25] OUT25 3軸目 目標位置 上位 [0.01mm]; [26] OUT26 3軸目 位置決め幅 下位 [0.01mm]; [27] OUT27 3軸目 位置決め幅 上位 [0.01mm]; [28] OUT28 3軸目 速度指令 [実機単位]; [29] OUT29 3軸目 共通加減速 [0.01G]; [30] OUT30 3軸目 押付け制限 [255=100%]; [31] OUT31 3軸目 制御信号（DSTR/SON等）; [32] OUT32 4軸目 目標位置 下位 [0.01mm]; [33] OUT33 4軸目 目標位置 上位 [0.01mm]; [34] OUT34 4軸目 位置決め幅 下位 [0.01mm]; [35] OUT35 4軸目 位置決め幅 上位 [0.01mm]; [36] OUT36 4軸目 速度指令 [実機単位]; [37] OUT37 4軸目 共通加減速 [0.01G]; [38] OUT38 4軸目 押付け制限 [255=100%]; [39] OUT39 4軸目 制御信号（DSTR/SON等）; [40] OUT40 5軸目 目標位置 下位 [0.01mm]; [41] OUT41 5軸目 目標位置 上位 [0.01mm]; [42] OUT42 5軸目 位置決め幅 下位 [0.01mm]; [43] OUT43 5軸目 位置決め幅 上位 [0.01mm]; [44] OUT44 5軸目 速度指令 [実機単位]; [45] OUT45 5軸目 共通加減速 [0.01G]; [46] OUT46 5軸目 押付け制限 [255=100%]; [47] OUT47 5軸目 制御信号（DSTR/SON等） *)
    RCON2_TxWord : ARRAY[0..47] OF WORD;  (* 送信ワード候補; [0] OUT00 共通制御（MON/RTE）; [1] OUT01 予約（書込禁止）; [2] OUT02 予約（書込禁止）; [3] OUT03 予約（書込禁止）; [4] OUT04 予約（書込禁止）; [5] OUT05 予約（書込禁止）; [6] OUT06 予約（書込禁止）; [7] OUT07 予約（書込禁止）; [8] OUT08 1軸目 目標位置 下位 [0.01mm]; [9] OUT09 1軸目 目標位置 上位 [0.01mm]; [10] OUT10 1軸目 位置決め幅 下位 [0.01mm]; [11] OUT11 1軸目 位置決め幅 上位 [0.01mm]; [12] OUT12 1軸目 速度指令 [実機単位]; [13] OUT13 1軸目 共通加減速 [0.01G]; [14] OUT14 1軸目 押付け制限 [255=100%]; [15] OUT15 1軸目 制御信号（DSTR/SON等）; [16] OUT16 2軸目 目標位置 下位 [0.01mm]; [17] OUT17 2軸目 目標位置 上位 [0.01mm]; [18] OUT18 2軸目 位置決め幅 下位 [0.01mm]; [19] OUT19 2軸目 位置決め幅 上位 [0.01mm]; [20] OUT20 2軸目 速度指令 [実機単位]; [21] OUT21 2軸目 共通加減速 [0.01G]; [22] OUT22 2軸目 押付け制限 [255=100%]; [23] OUT23 2軸目 制御信号（DSTR/SON等）; [24] OUT24 3軸目 目標位置 下位 [0.01mm]; [25] OUT25 3軸目 目標位置 上位 [0.01mm]; [26] OUT26 3軸目 位置決め幅 下位 [0.01mm]; [27] OUT27 3軸目 位置決め幅 上位 [0.01mm]; [28] OUT28 3軸目 速度指令 [実機単位]; [29] OUT29 3軸目 共通加減速 [0.01G]; [30] OUT30 3軸目 押付け制限 [255=100%]; [31] OUT31 3軸目 制御信号（DSTR/SON等）; [32] OUT32 4軸目 目標位置 下位 [0.01mm]; [33] OUT33 4軸目 目標位置 上位 [0.01mm]; [34] OUT34 4軸目 位置決め幅 下位 [0.01mm]; [35] OUT35 4軸目 位置決め幅 上位 [0.01mm]; [36] OUT36 4軸目 速度指令 [実機単位]; [37] OUT37 4軸目 共通加減速 [0.01G]; [38] OUT38 4軸目 押付け制限 [255=100%]; [39] OUT39 4軸目 制御信号（DSTR/SON等）; [40] OUT40 5軸目 目標位置 下位 [0.01mm]; [41] OUT41 5軸目 目標位置 上位 [0.01mm]; [42] OUT42 5軸目 位置決め幅 下位 [0.01mm]; [43] OUT43 5軸目 位置決め幅 上位 [0.01mm]; [44] OUT44 5軸目 速度指令 [実機単位]; [45] OUT45 5軸目 共通加減速 [0.01G]; [46] OUT46 5軸目 押付け制限 [255=100%]; [47] OUT47 5軸目 制御信号（DSTR/SON等） *)
    RCON2_WriteEnable : BOOL;  (* 実出力書込み許可（OFF=前値保持・停止不可） *)
    RCON1_1_Auto : ARRAY[0..99] OF Bool;  (* 自動移動要求; [1] 原点位置移動; [2] NG仕分け; [3] 動作完了後 原点位置移動 *)
    RCON1_1_OUT_PositionBand_mm : LREAL;  (* 位置決め幅 [mm] *)
    RCON1_1_OUT_TargetPos_mm : LREAL;  (* 目標位置 [mm] *)
    RCON1_1_OUT_Speed_mm_s : LREAL;  (* 指令速度 [mm/s] *)
    RCON1_1_OUT_AccDec_G : LREAL;  (* 加減速度 [G] *)
    RCON1_1_OUT_PushLimit_pct : LREAL;  (* 押付け制限 [%]（未使用） *)
    RCON1_1_ActualPos_mm : LREAL;  (* 現在位置 [mm] *)
    RCON1_1_Current_mA : DINT;  (* 指令電流 [mA]（監視値） *)
    RCON1_1_ActualSpeed_mm_s : LREAL;  (* 現在速度 [mm/s] *)
    RCON1_1_AlarmCode : UINT;  (* 軸異常コード *)
    RCON1_1_DataValid : BOOL;  (* 入力有効（安全許可とは別） *)
    RCON1_1_IN_PositionDone : BOOL;  (* 位置決め完了 *)
    RCON1_1_IN_HomeDone : BOOL;  (* 原点復帰完了 *)
    RCON1_1_IN_Moving : BOOL;  (* 移動中 *)
    RCON1_1_IN_EmergencyStop : BOOL;  (* 非常停止状態（監視） *)
    RCON1_1_IN_ControllerReady : BOOL;  (* 準備完了 *)
    RCON1_1_IN_Zone2 : BOOL;  (* ゾーン2内 *)
    RCON1_1_IN_Zone1 : BOOL;  (* ゾーン1内 *)
    RCON1_1_IN_CommandDone : BOOL;  (* 指令完了 *)
    RCON1_1_IN_OverloadWarning : BOOL;  (* 過負荷警告 *)
    RCON1_1_IN_PushMiss : BOOL;  (* 押付け空振り（未使用） *)
    RCON1_1_IN_ServoReady : BOOL;  (* サーボON状態 *)
    RCON1_1_IN_Alarm : BOOL;  (* 軸異常 *)
    RCON1_1_Ready : BOOL;  (* 動作準備（安全許可とは別） *)
    Error_M : ARRAY[0..99] OF Bool;  (* [3] 未使用：Error_ST1_A_M[0]へ移行; [9] 未使用：Error_ST5_A_M[0]へ移行; [10] 未使用：Error_ST1_B_M[0]へ移行; [11] 未使用：Error_ST5_B_M[0]へ移行; [12] 未使用：Error_ST6_A_M[0]へ移行 *)
    In_Sw_RESET : BOOL;
    RCON1_1_M : ARRAY[0..99] OF BOOL;  (* #A(左側) RCON1_1 NG1排出(上下); [1] 開始指令保持; [2] 予備 *)
    RCON1_1_MoveDone : BOOL;  (* 動作完了 *)
    TimerQ_In_SenCY_NG1_Pick_A_H : BOOL;
    Homing_Para_Stm : _sHOMING_REF;
END_VAR
VAR_EXTERNAL CONSTANT
    Stm_A_Rev_Axis000 : _sAXIS_REF;
END_VAR
VAR_EXTERNAL
    Stm_A_Rev_Axis000_OriginDone : BOOL;  (* A(左側) ST4 反転1 モータ原点復帰完了 *)
    Auto_A_Start : BOOL;
    HMI_Home_SW : BOOL;  (* HMI 原点復帰SW *)
    Stm_A_Rev_Axis000_Origin : BOOL;  (* A(左側) ST4 反転1 モータ原点復帰開始 *)
    Stm_A_Rev_Axis000_MovePos_Degree : LREAL;  (* A(左側)ステッピングモータ000 回転角度 *)
    Stm_A_Rev_Axis000_MoveAbsoluteDone : BOOL;  (* A(左側)ステッピング反転モータ1 絶対値位置決め 動作完了 *)
    Stm_A_Rev_Axis000_Auto : ARRAY[0..99] OF Bool;
    FH_A_ST5_Auto : BOOL;  (* A(左側) ST5 FH自動測定 *)
    FH_A_ST5_Manual : BOOL;  (* A(左側) ST5 FH手動測定 *)
    FH_A_ST5_Done : BOOL;  (* A(左側) ST5 画像検査完了 *)
    FH_Line1_Busy_1 : BOOL;  (* A(左側) 入力：ST5 処理実行中 *)
    FH_Line1_Command_Code_1 : DWORD;
    FH_Line1_Command_Completion_1 : BOOL;  (* A(左側) 入力：ST5 コマンド実行完了 *)
    FH_Line1_Command_Request_1 : BOOL;  (* A(左側) 出力：ST5 コマンド実行 *)
    FH_Line1_DINT_Result_Data_0_1 : DINT;  (* A(左側) 入力：ST5 判定0結果 *)
    FH_Line1_DINT_Result_Data_1_1 : DINT;  (* A(左側) 入力：ST5 判定1結果 *)
    FH_Line1_Error_Status_1 : BOOL;  (* A(左側) 入力：ST5 エラー信号 *)
    FH_Line1_Result_Notification_1 : BOOL;  (* A(左側) 入力：ST51 出力完了 *)
    FH_Line1_Trigger_1 : BOOL;  (* A(左側) 出力：ST5 測定トリガ *)
    FH_Line1_Trigger_Ready_1 : BOOL;  (* A(左側) 入力：ST5 測定準備完了 *)
    Homing_Para_Stm_Rev2 : _sHOMING_REF;  (* A(左側) ST6 反転2原点設定 *)
END_VAR
VAR_EXTERNAL CONSTANT
    Stm_A_Rev_Axis001 : _sAXIS_REF;
END_VAR
VAR_EXTERNAL
    Stm_A_Rev_Axis001_Auto : ARRAY[0..99] OF Bool;  (* A(左側) ST6 反転2自動指令; [1] A(左側) ST6 原点位置移動開始 *)
    Stm_A_Rev_Axis001_MoveAbsoluteDone : BOOL;  (* A(左側) ST6 反転2位置決め完了 *)
    Stm_A_Rev_Axis001_MovePos_Degree : LREAL;  (* A(左側) ST6 反転2指令角度 *)
    Stm_A_Rev_Axis001_Origin : BOOL;  (* A(左側) ST6 反転2 モータ原点復帰開始 *)
    Stm_A_Rev_Axis001_OriginDone : BOOL;  (* A(左側) ST6 反転2 モータ原点復帰完了 *)
    RCON1_2_IN_PositionDone : BOOL;  (* 位置決め完了 *)
    RCON1_2_IN_HomeDone : BOOL;  (* 原点復帰完了 *)
    RCON1_2_IN_Moving : BOOL;  (* 移動中 *)
    RCON1_2_IN_EmergencyStop : BOOL;  (* 非常停止状態（監視） *)
    RCON1_2_IN_ControllerReady : BOOL;  (* 準備完了 *)
    RCON1_2_IN_Zone2 : BOOL;  (* ゾーン2内 *)
    RCON1_2_IN_Zone1 : BOOL;  (* ゾーン1内 *)
    RCON1_2_IN_CommandDone : BOOL;  (* 指令完了 *)
    RCON1_2_IN_OverloadWarning : BOOL;  (* 過負荷警告 *)
    RCON1_2_IN_PushMiss : BOOL;  (* 押付け空振り（未使用） *)
    RCON1_2_IN_ServoReady : BOOL;  (* サーボON状態 *)
    RCON1_2_IN_Alarm : BOOL;  (* 軸異常 *)
    RCON1_2_Ready : BOOL;  (* 動作準備（安全許可とは別） *)
    RCON1_2_Error : BOOL;  (* 異常予備（未接続） *)
    RCON1_2_Error_Clear : BOOL;  (* 解除予備（未接続） *)
    RCON1_2_M : ARRAY[0..99] OF BOOL;  (* #B(右側) RCON1_2 NG1排出(上下); [1] 開始指令保持; [2] 予備 *)
    RCON1_2_MoveDone : BOOL;  (* 動作完了 *)
    RCON1_2_OUT_TargetPos_mm : LREAL;  (* 目標位置 [mm] *)
    RCON1_2_OUT_PositionBand_mm : LREAL;  (* 位置決め幅 [mm] *)
    RCON1_2_OUT_Speed_mm_s : LREAL;  (* 指令速度 [mm/s] *)
    RCON1_2_OUT_AccDec_G : LREAL;  (* 加減速度 [G] *)
    RCON1_2_OUT_PushLimit_pct : LREAL;  (* 押付け制限 [%]（未使用） *)
    RCON1_2_ActualPos_mm : LREAL;  (* 現在位置 [mm] *)
    RCON1_2_Current_mA : DINT;  (* 指令電流 [mA]（監視値） *)
    RCON1_2_ActualSpeed_mm_s : LREAL;  (* 現在速度 [mm/s] *)
    RCON1_2_AlarmCode : UINT;  (* 軸異常コード *)
    RCON1_2_DataValid : BOOL;  (* 入力有効（安全許可とは別） *)
    RCON1_2_Auto : ARRAY[0..99] OF Bool;  (* 自動移動要求; [1] 自動要求1（外部接続用）; [2] 自動要求2（外部接続用）; [3] 自動要求3（外部接続用） *)
    RCON1_3_IN_PositionDone : BOOL;  (* 位置決め完了 *)
    RCON1_3_IN_HomeDone : BOOL;  (* 原点復帰完了 *)
    RCON1_3_IN_Moving : BOOL;  (* 移動中 *)
    RCON1_3_IN_EmergencyStop : BOOL;  (* 非常停止状態（監視） *)
    RCON1_3_IN_ControllerReady : BOOL;  (* 準備完了 *)
    RCON1_3_IN_Zone2 : BOOL;  (* ゾーン2内 *)
    RCON1_3_IN_Zone1 : BOOL;  (* ゾーン1内 *)
    RCON1_3_IN_CommandDone : BOOL;  (* 指令完了 *)
    RCON1_3_IN_OverloadWarning : BOOL;  (* 過負荷警告 *)
    RCON1_3_IN_PushMiss : BOOL;  (* 押付け空振り（未使用） *)
    RCON1_3_IN_ServoReady : BOOL;  (* サーボON状態 *)
    RCON1_3_IN_Alarm : BOOL;  (* 軸異常 *)
    RCON1_3_Ready : BOOL;  (* 動作準備（安全許可とは別） *)
    RCON1_3_Error : BOOL;  (* 異常予備（未接続） *)
    RCON1_3_Error_Clear : BOOL;  (* 解除予備（未接続） *)
    RCON1_3_M : ARRAY[0..99] OF BOOL;  (* #A(左側) RCON1_3 SF/NG2仕分け(左右); [1] 開始指令保持; [2] 予備 *)
    RCON1_3_MoveDone : BOOL;  (* 動作完了 *)
    RCON1_3_OUT_TargetPos_mm : LREAL;  (* 目標位置 [mm] *)
    RCON1_3_OUT_PositionBand_mm : LREAL;  (* 位置決め幅 [mm] *)
    RCON1_3_OUT_Speed_mm_s : LREAL;  (* 指令速度 [mm/s] *)
    RCON1_3_OUT_AccDec_G : LREAL;  (* 加減速度 [G] *)
    RCON1_3_OUT_PushLimit_pct : LREAL;  (* 押付け制限 [%]（未使用） *)
    RCON1_3_ActualPos_mm : LREAL;  (* 現在位置 [mm] *)
    RCON1_3_Current_mA : DINT;  (* 指令電流 [mA]（監視値） *)
    RCON1_3_ActualSpeed_mm_s : LREAL;  (* 現在速度 [mm/s] *)
    RCON1_3_AlarmCode : UINT;  (* 軸異常コード *)
    RCON1_3_DataValid : BOOL;  (* 入力有効（安全許可とは別） *)
    RCON1_3_Auto : ARRAY[0..99] OF Bool;  (* 自動移動要求; [1] 自動要求1（外部接続用）; [2] 自動要求2（外部接続用）; [3] 自動要求3（外部接続用） *)
    RCON1_4_IN_PositionDone : BOOL;  (* 位置決め完了 *)
    RCON1_4_IN_HomeDone : BOOL;  (* 原点復帰完了 *)
    RCON1_4_IN_Moving : BOOL;  (* 移動中 *)
    RCON1_4_IN_EmergencyStop : BOOL;  (* 非常停止状態（監視） *)
    RCON1_4_IN_ControllerReady : BOOL;  (* 準備完了 *)
    RCON1_4_IN_Zone2 : BOOL;  (* ゾーン2内 *)
    RCON1_4_IN_Zone1 : BOOL;  (* ゾーン1内 *)
    RCON1_4_IN_CommandDone : BOOL;  (* 指令完了 *)
    RCON1_4_IN_OverloadWarning : BOOL;  (* 過負荷警告 *)
    RCON1_4_IN_PushMiss : BOOL;  (* 押付け空振り（未使用） *)
    RCON1_4_IN_ServoReady : BOOL;  (* サーボON状態 *)
    RCON1_4_IN_Alarm : BOOL;  (* 軸異常 *)
    RCON1_4_Ready : BOOL;  (* 動作準備（安全許可とは別） *)
    RCON1_4_Error : BOOL;  (* 異常予備（未接続） *)
    RCON1_4_Error_Clear : BOOL;  (* 解除予備（未接続） *)
    RCON1_4_M : ARRAY[0..99] OF BOOL;  (* #B(右側) RCON1_4 SF/NG2排出(送り); [1] 開始指令保持; [2] 予備 *)
    RCON1_4_MoveDone : BOOL;  (* 動作完了 *)
    RCON1_4_OUT_TargetPos_mm : LREAL;  (* 目標位置 [mm] *)
    RCON1_4_OUT_PositionBand_mm : LREAL;  (* 位置決め幅 [mm] *)
    RCON1_4_OUT_Speed_mm_s : LREAL;  (* 指令速度 [mm/s] *)
    RCON1_4_OUT_AccDec_G : LREAL;  (* 加減速度 [G] *)
    RCON1_4_OUT_PushLimit_pct : LREAL;  (* 押付け制限 [%]（未使用） *)
    RCON1_4_ActualPos_mm : LREAL;  (* 現在位置 [mm] *)
    RCON1_4_Current_mA : DINT;  (* 指令電流 [mA]（監視値） *)
    RCON1_4_ActualSpeed_mm_s : LREAL;  (* 現在速度 [mm/s] *)
    RCON1_4_AlarmCode : UINT;  (* 軸異常コード *)
    RCON1_4_DataValid : BOOL;  (* 入力有効（安全許可とは別） *)
    RCON1_4_Auto : ARRAY[0..99] OF Bool;  (* 自動移動要求; [1] 自動要求1（外部接続用）; [2] 自動要求2（外部接続用）; [3] 自動要求3（外部接続用） *)
    RCON1_5_IN_PositionDone : BOOL;  (* 位置決め完了 *)
    RCON1_5_IN_HomeDone : BOOL;  (* 原点復帰完了 *)
    RCON1_5_IN_Moving : BOOL;  (* 移動中 *)
    RCON1_5_IN_EmergencyStop : BOOL;  (* 非常停止状態（監視） *)
    RCON1_5_IN_ControllerReady : BOOL;  (* 準備完了 *)
    RCON1_5_IN_Zone2 : BOOL;  (* ゾーン2内 *)
    RCON1_5_IN_Zone1 : BOOL;  (* ゾーン1内 *)
    RCON1_5_IN_CommandDone : BOOL;  (* 指令完了 *)
    RCON1_5_IN_OverloadWarning : BOOL;  (* 過負荷警告 *)
    RCON1_5_IN_PushMiss : BOOL;  (* 押付け空振り（未使用） *)
    RCON1_5_IN_ServoReady : BOOL;  (* サーボON状態 *)
    RCON1_5_IN_Alarm : BOOL;  (* 軸異常 *)
    RCON1_5_Ready : BOOL;  (* 動作準備（安全許可とは別） *)
    RCON1_5_Error : BOOL;  (* 異常予備（未接続） *)
    RCON1_5_Error_Clear : BOOL;  (* 解除予備（未接続） *)
    RCON1_5_M : ARRAY[0..99] OF BOOL;  (* #A(左側) RCON1_5 SF/NG2排出(上下); [1] 開始指令保持; [2] 予備 *)
    RCON1_5_MoveDone : BOOL;  (* 動作完了 *)
    RCON1_5_OUT_TargetPos_mm : LREAL;  (* 目標位置 [mm] *)
    RCON1_5_OUT_PositionBand_mm : LREAL;  (* 位置決め幅 [mm] *)
    RCON1_5_OUT_Speed_mm_s : LREAL;  (* 指令速度 [mm/s] *)
    RCON1_5_OUT_AccDec_G : LREAL;  (* 加減速度 [G] *)
    RCON1_5_OUT_PushLimit_pct : LREAL;  (* 押付け制限 [%]（未使用） *)
    RCON1_5_ActualPos_mm : LREAL;  (* 現在位置 [mm] *)
    RCON1_5_Current_mA : DINT;  (* 指令電流 [mA]（監視値） *)
    RCON1_5_ActualSpeed_mm_s : LREAL;  (* 現在速度 [mm/s] *)
    RCON1_5_AlarmCode : UINT;  (* 軸異常コード *)
    RCON1_5_DataValid : BOOL;  (* 入力有効（安全許可とは別） *)
    RCON1_5_Auto : ARRAY[0..99] OF Bool;  (* 自動移動要求; [1] 原点位置移動; [2] 自動要求2（外部接続用）; [3] 自動要求3（外部接続用） *)
    RCON1_6_IN_PositionDone : BOOL;  (* 位置決め完了 *)
    RCON1_6_IN_HomeDone : BOOL;  (* 原点復帰完了 *)
    RCON1_6_IN_Moving : BOOL;  (* 移動中 *)
    RCON1_6_IN_EmergencyStop : BOOL;  (* 非常停止状態（監視） *)
    RCON1_6_IN_ControllerReady : BOOL;  (* 準備完了 *)
    RCON1_6_IN_Zone2 : BOOL;  (* ゾーン2内 *)
    RCON1_6_IN_Zone1 : BOOL;  (* ゾーン1内 *)
    RCON1_6_IN_CommandDone : BOOL;  (* 指令完了 *)
    RCON1_6_IN_OverloadWarning : BOOL;  (* 過負荷警告 *)
    RCON1_6_IN_PushMiss : BOOL;  (* 押付け空振り（未使用） *)
    RCON1_6_IN_ServoReady : BOOL;  (* サーボON状態 *)
    RCON1_6_IN_Alarm : BOOL;  (* 軸異常 *)
    RCON1_6_Ready : BOOL;  (* 動作準備（安全許可とは別） *)
    RCON1_6_Error : BOOL;  (* 異常予備（未接続） *)
    RCON1_6_Error_Clear : BOOL;  (* 解除予備（未接続） *)
    RCON1_6_M : ARRAY[0..99] OF BOOL;  (* #B(右側) RCON1_6 SF/NG2排出(上下); [1] 開始指令保持; [2] 予備 *)
    RCON1_6_MoveDone : BOOL;  (* 動作完了 *)
    RCON1_6_OUT_TargetPos_mm : LREAL;  (* 目標位置 [mm] *)
    RCON1_6_OUT_PositionBand_mm : LREAL;  (* 位置決め幅 [mm] *)
    RCON1_6_OUT_Speed_mm_s : LREAL;  (* 指令速度 [mm/s] *)
    RCON1_6_OUT_AccDec_G : LREAL;  (* 加減速度 [G] *)
    RCON1_6_OUT_PushLimit_pct : LREAL;  (* 押付け制限 [%]（未使用） *)
    RCON1_6_ActualPos_mm : LREAL;  (* 現在位置 [mm] *)
    RCON1_6_Current_mA : DINT;  (* 指令電流 [mA]（監視値） *)
    RCON1_6_ActualSpeed_mm_s : LREAL;  (* 現在速度 [mm/s] *)
    RCON1_6_AlarmCode : UINT;  (* 軸異常コード *)
    RCON1_6_DataValid : BOOL;  (* 入力有効（安全許可とは別） *)
    RCON1_6_Auto : ARRAY[0..99] OF Bool;  (* 自動移動要求; [1] 自動要求1（外部接続用）; [2] 自動要求2（外部接続用）; [3] 自動要求3（外部接続用） *)
    TimerQ_In_SenCY_NG1_Pick_B_H : BOOL;  (* 【X428】B(右側) NG1ピックアップ戻 *)
    HMI_Message_Request : ARRAY[0..121] OF BOOL;  (* #HMI メッセージ表示要求; [0] 未使用; [1] 【Y616】A(左側) 供給スライド戻 異常表示; [2] 【Y617】A(左側) 供給スライド行 異常表示; [3] 【Y618】A(左側) 供給ピックアップ戻 異常表示; [4] 【Y619】A(左側) 供給ピックアップ行 異常表示; [5] 【Y620】A(左側) 供給チャック閉 戻 異常表示; [6] 【Y621】A(左側) 供給チャック開 行 異常表示; [7] 【Y622】B(右側) 供給スライド戻 異常表示; [8] 【Y623】B(右側) 供給スライド行 異常表示; [9] 【Y624】B(右側) 供給ピックアップ戻 異常表示; [10] 【Y625】B(右側) 供給ピックアップ行 異常表示; [11] 【Y626】B(右側) 供給チャック閉 戻 異常表示; [12] 【Y627】B(右側) 供給チャック開 行 異常表示; [13] 【Y700】A(左側) 高さ検査押え戻 異常表示; [14] 【Y701】A(左側) 高さ検査押え行 異常表示; [15] 【Y702】A(左側) 高さ検査持上戻 異常表示; [16] 【Y703】A(左側) 高さ検査持上行 異常表示; [17] 【Y704】A(左側) NG1ピックアップ戻 異常表示; [18] 【Y705】A(左側) NG1ピックアップ 行 異常表示; [19] 【Y706】A(左側) NG1チャック戻 異常表示; [20] 【Y707】A(左側) NG1チャック行 異常表示; [21] 【Y708】A(左側)ST4 反転1チャック閉 異常表示; [22] 【Y709】A(左側)ST4 反転1チャック開 異常表示; [23] 【Y710】A(左側)ST4 反転1ピックアップ戻 異常表示; [24] 【Y711】A(左側)ST4 反転1ピックアップ行 異常表示; [25] 【Y712】A(左側)ST6 反転2チャック閉 戻 異常表示; [26] 【Y713】A(左側)ST6 反転2チャック開 行 異常表示; [27] 【Y714】A(左側)ST6 反転2ピックアップ戻 異常表示; [28] 【Y715】A(左側)ST6 反転2ピックアップ行 異常表示; [29] 【Y716】A(左側) 排出チャック閉 戻 異常表示; [30] 【Y717】A(左側) 排出チャック開 行 異常表示; [31] 【Y718】A(左側) 排出フォルダ送り戻 異常表示; [32] 【Y719】A(左側) 排出フォルダ送り行 異常表示; [33] A(左側) 位置1ストッパー戻 異常表示; [34] 【Y720】A(左側) 位置1ストッパー 行 異常表示; [35] 【Y721】A(左側) 位置2ストッパー 異常表示; [36] 【Y721】A(左側) 位置2ストッパー 異常表示; [37] 【Y722】A(左側) 位置3ストッパー戻 異常表示; [38] 【Y722】A(左側) 位置3ストッパー行 異常表示; [39] Output_A_Error_M[33] 異常表示; [40] 【Y723】A(左側) 位置4ストッパー行 異常表示; [41] 【Y724】A(左側) 位置5ストッパー戻 異常表示; [42] 【Y724】A(左側) 位置5ストッパー行 異常表示; [43] 【Y725】A(左側) 位置6ストッパー戻 異常表示; [44] 【Y725】A(左側) 位置6ストッパー行 異常表示; [45] 【Y726】A(左側) ストックフォルダターン戻 異常表示; [46] 【Y727】A(左側) ストックフォルダターン行 異常表示; [47] 【Y728】A(左側) NG1仕分け 戻 異常表示; [48] 【Y729】A(左側) NG1仕分け 行 異常表示; [49] 【Y800】B(右側) 高さ検査押え戻 異常表示; [50] 【Y801】B(右側) 高さ検査押え行 異常表示; [51] 【Y802】B(右側) 高さ検査持上戻 異常表示; [52] 【Y803】B(右側) 高さ検査持上行 異常表示; [53] 【Y804】B(右側) NG1ピックアップ戻 異常表示; [54] 【Y805】B(右側) NG1ピックアップ 行 異常表示; [55] 【Y806】B(右側) NG1チャック戻 異常表示; [56] 【Y807】B(右側) NG1チャック行 異常表示; [57] 【Y808】B(右側)ST4 反転1チャック閉 戻 異常表示; [58] 【Y809】B(右側)ST4 反転1チャック開 戻 異常表示; [59] 【Y810】B(右側)ST4 反転1ピックアップ戻 異常表示; [60] 【Y811】B(右側)ST4 反転1ピックアップ行 異常表示; [61] 【Y812】B(右側)ST6 反転2チャック閉 戻 異常表示; [62] 【Y813】B(右側)ST6 反転2チャック開 行 異常表示; [63] 【Y814】B(右側)ST6 反転2ピックアップ戻 異常表示; [64] 【Y815】B(右側)ST6 反転2ピックアップ行 異常表示; [65] 【Y816】B(右側) 排出チャック閉 戻 異常表示; [66] 【Y817】B(右側) 排出チャック開 行 異常表示; [67] 【Y818】B(右側) 排出フォルダ送り戻 異常表示; [68] 【Y819】B(右側) 排出フォルダ送り行 異常表示; [69] 【Y820】B(右側) 位置1ストッパー 戻 異常表示; [70] 【Y820】B(右側) 位置1ストッパー 行 異常表示; [71] 【Y821】B(右側) 位置2ストッパー戻 異常表示; [72] 【Y821】B(右側) 位置2ストッパー行 異常表示; [73] 【Y822】B(右側) 位置3ストッパー戻 異常表示; [74] 【Y822】B(右側) 位置3ストッパー行 異常表示; [75] 【Y823】B(右側) 位置4ストッパー戻 異常表示; [76] 【Y823】B(右側) 位置4ストッパー行 異常表示; [77] 【Y824】B(右側) 位置5ストッパー戻 異常表示; [78] 【Y824】B(右側) 位置5ストッパー行 異常表示; [79] 【Y825】B(右側) 位置6ストッパー戻 異常表示; [80] 【Y825】B(右側) 位置6ストッパー行 異常表示; [81] 【Y826】B(右側) ストックフォルダターン戻 異常表示; [82] 【Y827】B(右側) ストックフォルダターン行 異常表示; [83] 【Y828】B(右側) NG1仕分け 戻 異常表示; [84] 【Y829】B(右側) NG1仕分け 行 異常表示; [85] 【Y1200】空コンテナ送り 戻 異常表示; [86] 【Y1201】空コンテナ送り 行 異常表示; [87] 【Y1202】段バラシ爪 戻 異常表示; [88] 【Y1203】段バラシ爪 行 異常表示; [89] 【Y1204】コンテナ排出 戻 異常表示; [90] 【Y1205】コンテナ排出 行 異常表示; [91] Output_Share_Error_M[7] 異常表示; [92] 【Y1207】箱入れチャック 行 異常表示; [93] 【Y1208】コンテナ仕分けストッパー 戻 異常表示; [94] 【Y1209】コンテナ仕分けストッパー 行 異常表示; [95] 【Y1210】コンテナ仕分け送り 戻 異常表示; [96] Output_Share_Error_M[12] 異常表示; [97] 【Y1300】A(左側) コンベア受渡送り戻 異常表示; [98] 【Y1301】A(左側) コンベア受渡送り行 異常表示; [99] 【Y1302】B(右側) コンベア受渡送り戻 異常表示; [100] 【Y1303】B(右側) コンベア受渡送り行 異常表示; [101] ST1 搬送ワーク不一致; [102] ST2 搬送ワーク不一致; [103] ST3 搬送ワーク不一致; [104] ST4 搬送ワーク不一致; [105] ST5 搬送ワーク不一致; [106] ST6 搬送ワーク不一致; [107] ST7 搬送ワーク不一致; [108] A(左側) ST1 FH測定時間超過; [109] A(左側) ST1 FH異常; [110] A(左側) ST5 FH異常; [111] B(右側) ST1 FH異常; [112] B(右側) ST5 FH異常; [113] A(左側) ST1 FH判定OK; [114] A(左側) ST1 FH判定NG1; [115] A(左側) ST1 FH判定NG2; [116] A(左側) ST1 検査前ワーク不一致; [117] A(左側) ST5 FH測定時間超過; [118] A(左側) ST5 FH判定OK; [119] A(左側) ST5 FH判定NG1; [120] A(左側) ST5 FH判定NG2; [121] A(左側) ST5 検査前ワーク不一致 *)
    HMI_Error_WorkSample : ARRAY[0..1] OF BOOL;  (* #HMI 再開前のワーク不一致; [0] A(左側) ST1; [1] A(左側) ST5 *)
    Error_ST1_A_Timeout : BOOL;  (* FHタイムアウト（非保持） *)
    Error_ST5_A_Timeout : BOOL;  (* FHタイムアウト（非保持） *)
    FH_Line2_Error_Status_1 : BOOL;
    FH_Line3_Error_Status_1 : BOOL;
    RCON1_1_Error : BOOL;
    RCON1_1_Error_Clear : BOOL;
    Retry : ARRAY[0..99] OF BOOL;
    Stm_A_Rev_Axis000_MoveError : BOOL;  (* 動作エラー *)
    Stm_A_Rev1_Axis000_Power_Error : BOOL;  (* Stm A Axis000 サーボON エラー *)
    Stm_A_Rev_Axis001_MoveError : BOOL;  (* Stm A Axis001 絶対値位置決め エラー *)
    Stm_A_Rev2_Axis001_Power_Error : BOOL;  (* Stm A Axis001 サーボON エラー *)
    RCON2_1_M : ARRAY[0..99] OF BOOL;  (* #RCON2_1 段バラシ; [1] 開始指令保持; [2] 予備 *)
    RCON2_1_IN_PositionDone : BOOL;  (* 位置決め完了 *)
    RCON2_1_IN_HomeDone : BOOL;  (* 原点復帰完了 *)
    RCON2_1_IN_Moving : BOOL;  (* 移動中 *)
    RCON2_1_IN_EmergencyStop : BOOL;  (* 非常停止状態（監視） *)
    RCON2_1_IN_ControllerReady : BOOL;  (* 準備完了 *)
    RCON2_1_IN_Zone2 : BOOL;  (* ゾーン2内 *)
    RCON2_1_IN_Zone1 : BOOL;  (* ゾーン1内 *)
    RCON2_1_IN_CommandDone : BOOL;  (* 指令完了 *)
    RCON2_1_IN_OverloadWarning : BOOL;  (* 過負荷警告 *)
    RCON2_1_IN_PushMiss : BOOL;  (* 押付け空振り（未使用） *)
    RCON2_1_IN_ServoReady : BOOL;  (* サーボON状態 *)
    RCON2_1_IN_Alarm : BOOL;  (* 軸異常 *)
    RCON2_1_Ready : BOOL;  (* 動作準備（安全許可とは別） *)
    RCON2_1_MoveDone : BOOL;  (* 動作完了 *)
    RCON2_1_OUT_TargetPos_mm : LREAL;  (* 目標位置 [mm] *)
    RCON2_1_OUT_PositionBand_mm : LREAL;  (* 位置決め幅 [mm] *)
    RCON2_1_OUT_Speed_mm_s : LREAL;  (* 指令速度 [mm/s] *)
    RCON2_1_OUT_AccDec_G : LREAL;  (* 加減速度 [G] *)
    RCON2_1_OUT_PushLimit_pct : LREAL;  (* 押付け制限 [%]（未使用） *)
    RCON2_1_ActualPos_mm : LREAL;  (* 現在位置 [mm] *)
    RCON2_1_Current_mA : DINT;  (* 指令電流 [mA]（監視値） *)
    RCON2_1_ActualSpeed_mm_s : LREAL;  (* 現在速度 [mm/s] *)
    RCON2_1_AlarmCode : UINT;  (* 軸異常コード *)
    RCON2_1_DataValid : BOOL;  (* 入力有効（安全許可とは別） *)
    RCON2_1_Auto : ARRAY[0..99] OF Bool;  (* 自動移動要求; [1] 自動要求1（未接続）; [2] 自動要求2（未接続）; [3] 自動要求3（未接続） *)
    RCON2_2_M : ARRAY[0..99] OF BOOL;  (* #RCON2_2 箱詰めX; [1] 開始指令保持; [2] 予備 *)
    RCON2_2_IN_PositionDone : BOOL;  (* 位置決め完了 *)
    RCON2_2_IN_HomeDone : BOOL;  (* 原点復帰完了 *)
    RCON2_2_IN_Moving : BOOL;  (* 移動中 *)
    RCON2_2_IN_EmergencyStop : BOOL;  (* 非常停止状態（監視） *)
    RCON2_2_IN_ControllerReady : BOOL;  (* 準備完了 *)
    RCON2_2_IN_Zone2 : BOOL;  (* ゾーン2内 *)
    RCON2_2_IN_Zone1 : BOOL;  (* ゾーン1内 *)
    RCON2_2_IN_CommandDone : BOOL;  (* 指令完了 *)
    RCON2_2_IN_OverloadWarning : BOOL;  (* 過負荷警告 *)
    RCON2_2_IN_PushMiss : BOOL;  (* 押付け空振り（未使用） *)
    RCON2_2_IN_ServoReady : BOOL;  (* サーボON状態 *)
    RCON2_2_IN_Alarm : BOOL;  (* 軸異常 *)
    RCON2_2_Ready : BOOL;  (* 動作準備（安全許可とは別） *)
    RCON2_2_MoveDone : BOOL;  (* 動作完了 *)
    RCON2_2_OUT_TargetPos_mm : LREAL;  (* 目標位置 [mm] *)
    RCON2_2_OUT_PositionBand_mm : LREAL;  (* 位置決め幅 [mm] *)
    RCON2_2_OUT_Speed_mm_s : LREAL;  (* 指令速度 [mm/s] *)
    RCON2_2_OUT_AccDec_G : LREAL;  (* 加減速度 [G] *)
    RCON2_2_OUT_PushLimit_pct : LREAL;  (* 押付け制限 [%]（未使用） *)
    RCON2_2_ActualPos_mm : LREAL;  (* 現在位置 [mm] *)
    RCON2_2_Current_mA : DINT;  (* 指令電流 [mA]（監視値） *)
    RCON2_2_ActualSpeed_mm_s : LREAL;  (* 現在速度 [mm/s] *)
    RCON2_2_AlarmCode : UINT;  (* 軸異常コード *)
    RCON2_2_DataValid : BOOL;  (* 入力有効（安全許可とは別） *)
    RCON2_2_Auto : ARRAY[0..99] OF Bool;  (* 自動移動要求; [1] 自動要求1（未接続）; [2] 自動要求2（未接続）; [3] 自動要求3（未接続） *)
    RCON2_3_M : ARRAY[0..99] OF BOOL;  (* #RCON2_3 箱詰めY; [1] 開始指令保持; [2] 予備 *)
    RCON2_3_IN_PositionDone : BOOL;  (* 位置決め完了 *)
    RCON2_3_IN_HomeDone : BOOL;  (* 原点復帰完了 *)
    RCON2_3_IN_Moving : BOOL;  (* 移動中 *)
    RCON2_3_IN_EmergencyStop : BOOL;  (* 非常停止状態（監視） *)
    RCON2_3_IN_ControllerReady : BOOL;  (* 準備完了 *)
    RCON2_3_IN_Zone2 : BOOL;  (* ゾーン2内 *)
    RCON2_3_IN_Zone1 : BOOL;  (* ゾーン1内 *)
    RCON2_3_IN_CommandDone : BOOL;  (* 指令完了 *)
    RCON2_3_IN_OverloadWarning : BOOL;  (* 過負荷警告 *)
    RCON2_3_IN_PushMiss : BOOL;  (* 押付け空振り（未使用） *)
    RCON2_3_IN_ServoReady : BOOL;  (* サーボON状態 *)
    RCON2_3_IN_Alarm : BOOL;  (* 軸異常 *)
    RCON2_3_Ready : BOOL;  (* 動作準備（安全許可とは別） *)
    RCON2_3_MoveDone : BOOL;  (* 動作完了 *)
    RCON2_3_OUT_TargetPos_mm : LREAL;  (* 目標位置 [mm] *)
    RCON2_3_OUT_PositionBand_mm : LREAL;  (* 位置決め幅 [mm] *)
    RCON2_3_OUT_Speed_mm_s : LREAL;  (* 指令速度 [mm/s] *)
    RCON2_3_OUT_AccDec_G : LREAL;  (* 加減速度 [G] *)
    RCON2_3_OUT_PushLimit_pct : LREAL;  (* 押付け制限 [%]（未使用） *)
    RCON2_3_ActualPos_mm : LREAL;  (* 現在位置 [mm] *)
    RCON2_3_Current_mA : DINT;  (* 指令電流 [mA]（監視値） *)
    RCON2_3_ActualSpeed_mm_s : LREAL;  (* 現在速度 [mm/s] *)
    RCON2_3_AlarmCode : UINT;  (* 軸異常コード *)
    RCON2_3_DataValid : BOOL;  (* 入力有効（安全許可とは別） *)
    RCON2_3_Auto : ARRAY[0..99] OF Bool;  (* 自動移動要求; [1] 自動要求1（未接続）; [2] 自動要求2（未接続）; [3] 自動要求3（未接続） *)
    RCON2_4_M : ARRAY[0..99] OF BOOL;  (* #RCON2_4 箱詰めZ; [1] 開始指令保持; [2] 予備 *)
    RCON2_4_IN_PositionDone : BOOL;  (* 位置決め完了 *)
    RCON2_4_IN_HomeDone : BOOL;  (* 原点復帰完了 *)
    RCON2_4_IN_Moving : BOOL;  (* 移動中 *)
    RCON2_4_IN_EmergencyStop : BOOL;  (* 非常停止状態（監視） *)
    RCON2_4_IN_ControllerReady : BOOL;  (* 準備完了 *)
    RCON2_4_IN_Zone2 : BOOL;  (* ゾーン2内 *)
    RCON2_4_IN_Zone1 : BOOL;  (* ゾーン1内 *)
    RCON2_4_IN_CommandDone : BOOL;  (* 指令完了 *)
    RCON2_4_IN_OverloadWarning : BOOL;  (* 過負荷警告 *)
    RCON2_4_IN_PushMiss : BOOL;  (* 押付け空振り（未使用） *)
    RCON2_4_IN_ServoReady : BOOL;  (* サーボON状態 *)
    RCON2_4_IN_Alarm : BOOL;  (* 軸異常 *)
    RCON2_4_Ready : BOOL;  (* 動作準備（安全許可とは別） *)
    RCON2_4_MoveDone : BOOL;  (* 動作完了 *)
    RCON2_4_OUT_TargetPos_mm : LREAL;  (* 目標位置 [mm] *)
    RCON2_4_OUT_PositionBand_mm : LREAL;  (* 位置決め幅 [mm] *)
    RCON2_4_OUT_Speed_mm_s : LREAL;  (* 指令速度 [mm/s] *)
    RCON2_4_OUT_AccDec_G : LREAL;  (* 加減速度 [G] *)
    RCON2_4_OUT_PushLimit_pct : LREAL;  (* 押付け制限 [%]（未使用） *)
    RCON2_4_ActualPos_mm : LREAL;  (* 現在位置 [mm] *)
    RCON2_4_Current_mA : DINT;  (* 指令電流 [mA]（監視値） *)
    RCON2_4_ActualSpeed_mm_s : LREAL;  (* 現在速度 [mm/s] *)
    RCON2_4_AlarmCode : UINT;  (* 軸異常コード *)
    RCON2_4_DataValid : BOOL;  (* 入力有効（安全許可とは別） *)
    RCON2_4_Auto : ARRAY[0..99] OF Bool;  (* 自動移動要求; [1] 自動要求1（未接続）; [2] 自動要求2（未接続）; [3] 自動要求3（未接続） *)
    RCON2_5_M : ARRAY[0..99] OF BOOL;  (* #RCON2_5 コンテナ設置; [1] 開始指令保持; [2] 予備 *)
    RCON2_5_IN_PositionDone : BOOL;  (* 位置決め完了 *)
    RCON2_5_IN_HomeDone : BOOL;  (* 原点復帰完了 *)
    RCON2_5_IN_Moving : BOOL;  (* 移動中 *)
    RCON2_5_IN_EmergencyStop : BOOL;  (* 非常停止状態（監視） *)
    RCON2_5_IN_ControllerReady : BOOL;  (* 準備完了 *)
    RCON2_5_IN_Zone2 : BOOL;  (* ゾーン2内 *)
    RCON2_5_IN_Zone1 : BOOL;  (* ゾーン1内 *)
    RCON2_5_IN_CommandDone : BOOL;  (* 指令完了 *)
    RCON2_5_IN_OverloadWarning : BOOL;  (* 過負荷警告 *)
    RCON2_5_IN_PushMiss : BOOL;  (* 押付け空振り（未使用） *)
    RCON2_5_IN_ServoReady : BOOL;  (* サーボON状態 *)
    RCON2_5_IN_Alarm : BOOL;  (* 軸異常 *)
    RCON2_5_Ready : BOOL;  (* 動作準備（安全許可とは別） *)
    RCON2_5_MoveDone : BOOL;  (* 動作完了 *)
    RCON2_5_OUT_TargetPos_mm : LREAL;  (* 目標位置 [mm] *)
    RCON2_5_OUT_PositionBand_mm : LREAL;  (* 位置決め幅 [mm] *)
    RCON2_5_OUT_Speed_mm_s : LREAL;  (* 指令速度 [mm/s] *)
    RCON2_5_OUT_AccDec_G : LREAL;  (* 加減速度 [G] *)
    RCON2_5_OUT_PushLimit_pct : LREAL;  (* 押付け制限 [%]（未使用） *)
    RCON2_5_ActualPos_mm : LREAL;  (* 現在位置 [mm] *)
    RCON2_5_Current_mA : DINT;  (* 指令電流 [mA]（監視値） *)
    RCON2_5_ActualSpeed_mm_s : LREAL;  (* 現在速度 [mm/s] *)
    RCON2_5_AlarmCode : UINT;  (* 軸異常コード *)
    RCON2_5_DataValid : BOOL;  (* 入力有効（安全許可とは別） *)
    RCON2_5_Auto : ARRAY[0..99] OF Bool;  (* 自動移動要求; [1] 自動要求1（未接続）; [2] 自動要求2（未接続）; [3] 自動要求3（未接続） *)
END_VAR
VAR
    _e1 : R_TRIG;
    _e2 : R_TRIG;
    _e3 : R_TRIG;
    _p4 : BOOL;
    _e5 : R_TRIG;
    _e6 : R_TRIG;
    _e7 : R_TRIG;
    _p8 : BOOL;
    _e9 : R_TRIG;
    _e10 : R_TRIG;
    _e11 : R_TRIG;
    _p12 : BOOL;
    _e13 : R_TRIG;
    _e14 : R_TRIG;
    _e15 : R_TRIG;
    _p16 : BOOL;
    _e17 : R_TRIG;
    _e18 : R_TRIG;
    _e19 : R_TRIG;
    _p20 : BOOL;
    _e21 : R_TRIG;
    _e22 : R_TRIG;
    _e23 : R_TRIG;
    _p24 : BOOL;
    _e25 : R_TRIG;
    _e26 : R_TRIG;
    _e27 : R_TRIG;
    _p28 : BOOL;
    _e29 : R_TRIG;
    _e30 : R_TRIG;
    _e31 : R_TRIG;
    _p32 : BOOL;
    _e33 : R_TRIG;
    _e34 : R_TRIG;
    _e35 : R_TRIG;
    _p36 : BOOL;
    _e37 : R_TRIG;
    _e38 : R_TRIG;
    _e39 : R_TRIG;
    _p40 : BOOL;
    _e41 : R_TRIG;
    _e42 : R_TRIG;
    _e43 : R_TRIG;
    _p44 : BOOL;
    _e45 : R_TRIG;
    _p46 : BOOL;
    _e47 : R_TRIG;
    _p48 : BOOL;
    _e49 : R_TRIG;
    _p50 : BOOL;
    _e51 : R_TRIG;
    _e52 : R_TRIG;
    _p53 : BOOL;
    _e54 : R_TRIG;
    _e55 : R_TRIG;
    _p56 : BOOL;
    _p57 : BOOL;
    _e58 : R_TRIG;
    _p59 : BOOL;
    _e60 : R_TRIG;
    _p61 : BOOL;
    _e62 : R_TRIG;
    _p63 : BOOL;
    _e64 : R_TRIG;
    _e65 : R_TRIG;
    _p66 : BOOL;
    _e67 : R_TRIG;
    _e68 : R_TRIG;
    _p69 : BOOL;
    _p70 : BOOL;
    _p71 : BOOL;
    _p72 : BOOL;
END_VAR

(* Section RCON_IAI: ladder, written here as Structured Text *)

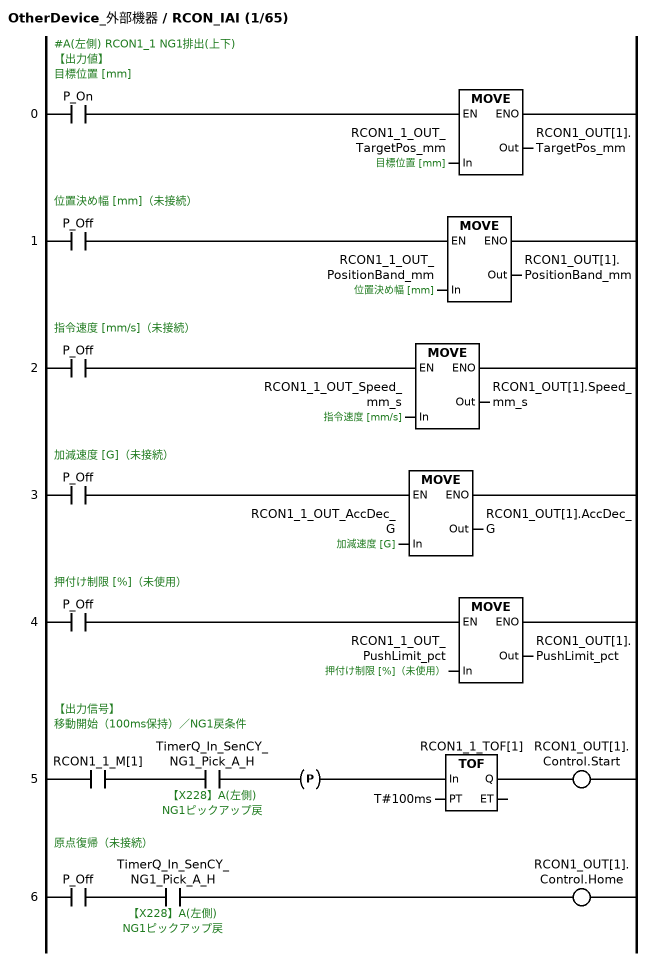
(* Rung 0: #A(左側) RCON1_1 NG1排出(上下) / 【出力値】 / 目標位置 [mm] *)
IF P_On THEN RCON1_OUT[1].TargetPos_mm := RCON1_1_OUT_TargetPos_mm; END_IF;
(* Rung 1: 位置決め幅 [mm]（未接続） *)
IF P_Off THEN RCON1_OUT[1].PositionBand_mm := RCON1_1_OUT_PositionBand_mm; END_IF;
(* Rung 2: 指令速度 [mm/s]（未接続） *)
IF P_Off THEN RCON1_OUT[1].Speed_mm_s := RCON1_1_OUT_Speed_mm_s; END_IF;
(* Rung 3: 加減速度 [G]（未接続） *)
IF P_Off THEN RCON1_OUT[1].AccDec_G := RCON1_1_OUT_AccDec_G; END_IF;
(* Rung 4: 押付け制限 [%]（未使用） *)
IF P_Off THEN RCON1_OUT[1].PushLimit_pct := RCON1_1_OUT_PushLimit_pct; END_IF;
(* Rung 5: 【出力信号】 / 移動開始（100ms保持）／NG1戻条件 *)
_e1(CLK := RCON1_1_M[1] AND TimerQ_In_SenCY_NG1_Pick_A_H);
RCON1_1_TOF[1](In := _e1.Q, PT := T#100ms);
RCON1_OUT[1].Control.Start := RCON1_1_TOF[1].Q;
(* Rung 6: 原点復帰（未接続） *)
RCON1_OUT[1].Control.Home := P_Off AND TimerQ_In_SenCY_NG1_Pick_A_H;

